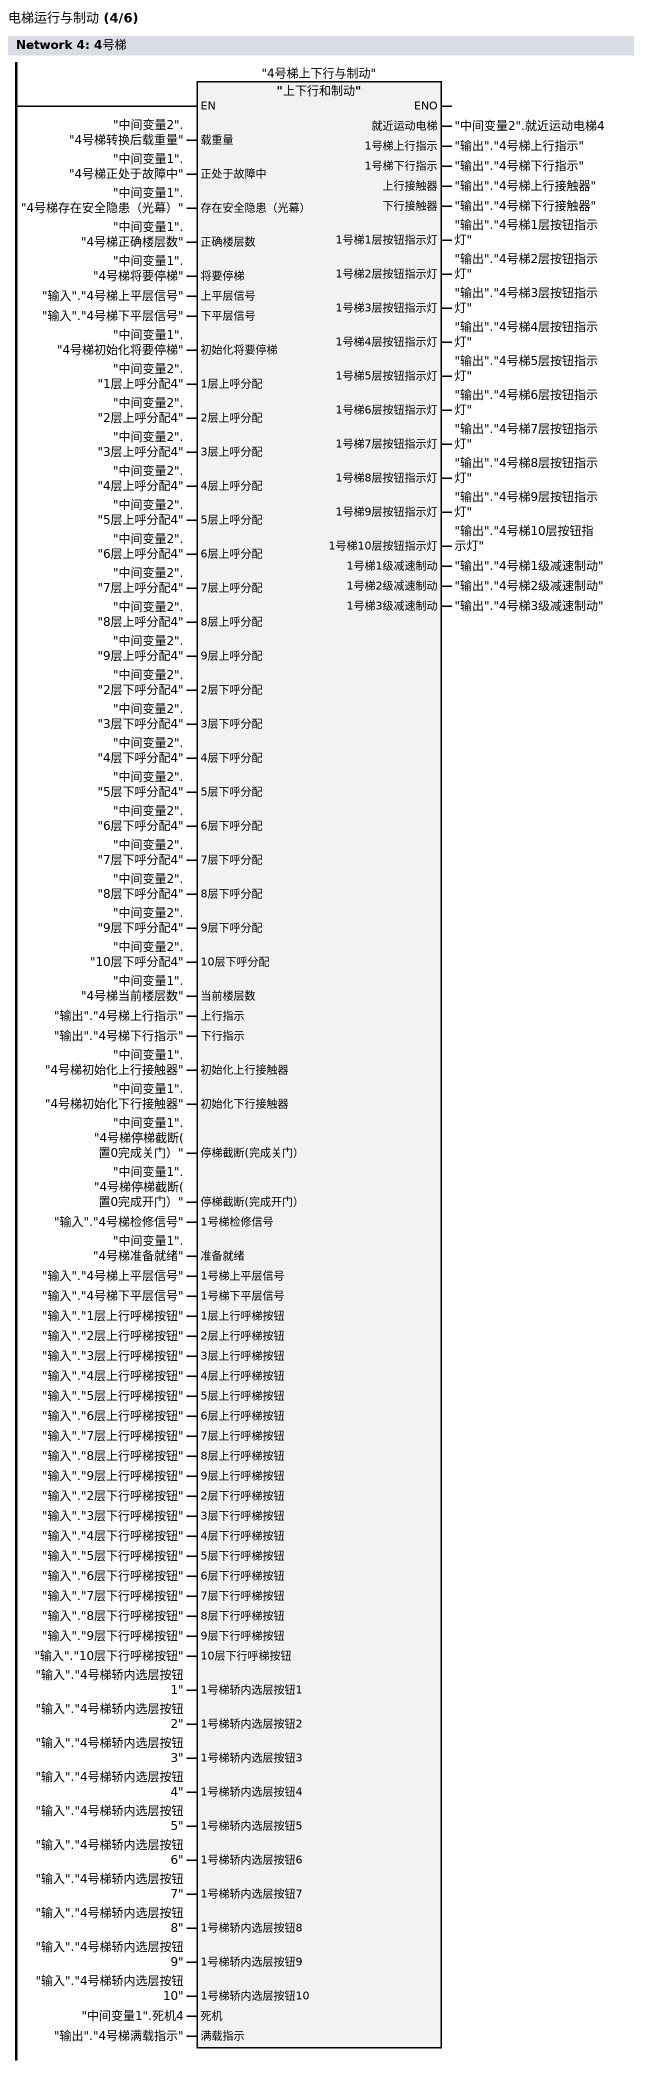
   RUNG wire#powerrail
      "4号梯上下行与制动"(载重量 := "中间变量2"."4号梯转换后载重量", 正处于故障中 := "中间变量1"."4号梯正处于故障中", "存在安全隐患（光幕）" := "中间变量1"."4号梯存在安全隐患（光幕）", 正确楼层数 := "中间变量1"."4号梯正确楼层数", 将要停梯 := "中间变量1"."4号梯将要停梯", 上平层信号 := "输入"."4号梯上平层信号", 下平层信号 := "输入"."4号梯下平层信号", 初始化将要停梯 := "中间变量1"."4号梯初始化将要停梯", "1层上呼分配" := "中间变量2"."1层上呼分配4", "2层上呼分配" := "中间变量2"."2层上呼分配4", "3层上呼分配" := "中间变量2"."3层上呼分配4", "4层上呼分配" := "中间变量2"."4层上呼分配4", "5层上呼分配" := "中间变量2"."5层上呼分配4", "6层上呼分配" := "中间变量2"."6层上呼分配4", "7层上呼分配" := "中间变量2"."7层上呼分配4", "8层上呼分配" := "中间变量2"."8层上呼分配4", "9层上呼分配" := "中间变量2"."9层上呼分配4", "2层下呼分配" := "中间变量2"."2层下呼分配4", "3层下呼分配" := "中间变量2"."3层下呼分配4", "4层下呼分配" := "中间变量2"."4层下呼分配4", "5层下呼分配" := "中间变量2"."5层下呼分配4", "6层下呼分配" := "中间变量2"."6层下呼分配4", "7层下呼分配" := "中间变量2"."7层下呼分配4", "8层下呼分配" := "中间变量2"."8层下呼分配4", "9层下呼分配" := "中间变量2"."9层下呼分配4", "10层下呼分配" := "中间变量2"."10层下呼分配4", 当前楼层数 := "中间变量1"."4号梯当前楼层数", 上行指示 := "输出"."4号梯上行指示", 下行指示 := "输出"."4号梯下行指示", 初始化上行接触器 := "中间变量1"."4号梯初始化上行接触器", 初始化下行接触器 := "中间变量1"."4号梯初始化下行接触器", "停梯截断(完成关门）" := "中间变量1"."4号梯停梯截断(置0完成关门）", "停梯截断(完成开门）" := "中间变量1"."4号梯停梯截断(置0完成开门）", "1号梯检修信号" := "输入"."4号梯检修信号", 准备就绪 := "中间变量1"."4号梯准备就绪", "1号梯上平层信号" := "输入"."4号梯上平层信号", "1号梯下平层信号" := "输入"."4号梯下平层信号", "1层上行呼梯按钮" := "输入"."1层上行呼梯按钮", "2层上行呼梯按钮" := "输入"."2层上行呼梯按钮", "3层上行呼梯按钮" := "输入"."3层上行呼梯按钮", "4层上行呼梯按钮" := "输入"."4层上行呼梯按钮", "5层上行呼梯按钮" := "输入"."5层上行呼梯按钮", "6层上行呼梯按钮" := "输入"."6层上行呼梯按钮", "7层上行呼梯按钮" := "输入"."7层上行呼梯按钮", "8层上行呼梯按钮" := "输入"."8层上行呼梯按钮", "9层上行呼梯按钮" := "输入"."9层上行呼梯按钮", "2层下行呼梯按钮" := "输入"."2层下行呼梯按钮", "3层下行呼梯按钮" := "输入"."3层下行呼梯按钮", "4层下行呼梯按钮" := "输入"."4层下行呼梯按钮", "5层下行呼梯按钮" := "输入"."5层下行呼梯按钮", "6层下行呼梯按钮" := "输入"."6层下行呼梯按钮", "7层下行呼梯按钮" := "输入"."7层下行呼梯按钮", "8层下行呼梯按钮" := "输入"."8层下行呼梯按钮", "9层下行呼梯按钮" := "输入"."9层下行呼梯按钮", "10层下行呼梯按钮" := "输入"."10层下行呼梯按钮", "1号梯轿内选层按钮1" := "输入"."4号梯轿内选层按钮1", "1号梯轿内选层按钮2" := "输入"."4号梯轿内选层按钮2", "1号梯轿内选层按钮3" := "输入"."4号梯轿内选层按钮3", "1号梯轿内选层按钮4" := "输入"."4号梯轿内选层按钮4", "1号梯轿内选层按钮5" := "输入"."4号梯轿内选层按钮5", "1号梯轿内选层按钮6" := "输入"."4号梯轿内选层按钮6", "1号梯轿内选层按钮7" := "输入"."4号梯轿内选层按钮7", "1号梯轿内选层按钮8" := "输入"."4号梯轿内选层按钮8", "1号梯轿内选层按钮9" := "输入"."4号梯轿内选层按钮9", "1号梯轿内选层按钮10" := "输入"."4号梯轿内选层按钮10", 死机 := "中间变量1".死机4, 满载指示 := "输出"."4号梯满载指示", 就近运动电梯 => "中间变量2".就近运动电梯4, "1号梯上行指示" => "输出"."4号梯上行指示", "1号梯下行指示" => "输出"."4号梯下行指示", 上行接触器 => "输出"."4号梯上行接触器", 下行接触器 => "输出"."4号梯下行接触器", "1号梯1层按钮指示灯" => "输出"."4号梯1层按钮指示灯", "1号梯2层按钮指示灯" => "输出"."4号梯2层按钮指示灯", "1号梯3层按钮指示灯" => "输出"."4号梯3层按钮指示灯", "1号梯4层按钮指示灯" => "输出"."4号梯4层按钮指示灯", "1号梯5层按钮指示灯" => "输出"."4号梯5层按钮指示灯", "1号梯6层按钮指示灯" => "输出"."4号梯6层按钮指示灯", "1号梯7层按钮指示灯" => "输出"."4号梯7层按钮指示灯", "1号梯8层按钮指示灯" => "输出"."4号梯8层按钮指示灯", "1号梯9层按钮指示灯" => "输出"."4号梯9层按钮指示灯", "1号梯10层按钮指示灯" => "输出"."4号梯10层按钮指示灯", "1号梯1级减速制动" => "输出"."4号梯1级减速制动", "1号梯2级减速制动" => "输出"."4号梯2级减速制动", "1号梯3级减速制动" => "输出"."4号梯3级减速制动")
   END_RUNG
   // the same network as SCL:
   "4号梯上下行与制动"(载重量 := "中间变量2"."4号梯转换后载重量",   // "上下行和制动"
               正处于故障中 := "中间变量1"."4号梯正处于故障中",
               "存在安全隐患（光幕）" := "中间变量1"."4号梯存在安全隐患（光幕）",
               正确楼层数 := "中间变量1"."4号梯正确楼层数",
               将要停梯 := "中间变量1"."4号梯将要停梯",
               上平层信号 := "输入"."4号梯上平层信号",
               下平层信号 := "输入"."4号梯下平层信号",
               初始化将要停梯 := "中间变量1"."4号梯初始化将要停梯",
               "1层上呼分配" := "中间变量2"."1层上呼分配4",
               "2层上呼分配" := "中间变量2"."2层上呼分配4",
               "3层上呼分配" := "中间变量2"."3层上呼分配4",
               "4层上呼分配" := "中间变量2"."4层上呼分配4",
               "5层上呼分配" := "中间变量2"."5层上呼分配4",
               "6层上呼分配" := "中间变量2"."6层上呼分配4",
               "7层上呼分配" := "中间变量2"."7层上呼分配4",
               "8层上呼分配" := "中间变量2"."8层上呼分配4",
               "9层上呼分配" := "中间变量2"."9层上呼分配4",
               "2层下呼分配" := "中间变量2"."2层下呼分配4",
               "3层下呼分配" := "中间变量2"."3层下呼分配4",
               "4层下呼分配" := "中间变量2"."4层下呼分配4",
               "5层下呼分配" := "中间变量2"."5层下呼分配4",
               "6层下呼分配" := "中间变量2"."6层下呼分配4",
               "7层下呼分配" := "中间变量2"."7层下呼分配4",
               "8层下呼分配" := "中间变量2"."8层下呼分配4",
               "9层下呼分配" := "中间变量2"."9层下呼分配4",
               "10层下呼分配" := "中间变量2"."10层下呼分配4",
               当前楼层数 := "中间变量1"."4号梯当前楼层数",
               上行指示 := "输出"."4号梯上行指示",
               下行指示 := "输出"."4号梯下行指示",
               初始化上行接触器 := "中间变量1"."4号梯初始化上行接触器",
               初始化下行接触器 := "中间变量1"."4号梯初始化下行接触器",
               "停梯截断(完成关门）" := "中间变量1"."4号梯停梯截断(置0完成关门）",
               "停梯截断(完成开门）" := "中间变量1"."4号梯停梯截断(置0完成开门）",
               "1号梯检修信号" := "输入"."4号梯检修信号",
               准备就绪 := "中间变量1"."4号梯准备就绪",
               "1号梯上平层信号" := "输入"."4号梯上平层信号",
               "1号梯下平层信号" := "输入"."4号梯下平层信号",
               "1层上行呼梯按钮" := "输入"."1层上行呼梯按钮",
               "2层上行呼梯按钮" := "输入"."2层上行呼梯按钮",
               "3层上行呼梯按钮" := "输入"."3层上行呼梯按钮",
               "4层上行呼梯按钮" := "输入"."4层上行呼梯按钮",
               "5层上行呼梯按钮" := "输入"."5层上行呼梯按钮",
               "6层上行呼梯按钮" := "输入"."6层上行呼梯按钮",
               "7层上行呼梯按钮" := "输入"."7层上行呼梯按钮",
               "8层上行呼梯按钮" := "输入"."8层上行呼梯按钮",
               "9层上行呼梯按钮" := "输入"."9层上行呼梯按钮",
               "2层下行呼梯按钮" := "输入"."2层下行呼梯按钮",
               "3层下行呼梯按钮" := "输入"."3层下行呼梯按钮",
               "4层下行呼梯按钮" := "输入"."4层下行呼梯按钮",
               "5层下行呼梯按钮" := "输入"."5层下行呼梯按钮",
               "6层下行呼梯按钮" := "输入"."6层下行呼梯按钮",
               "7层下行呼梯按钮" := "输入"."7层下行呼梯按钮",
               "8层下行呼梯按钮" := "输入"."8层下行呼梯按钮",
               "9层下行呼梯按钮" := "输入"."9层下行呼梯按钮",
               "10层下行呼梯按钮" := "输入"."10层下行呼梯按钮",
               "1号梯轿内选层按钮1" := "输入"."4号梯轿内选层按钮1",
               "1号梯轿内选层按钮2" := "输入"."4号梯轿内选层按钮2",
               "1号梯轿内选层按钮3" := "输入"."4号梯轿内选层按钮3",
               "1号梯轿内选层按钮4" := "输入"."4号梯轿内选层按钮4",
               "1号梯轿内选层按钮5" := "输入"."4号梯轿内选层按钮5",
               "1号梯轿内选层按钮6" := "输入"."4号梯轿内选层按钮6",
               "1号梯轿内选层按钮7" := "输入"."4号梯轿内选层按钮7",
               "1号梯轿内选层按钮8" := "输入"."4号梯轿内选层按钮8",
               "1号梯轿内选层按钮9" := "输入"."4号梯轿内选层按钮9",
               "1号梯轿内选层按钮10" := "输入"."4号梯轿内选层按钮10",
               死机 := "中间变量1".死机4,
               满载指示 := "输出"."4号梯满载指示",
               就近运动电梯 => "中间变量2".就近运动电梯4,
               "1号梯上行指示" => "输出"."4号梯上行指示",
               "1号梯下行指示" => "输出"."4号梯下行指示",
               上行接触器 => "输出"."4号梯上行接触器",
               下行接触器 => "输出"."4号梯下行接触器",
               "1号梯1层按钮指示灯" => "输出"."4号梯1层按钮指示灯",
               "1号梯2层按钮指示灯" => "输出"."4号梯2层按钮指示灯",
               "1号梯3层按钮指示灯" => "输出"."4号梯3层按钮指示灯",
               "1号梯4层按钮指示灯" => "输出"."4号梯4层按钮指示灯",
               "1号梯5层按钮指示灯" => "输出"."4号梯5层按钮指示灯",
               "1号梯6层按钮指示灯" => "输出"."4号梯6层按钮指示灯",
               "1号梯7层按钮指示灯" => "输出"."4号梯7层按钮指示灯",
               "1号梯8层按钮指示灯" => "输出"."4号梯8层按钮指示灯",
               "1号梯9层按钮指示灯" => "输出"."4号梯9层按钮指示灯",
               "1号梯10层按钮指示灯" => "输出"."4号梯10层按钮指示灯",
               "1号梯1级减速制动" => "输出"."4号梯1级减速制动",
               "1号梯2级减速制动" => "输出"."4号梯2级减速制动",
               "1号梯3级减速制动" => "输出"."4号梯3级减速制动");
END_REGION

REGION Network 5: 5号梯
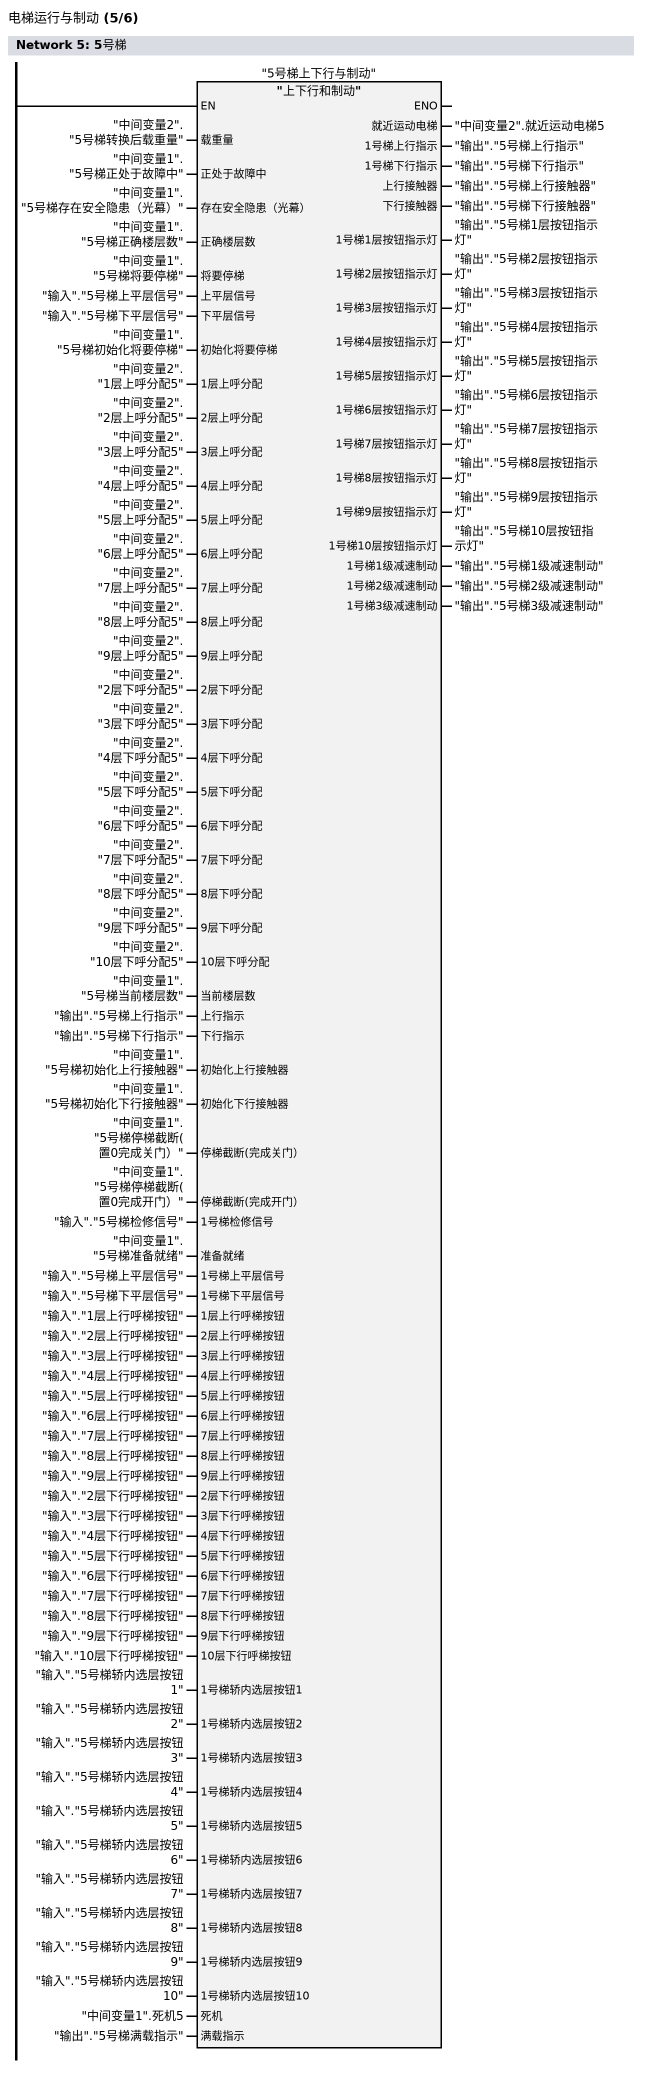
   RUNG wire#powerrail
      "5号梯上下行与制动"(载重量 := "中间变量2"."5号梯转换后载重量", 正处于故障中 := "中间变量1"."5号梯正处于故障中", "存在安全隐患（光幕）" := "中间变量1"."5号梯存在安全隐患（光幕）", 正确楼层数 := "中间变量1"."5号梯正确楼层数", 将要停梯 := "中间变量1"."5号梯将要停梯", 上平层信号 := "输入"."5号梯上平层信号", 下平层信号 := "输入"."5号梯下平层信号", 初始化将要停梯 := "中间变量1"."5号梯初始化将要停梯", "1层上呼分配" := "中间变量2"."1层上呼分配5", "2层上呼分配" := "中间变量2"."2层上呼分配5", "3层上呼分配" := "中间变量2"."3层上呼分配5", "4层上呼分配" := "中间变量2"."4层上呼分配5", "5层上呼分配" := "中间变量2"."5层上呼分配5", "6层上呼分配" := "中间变量2"."6层上呼分配5", "7层上呼分配" := "中间变量2"."7层上呼分配5", "8层上呼分配" := "中间变量2"."8层上呼分配5", "9层上呼分配" := "中间变量2"."9层上呼分配5", "2层下呼分配" := "中间变量2"."2层下呼分配5", "3层下呼分配" := "中间变量2"."3层下呼分配5", "4层下呼分配" := "中间变量2"."4层下呼分配5", "5层下呼分配" := "中间变量2"."5层下呼分配5", "6层下呼分配" := "中间变量2"."6层下呼分配5", "7层下呼分配" := "中间变量2"."7层下呼分配5", "8层下呼分配" := "中间变量2"."8层下呼分配5", "9层下呼分配" := "中间变量2"."9层下呼分配5", "10层下呼分配" := "中间变量2"."10层下呼分配5", 当前楼层数 := "中间变量1"."5号梯当前楼层数", 上行指示 := "输出"."5号梯上行指示", 下行指示 := "输出"."5号梯下行指示", 初始化上行接触器 := "中间变量1"."5号梯初始化上行接触器", 初始化下行接触器 := "中间变量1"."5号梯初始化下行接触器", "停梯截断(完成关门）" := "中间变量1"."5号梯停梯截断(置0完成关门）", "停梯截断(完成开门）" := "中间变量1"."5号梯停梯截断(置0完成开门）", "1号梯检修信号" := "输入"."5号梯检修信号", 准备就绪 := "中间变量1"."5号梯准备就绪", "1号梯上平层信号" := "输入"."5号梯上平层信号", "1号梯下平层信号" := "输入"."5号梯下平层信号", "1层上行呼梯按钮" := "输入"."1层上行呼梯按钮", "2层上行呼梯按钮" := "输入"."2层上行呼梯按钮", "3层上行呼梯按钮" := "输入"."3层上行呼梯按钮", "4层上行呼梯按钮" := "输入"."4层上行呼梯按钮", "5层上行呼梯按钮" := "输入"."5层上行呼梯按钮", "6层上行呼梯按钮" := "输入"."6层上行呼梯按钮", "7层上行呼梯按钮" := "输入"."7层上行呼梯按钮", "8层上行呼梯按钮" := "输入"."8层上行呼梯按钮", "9层上行呼梯按钮" := "输入"."9层上行呼梯按钮", "2层下行呼梯按钮" := "输入"."2层下行呼梯按钮", "3层下行呼梯按钮" := "输入"."3层下行呼梯按钮", "4层下行呼梯按钮" := "输入"."4层下行呼梯按钮", "5层下行呼梯按钮" := "输入"."5层下行呼梯按钮", "6层下行呼梯按钮" := "输入"."6层下行呼梯按钮", "7层下行呼梯按钮" := "输入"."7层下行呼梯按钮", "8层下行呼梯按钮" := "输入"."8层下行呼梯按钮", "9层下行呼梯按钮" := "输入"."9层下行呼梯按钮", "10层下行呼梯按钮" := "输入"."10层下行呼梯按钮", "1号梯轿内选层按钮1" := "输入"."5号梯轿内选层按钮1", "1号梯轿内选层按钮2" := "输入"."5号梯轿内选层按钮2", "1号梯轿内选层按钮3" := "输入"."5号梯轿内选层按钮3", "1号梯轿内选层按钮4" := "输入"."5号梯轿内选层按钮4", "1号梯轿内选层按钮5" := "输入"."5号梯轿内选层按钮5", "1号梯轿内选层按钮6" := "输入"."5号梯轿内选层按钮6", "1号梯轿内选层按钮7" := "输入"."5号梯轿内选层按钮7", "1号梯轿内选层按钮8" := "输入"."5号梯轿内选层按钮8", "1号梯轿内选层按钮9" := "输入"."5号梯轿内选层按钮9", "1号梯轿内选层按钮10" := "输入"."5号梯轿内选层按钮10", 死机 := "中间变量1".死机5, 满载指示 := "输出"."5号梯满载指示", 就近运动电梯 => "中间变量2".就近运动电梯5, "1号梯上行指示" => "输出"."5号梯上行指示", "1号梯下行指示" => "输出"."5号梯下行指示", 上行接触器 => "输出"."5号梯上行接触器", 下行接触器 => "输出"."5号梯下行接触器", "1号梯1层按钮指示灯" => "输出"."5号梯1层按钮指示灯", "1号梯2层按钮指示灯" => "输出"."5号梯2层按钮指示灯", "1号梯3层按钮指示灯" => "输出"."5号梯3层按钮指示灯", "1号梯4层按钮指示灯" => "输出"."5号梯4层按钮指示灯", "1号梯5层按钮指示灯" => "输出"."5号梯5层按钮指示灯", "1号梯6层按钮指示灯" => "输出"."5号梯6层按钮指示灯", "1号梯7层按钮指示灯" => "输出"."5号梯7层按钮指示灯", "1号梯8层按钮指示灯" => "输出"."5号梯8层按钮指示灯", "1号梯9层按钮指示灯" => "输出"."5号梯9层按钮指示灯", "1号梯10层按钮指示灯" => "输出"."5号梯10层按钮指示灯", "1号梯1级减速制动" => "输出"."5号梯1级减速制动", "1号梯2级减速制动" => "输出"."5号梯2级减速制动", "1号梯3级减速制动" => "输出"."5号梯3级减速制动")
   END_RUNG
   // the same network as SCL:
   "5号梯上下行与制动"(载重量 := "中间变量2"."5号梯转换后载重量",   // "上下行和制动"
               正处于故障中 := "中间变量1"."5号梯正处于故障中",
               "存在安全隐患（光幕）" := "中间变量1"."5号梯存在安全隐患（光幕）",
               正确楼层数 := "中间变量1"."5号梯正确楼层数",
               将要停梯 := "中间变量1"."5号梯将要停梯",
               上平层信号 := "输入"."5号梯上平层信号",
               下平层信号 := "输入"."5号梯下平层信号",
               初始化将要停梯 := "中间变量1"."5号梯初始化将要停梯",
               "1层上呼分配" := "中间变量2"."1层上呼分配5",
               "2层上呼分配" := "中间变量2"."2层上呼分配5",
               "3层上呼分配" := "中间变量2"."3层上呼分配5",
               "4层上呼分配" := "中间变量2"."4层上呼分配5",
               "5层上呼分配" := "中间变量2"."5层上呼分配5",
               "6层上呼分配" := "中间变量2"."6层上呼分配5",
               "7层上呼分配" := "中间变量2"."7层上呼分配5",
               "8层上呼分配" := "中间变量2"."8层上呼分配5",
               "9层上呼分配" := "中间变量2"."9层上呼分配5",
               "2层下呼分配" := "中间变量2"."2层下呼分配5",
               "3层下呼分配" := "中间变量2"."3层下呼分配5",
               "4层下呼分配" := "中间变量2"."4层下呼分配5",
               "5层下呼分配" := "中间变量2"."5层下呼分配5",
               "6层下呼分配" := "中间变量2"."6层下呼分配5",
               "7层下呼分配" := "中间变量2"."7层下呼分配5",
               "8层下呼分配" := "中间变量2"."8层下呼分配5",
               "9层下呼分配" := "中间变量2"."9层下呼分配5",
               "10层下呼分配" := "中间变量2"."10层下呼分配5",
               当前楼层数 := "中间变量1"."5号梯当前楼层数",
               上行指示 := "输出"."5号梯上行指示",
               下行指示 := "输出"."5号梯下行指示",
               初始化上行接触器 := "中间变量1"."5号梯初始化上行接触器",
               初始化下行接触器 := "中间变量1"."5号梯初始化下行接触器",
               "停梯截断(完成关门）" := "中间变量1"."5号梯停梯截断(置0完成关门）",
               "停梯截断(完成开门）" := "中间变量1"."5号梯停梯截断(置0完成开门）",
               "1号梯检修信号" := "输入"."5号梯检修信号",
               准备就绪 := "中间变量1"."5号梯准备就绪",
               "1号梯上平层信号" := "输入"."5号梯上平层信号",
               "1号梯下平层信号" := "输入"."5号梯下平层信号",
               "1层上行呼梯按钮" := "输入"."1层上行呼梯按钮",
               "2层上行呼梯按钮" := "输入"."2层上行呼梯按钮",
               "3层上行呼梯按钮" := "输入"."3层上行呼梯按钮",
               "4层上行呼梯按钮" := "输入"."4层上行呼梯按钮",
               "5层上行呼梯按钮" := "输入"."5层上行呼梯按钮",
               "6层上行呼梯按钮" := "输入"."6层上行呼梯按钮",
               "7层上行呼梯按钮" := "输入"."7层上行呼梯按钮",
               "8层上行呼梯按钮" := "输入"."8层上行呼梯按钮",
               "9层上行呼梯按钮" := "输入"."9层上行呼梯按钮",
               "2层下行呼梯按钮" := "输入"."2层下行呼梯按钮",
               "3层下行呼梯按钮" := "输入"."3层下行呼梯按钮",
               "4层下行呼梯按钮" := "输入"."4层下行呼梯按钮",
               "5层下行呼梯按钮" := "输入"."5层下行呼梯按钮",
               "6层下行呼梯按钮" := "输入"."6层下行呼梯按钮",
               "7层下行呼梯按钮" := "输入"."7层下行呼梯按钮",
               "8层下行呼梯按钮" := "输入"."8层下行呼梯按钮",
               "9层下行呼梯按钮" := "输入"."9层下行呼梯按钮",
               "10层下行呼梯按钮" := "输入"."10层下行呼梯按钮",
               "1号梯轿内选层按钮1" := "输入"."5号梯轿内选层按钮1",
               "1号梯轿内选层按钮2" := "输入"."5号梯轿内选层按钮2",
               "1号梯轿内选层按钮3" := "输入"."5号梯轿内选层按钮3",
               "1号梯轿内选层按钮4" := "输入"."5号梯轿内选层按钮4",
               "1号梯轿内选层按钮5" := "输入"."5号梯轿内选层按钮5",
               "1号梯轿内选层按钮6" := "输入"."5号梯轿内选层按钮6",
               "1号梯轿内选层按钮7" := "输入"."5号梯轿内选层按钮7",
               "1号梯轿内选层按钮8" := "输入"."5号梯轿内选层按钮8",
               "1号梯轿内选层按钮9" := "输入"."5号梯轿内选层按钮9",
               "1号梯轿内选层按钮10" := "输入"."5号梯轿内选层按钮10",
               死机 := "中间变量1".死机5,
               满载指示 := "输出"."5号梯满载指示",
               就近运动电梯 => "中间变量2".就近运动电梯5,
               "1号梯上行指示" => "输出"."5号梯上行指示",
               "1号梯下行指示" => "输出"."5号梯下行指示",
               上行接触器 => "输出"."5号梯上行接触器",
               下行接触器 => "输出"."5号梯下行接触器",
               "1号梯1层按钮指示灯" => "输出"."5号梯1层按钮指示灯",
               "1号梯2层按钮指示灯" => "输出"."5号梯2层按钮指示灯",
               "1号梯3层按钮指示灯" => "输出"."5号梯3层按钮指示灯",
               "1号梯4层按钮指示灯" => "输出"."5号梯4层按钮指示灯",
               "1号梯5层按钮指示灯" => "输出"."5号梯5层按钮指示灯",
               "1号梯6层按钮指示灯" => "输出"."5号梯6层按钮指示灯",
               "1号梯7层按钮指示灯" => "输出"."5号梯7层按钮指示灯",
               "1号梯8层按钮指示灯" => "输出"."5号梯8层按钮指示灯",
               "1号梯9层按钮指示灯" => "输出"."5号梯9层按钮指示灯",
               "1号梯10层按钮指示灯" => "输出"."5号梯10层按钮指示灯",
               "1号梯1级减速制动" => "输出"."5号梯1级减速制动",
               "1号梯2级减速制动" => "输出"."5号梯2级减速制动",
               "1号梯3级减速制动" => "输出"."5号梯3级减速制动");
END_REGION

REGION Network 6: 6号梯
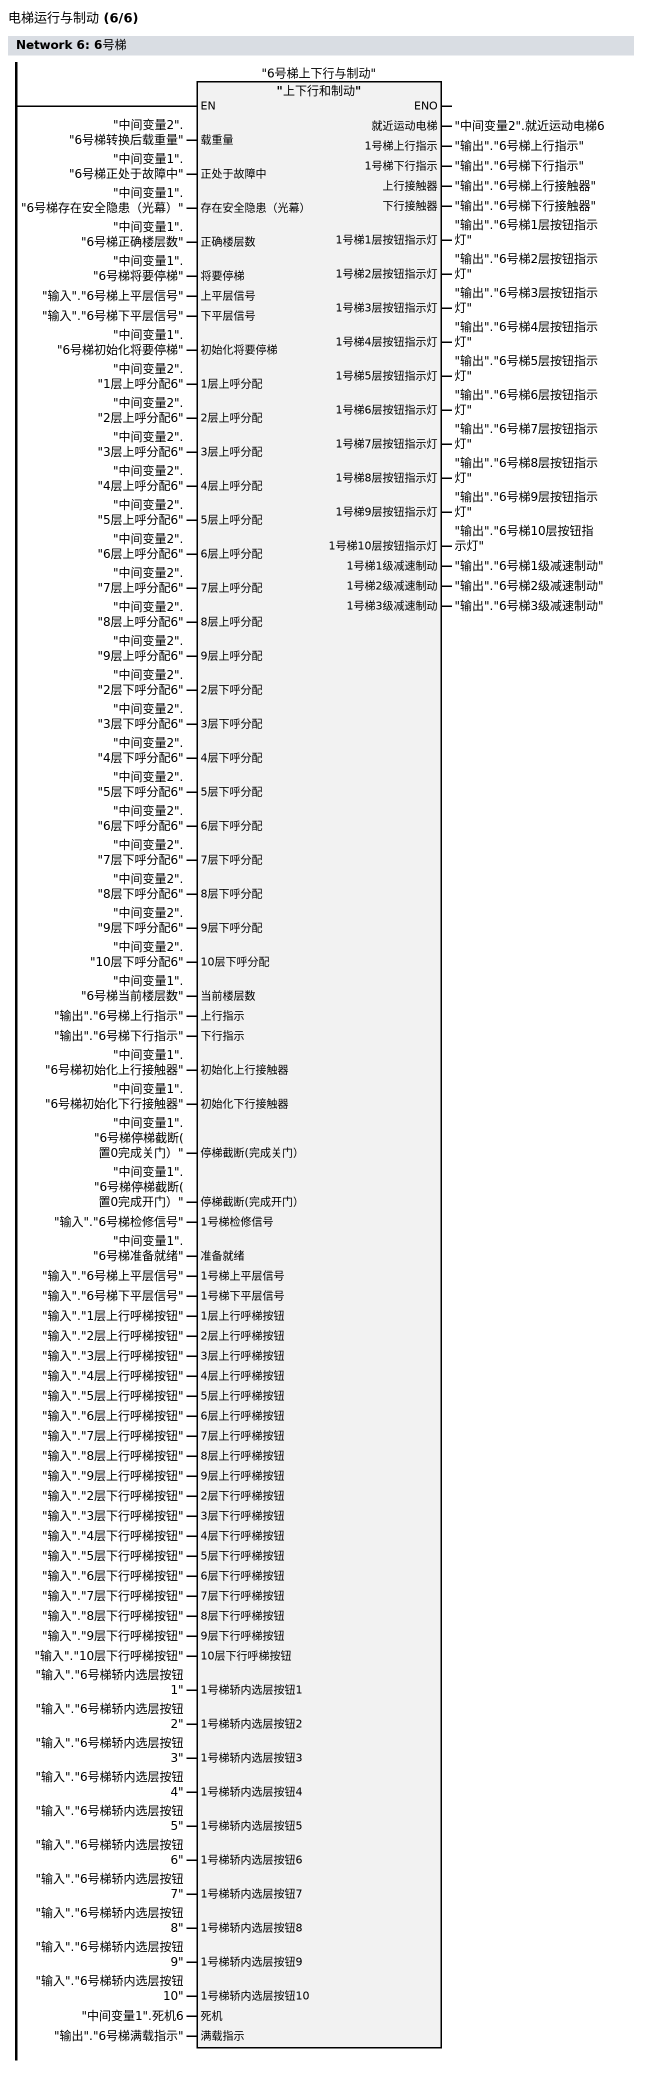
   RUNG wire#powerrail
      "6号梯上下行与制动"(载重量 := "中间变量2"."6号梯转换后载重量", 正处于故障中 := "中间变量1"."6号梯正处于故障中", "存在安全隐患（光幕）" := "中间变量1"."6号梯存在安全隐患（光幕）", 正确楼层数 := "中间变量1"."6号梯正确楼层数", 将要停梯 := "中间变量1"."6号梯将要停梯", 上平层信号 := "输入"."6号梯上平层信号", 下平层信号 := "输入"."6号梯下平层信号", 初始化将要停梯 := "中间变量1"."6号梯初始化将要停梯", "1层上呼分配" := "中间变量2"."1层上呼分配6", "2层上呼分配" := "中间变量2"."2层上呼分配6", "3层上呼分配" := "中间变量2"."3层上呼分配6", "4层上呼分配" := "中间变量2"."4层上呼分配6", "5层上呼分配" := "中间变量2"."5层上呼分配6", "6层上呼分配" := "中间变量2"."6层上呼分配6", "7层上呼分配" := "中间变量2"."7层上呼分配6", "8层上呼分配" := "中间变量2"."8层上呼分配6", "9层上呼分配" := "中间变量2"."9层上呼分配6", "2层下呼分配" := "中间变量2"."2层下呼分配6", "3层下呼分配" := "中间变量2"."3层下呼分配6", "4层下呼分配" := "中间变量2"."4层下呼分配6", "5层下呼分配" := "中间变量2"."5层下呼分配6", "6层下呼分配" := "中间变量2"."6层下呼分配6", "7层下呼分配" := "中间变量2"."7层下呼分配6", "8层下呼分配" := "中间变量2"."8层下呼分配6", "9层下呼分配" := "中间变量2"."9层下呼分配6", "10层下呼分配" := "中间变量2"."10层下呼分配6", 当前楼层数 := "中间变量1"."6号梯当前楼层数", 上行指示 := "输出"."6号梯上行指示", 下行指示 := "输出"."6号梯下行指示", 初始化上行接触器 := "中间变量1"."6号梯初始化上行接触器", 初始化下行接触器 := "中间变量1"."6号梯初始化下行接触器", "停梯截断(完成关门）" := "中间变量1"."6号梯停梯截断(置0完成关门）", "停梯截断(完成开门）" := "中间变量1"."6号梯停梯截断(置0完成开门）", "1号梯检修信号" := "输入"."6号梯检修信号", 准备就绪 := "中间变量1"."6号梯准备就绪", "1号梯上平层信号" := "输入"."6号梯上平层信号", "1号梯下平层信号" := "输入"."6号梯下平层信号", "1层上行呼梯按钮" := "输入"."1层上行呼梯按钮", "2层上行呼梯按钮" := "输入"."2层上行呼梯按钮", "3层上行呼梯按钮" := "输入"."3层上行呼梯按钮", "4层上行呼梯按钮" := "输入"."4层上行呼梯按钮", "5层上行呼梯按钮" := "输入"."5层上行呼梯按钮", "6层上行呼梯按钮" := "输入"."6层上行呼梯按钮", "7层上行呼梯按钮" := "输入"."7层上行呼梯按钮", "8层上行呼梯按钮" := "输入"."8层上行呼梯按钮", "9层上行呼梯按钮" := "输入"."9层上行呼梯按钮", "2层下行呼梯按钮" := "输入"."2层下行呼梯按钮", "3层下行呼梯按钮" := "输入"."3层下行呼梯按钮", "4层下行呼梯按钮" := "输入"."4层下行呼梯按钮", "5层下行呼梯按钮" := "输入"."5层下行呼梯按钮", "6层下行呼梯按钮" := "输入"."6层下行呼梯按钮", "7层下行呼梯按钮" := "输入"."7层下行呼梯按钮", "8层下行呼梯按钮" := "输入"."8层下行呼梯按钮", "9层下行呼梯按钮" := "输入"."9层下行呼梯按钮", "10层下行呼梯按钮" := "输入"."10层下行呼梯按钮", "1号梯轿内选层按钮1" := "输入"."6号梯轿内选层按钮1", "1号梯轿内选层按钮2" := "输入"."6号梯轿内选层按钮2", "1号梯轿内选层按钮3" := "输入"."6号梯轿内选层按钮3", "1号梯轿内选层按钮4" := "输入"."6号梯轿内选层按钮4", "1号梯轿内选层按钮5" := "输入"."6号梯轿内选层按钮5", "1号梯轿内选层按钮6" := "输入"."6号梯轿内选层按钮6", "1号梯轿内选层按钮7" := "输入"."6号梯轿内选层按钮7", "1号梯轿内选层按钮8" := "输入"."6号梯轿内选层按钮8", "1号梯轿内选层按钮9" := "输入"."6号梯轿内选层按钮9", "1号梯轿内选层按钮10" := "输入"."6号梯轿内选层按钮10", 死机 := "中间变量1".死机6, 满载指示 := "输出"."6号梯满载指示", 就近运动电梯 => "中间变量2".就近运动电梯6, "1号梯上行指示" => "输出"."6号梯上行指示", "1号梯下行指示" => "输出"."6号梯下行指示", 上行接触器 => "输出"."6号梯上行接触器", 下行接触器 => "输出"."6号梯下行接触器", "1号梯1层按钮指示灯" => "输出"."6号梯1层按钮指示灯", "1号梯2层按钮指示灯" => "输出"."6号梯2层按钮指示灯", "1号梯3层按钮指示灯" => "输出"."6号梯3层按钮指示灯", "1号梯4层按钮指示灯" => "输出"."6号梯4层按钮指示灯", "1号梯5层按钮指示灯" => "输出"."6号梯5层按钮指示灯", "1号梯6层按钮指示灯" => "输出"."6号梯6层按钮指示灯", "1号梯7层按钮指示灯" => "输出"."6号梯7层按钮指示灯", "1号梯8层按钮指示灯" => "输出"."6号梯8层按钮指示灯", "1号梯9层按钮指示灯" => "输出"."6号梯9层按钮指示灯", "1号梯10层按钮指示灯" => "输出"."6号梯10层按钮指示灯", "1号梯1级减速制动" => "输出"."6号梯1级减速制动", "1号梯2级减速制动" => "输出"."6号梯2级减速制动", "1号梯3级减速制动" => "输出"."6号梯3级减速制动")
   END_RUNG
   // the same network as SCL:
   "6号梯上下行与制动"(载重量 := "中间变量2"."6号梯转换后载重量",   // "上下行和制动"
               正处于故障中 := "中间变量1"."6号梯正处于故障中",
               "存在安全隐患（光幕）" := "中间变量1"."6号梯存在安全隐患（光幕）",
               正确楼层数 := "中间变量1"."6号梯正确楼层数",
               将要停梯 := "中间变量1"."6号梯将要停梯",
               上平层信号 := "输入"."6号梯上平层信号",
               下平层信号 := "输入"."6号梯下平层信号",
               初始化将要停梯 := "中间变量1"."6号梯初始化将要停梯",
               "1层上呼分配" := "中间变量2"."1层上呼分配6",
               "2层上呼分配" := "中间变量2"."2层上呼分配6",
               "3层上呼分配" := "中间变量2"."3层上呼分配6",
               "4层上呼分配" := "中间变量2"."4层上呼分配6",
               "5层上呼分配" := "中间变量2"."5层上呼分配6",
               "6层上呼分配" := "中间变量2"."6层上呼分配6",
               "7层上呼分配" := "中间变量2"."7层上呼分配6",
               "8层上呼分配" := "中间变量2"."8层上呼分配6",
               "9层上呼分配" := "中间变量2"."9层上呼分配6",
               "2层下呼分配" := "中间变量2"."2层下呼分配6",
               "3层下呼分配" := "中间变量2"."3层下呼分配6",
               "4层下呼分配" := "中间变量2"."4层下呼分配6",
               "5层下呼分配" := "中间变量2"."5层下呼分配6",
               "6层下呼分配" := "中间变量2"."6层下呼分配6",
               "7层下呼分配" := "中间变量2"."7层下呼分配6",
               "8层下呼分配" := "中间变量2"."8层下呼分配6",
               "9层下呼分配" := "中间变量2"."9层下呼分配6",
               "10层下呼分配" := "中间变量2"."10层下呼分配6",
               当前楼层数 := "中间变量1"."6号梯当前楼层数",
               上行指示 := "输出"."6号梯上行指示",
               下行指示 := "输出"."6号梯下行指示",
               初始化上行接触器 := "中间变量1"."6号梯初始化上行接触器",
               初始化下行接触器 := "中间变量1"."6号梯初始化下行接触器",
               "停梯截断(完成关门）" := "中间变量1"."6号梯停梯截断(置0完成关门）",
               "停梯截断(完成开门）" := "中间变量1"."6号梯停梯截断(置0完成开门）",
               "1号梯检修信号" := "输入"."6号梯检修信号",
               准备就绪 := "中间变量1"."6号梯准备就绪",
               "1号梯上平层信号" := "输入"."6号梯上平层信号",
               "1号梯下平层信号" := "输入"."6号梯下平层信号",
               "1层上行呼梯按钮" := "输入"."1层上行呼梯按钮",
               "2层上行呼梯按钮" := "输入"."2层上行呼梯按钮",
               "3层上行呼梯按钮" := "输入"."3层上行呼梯按钮",
               "4层上行呼梯按钮" := "输入"."4层上行呼梯按钮",
               "5层上行呼梯按钮" := "输入"."5层上行呼梯按钮",
               "6层上行呼梯按钮" := "输入"."6层上行呼梯按钮",
               "7层上行呼梯按钮" := "输入"."7层上行呼梯按钮",
               "8层上行呼梯按钮" := "输入"."8层上行呼梯按钮",
               "9层上行呼梯按钮" := "输入"."9层上行呼梯按钮",
               "2层下行呼梯按钮" := "输入"."2层下行呼梯按钮",
               "3层下行呼梯按钮" := "输入"."3层下行呼梯按钮",
               "4层下行呼梯按钮" := "输入"."4层下行呼梯按钮",
               "5层下行呼梯按钮" := "输入"."5层下行呼梯按钮",
               "6层下行呼梯按钮" := "输入"."6层下行呼梯按钮",
               "7层下行呼梯按钮" := "输入"."7层下行呼梯按钮",
               "8层下行呼梯按钮" := "输入"."8层下行呼梯按钮",
               "9层下行呼梯按钮" := "输入"."9层下行呼梯按钮",
               "10层下行呼梯按钮" := "输入"."10层下行呼梯按钮",
               "1号梯轿内选层按钮1" := "输入"."6号梯轿内选层按钮1",
               "1号梯轿内选层按钮2" := "输入"."6号梯轿内选层按钮2",
               "1号梯轿内选层按钮3" := "输入"."6号梯轿内选层按钮3",
               "1号梯轿内选层按钮4" := "输入"."6号梯轿内选层按钮4",
               "1号梯轿内选层按钮5" := "输入"."6号梯轿内选层按钮5",
               "1号梯轿内选层按钮6" := "输入"."6号梯轿内选层按钮6",
               "1号梯轿内选层按钮7" := "输入"."6号梯轿内选层按钮7",
               "1号梯轿内选层按钮8" := "输入"."6号梯轿内选层按钮8",
               "1号梯轿内选层按钮9" := "输入"."6号梯轿内选层按钮9",
               "1号梯轿内选层按钮10" := "输入"."6号梯轿内选层按钮10",
               死机 := "中间变量1".死机6,
               满载指示 := "输出"."6号梯满载指示",
               就近运动电梯 => "中间变量2".就近运动电梯6,
               "1号梯上行指示" => "输出"."6号梯上行指示",
               "1号梯下行指示" => "输出"."6号梯下行指示",
               上行接触器 => "输出"."6号梯上行接触器",
               下行接触器 => "输出"."6号梯下行接触器",
               "1号梯1层按钮指示灯" => "输出"."6号梯1层按钮指示灯",
               "1号梯2层按钮指示灯" => "输出"."6号梯2层按钮指示灯",
               "1号梯3层按钮指示灯" => "输出"."6号梯3层按钮指示灯",
               "1号梯4层按钮指示灯" => "输出"."6号梯4层按钮指示灯",
               "1号梯5层按钮指示灯" => "输出"."6号梯5层按钮指示灯",
               "1号梯6层按钮指示灯" => "输出"."6号梯6层按钮指示灯",
               "1号梯7层按钮指示灯" => "输出"."6号梯7层按钮指示灯",
               "1号梯8层按钮指示灯" => "输出"."6号梯8层按钮指示灯",
               "1号梯9层按钮指示灯" => "输出"."6号梯9层按钮指示灯",
               "1号梯10层按钮指示灯" => "输出"."6号梯10层按钮指示灯",
               "1号梯1级减速制动" => "输出"."6号梯1级减速制动",
               "1号梯2级减速制动" => "输出"."6号梯2级减速制动",
               "1号梯3级减速制动" => "输出"."6号梯3级减速制动");
END_REGION
END_FUNCTION

FUNCTION "距离调度算法" : Void   // FC5, LAD
{ S7_Optimized_Access := 'TRUE' }
VERSION : 0.1
BEGIN

REGION Network 2: 1号梯调度距离
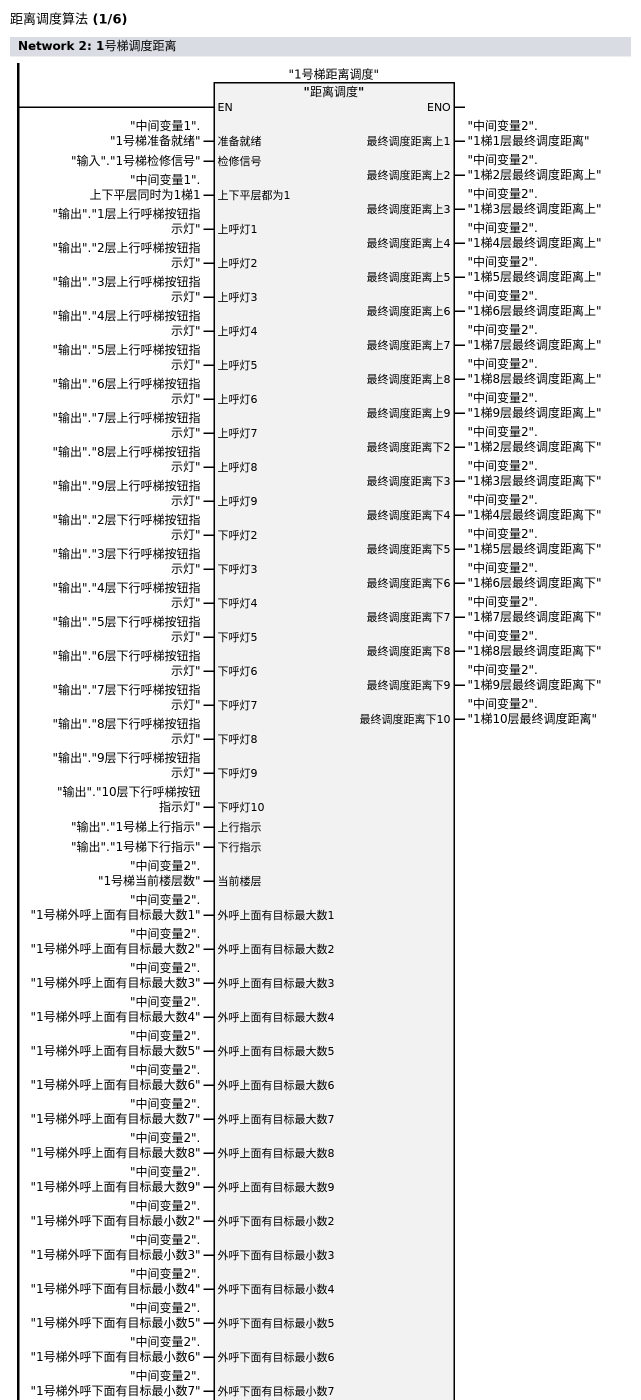
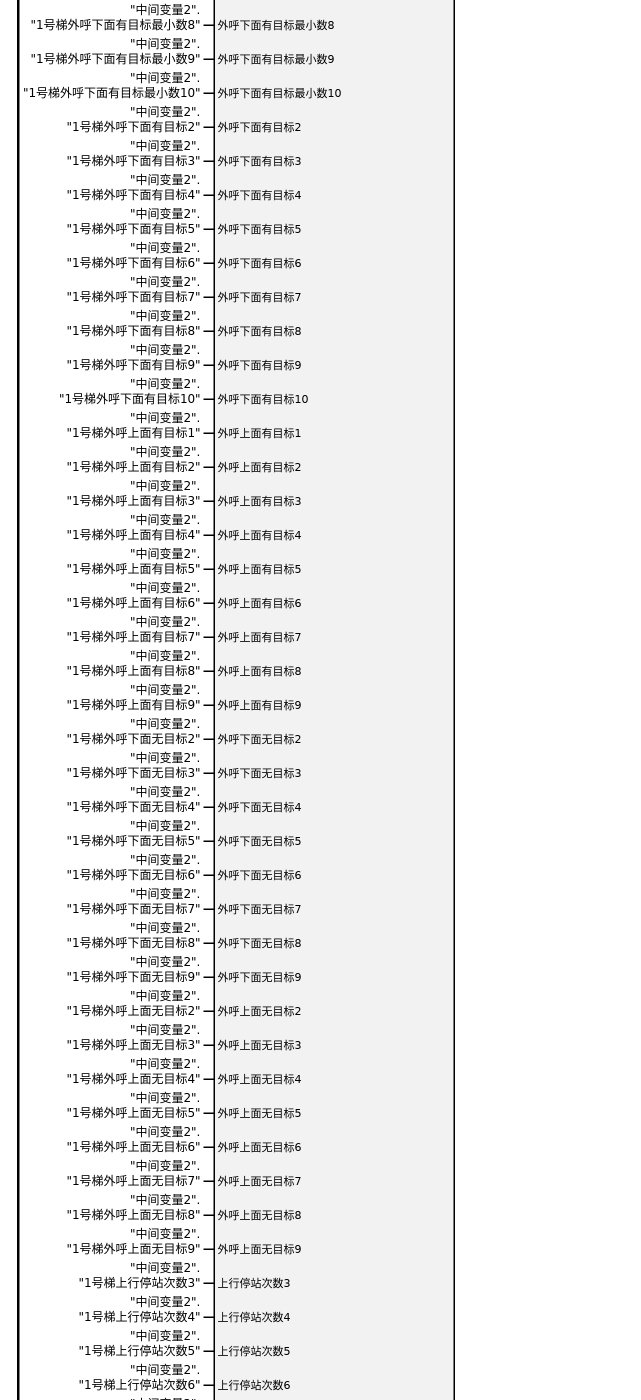
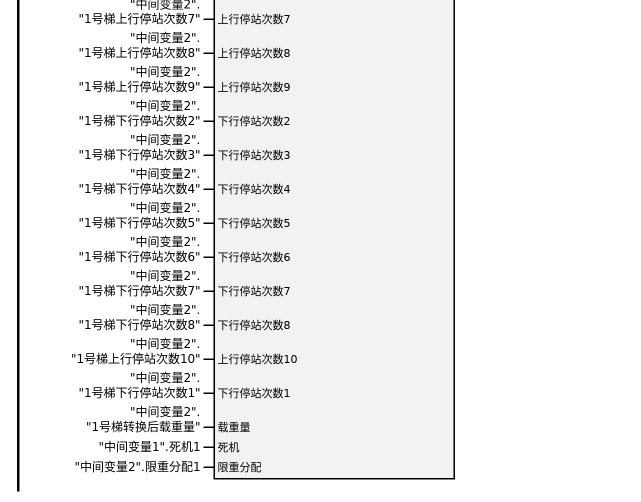
   RUNG wire#powerrail
      "1号梯距离调度"(准备就绪 := "中间变量1"."1号梯准备就绪", 检修信号 := "输入"."1号梯检修信号", 上下平层都为1 := "中间变量1".上下平层同时为1梯1, 上呼灯1 := "输出"."1层上行呼梯按钮指示灯", 上呼灯2 := "输出"."2层上行呼梯按钮指示灯", 上呼灯3 := "输出"."3层上行呼梯按钮指示灯", 上呼灯4 := "输出"."4层上行呼梯按钮指示灯", 上呼灯5 := "输出"."5层上行呼梯按钮指示灯", 上呼灯6 := "输出"."6层上行呼梯按钮指示灯", 上呼灯7 := "输出"."7层上行呼梯按钮指示灯", 上呼灯8 := "输出"."8层上行呼梯按钮指示灯", 上呼灯9 := "输出"."9层上行呼梯按钮指示灯", 下呼灯2 := "输出"."2层下行呼梯按钮指示灯", 下呼灯3 := "输出"."3层下行呼梯按钮指示灯", 下呼灯4 := "输出"."4层下行呼梯按钮指示灯", 下呼灯5 := "输出"."5层下行呼梯按钮指示灯", 下呼灯6 := "输出"."6层下行呼梯按钮指示灯", 下呼灯7 := "输出"."7层下行呼梯按钮指示灯", 下呼灯8 := "输出"."8层下行呼梯按钮指示灯", 下呼灯9 := "输出"."9层下行呼梯按钮指示灯", 下呼灯10 := "输出"."10层下行呼梯按钮指示灯", 上行指示 := "输出"."1号梯上行指示", 下行指示 := "输出"."1号梯下行指示", 当前楼层 := "中间变量2"."1号梯当前楼层数", 外呼上面有目标最大数1 := "中间变量2"."1号梯外呼上面有目标最大数1", 外呼上面有目标最大数2 := "中间变量2"."1号梯外呼上面有目标最大数2", 外呼上面有目标最大数3 := "中间变量2"."1号梯外呼上面有目标最大数3", 外呼上面有目标最大数4 := "中间变量2"."1号梯外呼上面有目标最大数4", 外呼上面有目标最大数5 := "中间变量2"."1号梯外呼上面有目标最大数5", 外呼上面有目标最大数6 := "中间变量2"."1号梯外呼上面有目标最大数6", 外呼上面有目标最大数7 := "中间变量2"."1号梯外呼上面有目标最大数7", 外呼上面有目标最大数8 := "中间变量2"."1号梯外呼上面有目标最大数8", 外呼上面有目标最大数9 := "中间变量2"."1号梯外呼上面有目标最大数9", 外呼下面有目标最小数2 := "中间变量2"."1号梯外呼下面有目标最小数2", 外呼下面有目标最小数3 := "中间变量2"."1号梯外呼下面有目标最小数3", 外呼下面有目标最小数4 := "中间变量2"."1号梯外呼下面有目标最小数4", 外呼下面有目标最小数5 := "中间变量2"."1号梯外呼下面有目标最小数5", 外呼下面有目标最小数6 := "中间变量2"."1号梯外呼下面有目标最小数6", 外呼下面有目标最小数7 := "中间变量2"."1号梯外呼下面有目标最小数7", 外呼下面有目标最小数8 := "中间变量2"."1号梯外呼下面有目标最小数8", 外呼下面有目标最小数9 := "中间变量2"."1号梯外呼下面有目标最小数9", 外呼下面有目标最小数10 := "中间变量2"."1号梯外呼下面有目标最小数10", 外呼下面有目标2 := "中间变量2"."1号梯外呼下面有目标2", 外呼下面有目标3 := "中间变量2"."1号梯外呼下面有目标3", 外呼下面有目标4 := "中间变量2"."1号梯外呼下面有目标4", 外呼下面有目标5 := "中间变量2"."1号梯外呼下面有目标5", 外呼下面有目标6 := "中间变量2"."1号梯外呼下面有目标6", 外呼下面有目标7 := "中间变量2"."1号梯外呼下面有目标7", 外呼下面有目标8 := "中间变量2"."1号梯外呼下面有目标8", 外呼下面有目标9 := "中间变量2"."1号梯外呼下面有目标9", 外呼下面有目标10 := "中间变量2"."1号梯外呼下面有目标10", 外呼上面有目标1 := "中间变量2"."1号梯外呼上面有目标1", 外呼上面有目标2 := "中间变量2"."1号梯外呼上面有目标2", 外呼上面有目标3 := "中间变量2"."1号梯外呼上面有目标3", 外呼上面有目标4 := "中间变量2"."1号梯外呼上面有目标4", 外呼上面有目标5 := "中间变量2"."1号梯外呼上面有目标5", 外呼上面有目标6 := "中间变量2"."1号梯外呼上面有目标6", 外呼上面有目标7 := "中间变量2"."1号梯外呼上面有目标7", 外呼上面有目标8 := "中间变量2"."1号梯外呼上面有目标8", 外呼上面有目标9 := "中间变量2"."1号梯外呼上面有目标9", 外呼下面无目标2 := "中间变量2"."1号梯外呼下面无目标2", 外呼下面无目标3 := "中间变量2"."1号梯外呼下面无目标3", 外呼下面无目标4 := "中间变量2"."1号梯外呼下面无目标4", 外呼下面无目标5 := "中间变量2"."1号梯外呼下面无目标5", 外呼下面无目标6 := "中间变量2"."1号梯外呼下面无目标6", 外呼下面无目标7 := "中间变量2"."1号梯外呼下面无目标7", 外呼下面无目标8 := "中间变量2"."1号梯外呼下面无目标8", 外呼下面无目标9 := "中间变量2"."1号梯外呼下面无目标9", 外呼上面无目标2 := "中间变量2"."1号梯外呼上面无目标2", 外呼上面无目标3 := "中间变量2"."1号梯外呼上面无目标3", 外呼上面无目标4 := "中间变量2"."1号梯外呼上面无目标4", 外呼上面无目标5 := "中间变量2"."1号梯外呼上面无目标5", 外呼上面无目标6 := "中间变量2"."1号梯外呼上面无目标6", 外呼上面无目标7 := "中间变量2"."1号梯外呼上面无目标7", 外呼上面无目标8 := "中间变量2"."1号梯外呼上面无目标8", 外呼上面无目标9 := "中间变量2"."1号梯外呼上面无目标9", 上行停站次数3 := "中间变量2"."1号梯上行停站次数3", 上行停站次数4 := "中间变量2"."1号梯上行停站次数4", 上行停站次数5 := "中间变量2"."1号梯上行停站次数5", 上行停站次数6 := "中间变量2"."1号梯上行停站次数6", 上行停站次数7 := "中间变量2"."1号梯上行停站次数7", 上行停站次数8 := "中间变量2"."1号梯上行停站次数8", 上行停站次数9 := "中间变量2"."1号梯上行停站次数9", 下行停站次数2 := "中间变量2"."1号梯下行停站次数2", 下行停站次数3 := "中间变量2"."1号梯下行停站次数3", 下行停站次数4 := "中间变量2"."1号梯下行停站次数4", 下行停站次数5 := "中间变量2"."1号梯下行停站次数5", 下行停站次数6 := "中间变量2"."1号梯下行停站次数6", 下行停站次数7 := "中间变量2"."1号梯下行停站次数7", 下行停站次数8 := "中间变量2"."1号梯下行停站次数8", 上行停站次数10 := "中间变量2"."1号梯上行停站次数10", 下行停站次数1 := "中间变量2"."1号梯下行停站次数1", 载重量 := "中间变量2"."1号梯转换后载重量", 死机 := "中间变量1".死机1, 限重分配 := "中间变量2".限重分配1, 最终调度距离上1 => "中间变量2"."1梯1层最终调度距离", 最终调度距离上2 => "中间变量2"."1梯2层最终调度距离上", 最终调度距离上3 => "中间变量2"."1梯3层最终调度距离上", 最终调度距离上4 => "中间变量2"."1梯4层最终调度距离上", 最终调度距离上5 => "中间变量2"."1梯5层最终调度距离上", 最终调度距离上6 => "中间变量2"."1梯6层最终调度距离上", 最终调度距离上7 => "中间变量2"."1梯7层最终调度距离上", 最终调度距离上8 => "中间变量2"."1梯8层最终调度距离上", 最终调度距离上9 => "中间变量2"."1梯9层最终调度距离上", 最终调度距离下2 => "中间变量2"."1梯2层最终调度距离下", 最终调度距离下3 => "中间变量2"."1梯3层最终调度距离下", 最终调度距离下4 => "中间变量2"."1梯4层最终调度距离下", 最终调度距离下5 => "中间变量2"."1梯5层最终调度距离下", 最终调度距离下6 => "中间变量2"."1梯6层最终调度距离下", 最终调度距离下7 => "中间变量2"."1梯7层最终调度距离下", 最终调度距离下8 => "中间变量2"."1梯8层最终调度距离下", 最终调度距离下9 => "中间变量2"."1梯9层最终调度距离下", 最终调度距离下10 => "中间变量2"."1梯10层最终调度距离")
   END_RUNG
   // the same network as SCL:
   "1号梯距离调度"(准备就绪 := "中间变量1"."1号梯准备就绪",   // "距离调度"
             检修信号 := "输入"."1号梯检修信号",
             上下平层都为1 := "中间变量1".上下平层同时为1梯1,
             上呼灯1 := "输出"."1层上行呼梯按钮指示灯",
             上呼灯2 := "输出"."2层上行呼梯按钮指示灯",
             上呼灯3 := "输出"."3层上行呼梯按钮指示灯",
             上呼灯4 := "输出"."4层上行呼梯按钮指示灯",
             上呼灯5 := "输出"."5层上行呼梯按钮指示灯",
             上呼灯6 := "输出"."6层上行呼梯按钮指示灯",
             上呼灯7 := "输出"."7层上行呼梯按钮指示灯",
             上呼灯8 := "输出"."8层上行呼梯按钮指示灯",
             上呼灯9 := "输出"."9层上行呼梯按钮指示灯",
             下呼灯2 := "输出"."2层下行呼梯按钮指示灯",
             下呼灯3 := "输出"."3层下行呼梯按钮指示灯",
             下呼灯4 := "输出"."4层下行呼梯按钮指示灯",
             下呼灯5 := "输出"."5层下行呼梯按钮指示灯",
             下呼灯6 := "输出"."6层下行呼梯按钮指示灯",
             下呼灯7 := "输出"."7层下行呼梯按钮指示灯",
             下呼灯8 := "输出"."8层下行呼梯按钮指示灯",
             下呼灯9 := "输出"."9层下行呼梯按钮指示灯",
             下呼灯10 := "输出"."10层下行呼梯按钮指示灯",
             上行指示 := "输出"."1号梯上行指示",
             下行指示 := "输出"."1号梯下行指示",
             当前楼层 := "中间变量2"."1号梯当前楼层数",
             外呼上面有目标最大数1 := "中间变量2"."1号梯外呼上面有目标最大数1",
             外呼上面有目标最大数2 := "中间变量2"."1号梯外呼上面有目标最大数2",
             外呼上面有目标最大数3 := "中间变量2"."1号梯外呼上面有目标最大数3",
             外呼上面有目标最大数4 := "中间变量2"."1号梯外呼上面有目标最大数4",
             外呼上面有目标最大数5 := "中间变量2"."1号梯外呼上面有目标最大数5",
             外呼上面有目标最大数6 := "中间变量2"."1号梯外呼上面有目标最大数6",
             外呼上面有目标最大数7 := "中间变量2"."1号梯外呼上面有目标最大数7",
             外呼上面有目标最大数8 := "中间变量2"."1号梯外呼上面有目标最大数8",
             外呼上面有目标最大数9 := "中间变量2"."1号梯外呼上面有目标最大数9",
             外呼下面有目标最小数2 := "中间变量2"."1号梯外呼下面有目标最小数2",
             外呼下面有目标最小数3 := "中间变量2"."1号梯外呼下面有目标最小数3",
             外呼下面有目标最小数4 := "中间变量2"."1号梯外呼下面有目标最小数4",
             外呼下面有目标最小数5 := "中间变量2"."1号梯外呼下面有目标最小数5",
             外呼下面有目标最小数6 := "中间变量2"."1号梯外呼下面有目标最小数6",
             外呼下面有目标最小数7 := "中间变量2"."1号梯外呼下面有目标最小数7",
             外呼下面有目标最小数8 := "中间变量2"."1号梯外呼下面有目标最小数8",
             外呼下面有目标最小数9 := "中间变量2"."1号梯外呼下面有目标最小数9",
             外呼下面有目标最小数10 := "中间变量2"."1号梯外呼下面有目标最小数10",
             外呼下面有目标2 := "中间变量2"."1号梯外呼下面有目标2",
             外呼下面有目标3 := "中间变量2"."1号梯外呼下面有目标3",
             外呼下面有目标4 := "中间变量2"."1号梯外呼下面有目标4",
             外呼下面有目标5 := "中间变量2"."1号梯外呼下面有目标5",
             外呼下面有目标6 := "中间变量2"."1号梯外呼下面有目标6",
             外呼下面有目标7 := "中间变量2"."1号梯外呼下面有目标7",
             外呼下面有目标8 := "中间变量2"."1号梯外呼下面有目标8",
             外呼下面有目标9 := "中间变量2"."1号梯外呼下面有目标9",
             外呼下面有目标10 := "中间变量2"."1号梯外呼下面有目标10",
             外呼上面有目标1 := "中间变量2"."1号梯外呼上面有目标1",
             外呼上面有目标2 := "中间变量2"."1号梯外呼上面有目标2",
             外呼上面有目标3 := "中间变量2"."1号梯外呼上面有目标3",
             外呼上面有目标4 := "中间变量2"."1号梯外呼上面有目标4",
             外呼上面有目标5 := "中间变量2"."1号梯外呼上面有目标5",
             外呼上面有目标6 := "中间变量2"."1号梯外呼上面有目标6",
             外呼上面有目标7 := "中间变量2"."1号梯外呼上面有目标7",
             外呼上面有目标8 := "中间变量2"."1号梯外呼上面有目标8",
             外呼上面有目标9 := "中间变量2"."1号梯外呼上面有目标9",
             外呼下面无目标2 := "中间变量2"."1号梯外呼下面无目标2",
             外呼下面无目标3 := "中间变量2"."1号梯外呼下面无目标3",
             外呼下面无目标4 := "中间变量2"."1号梯外呼下面无目标4",
             外呼下面无目标5 := "中间变量2"."1号梯外呼下面无目标5",
             外呼下面无目标6 := "中间变量2"."1号梯外呼下面无目标6",
             外呼下面无目标7 := "中间变量2"."1号梯外呼下面无目标7",
             外呼下面无目标8 := "中间变量2"."1号梯外呼下面无目标8",
             外呼下面无目标9 := "中间变量2"."1号梯外呼下面无目标9",
             外呼上面无目标2 := "中间变量2"."1号梯外呼上面无目标2",
             外呼上面无目标3 := "中间变量2"."1号梯外呼上面无目标3",
             外呼上面无目标4 := "中间变量2"."1号梯外呼上面无目标4",
             外呼上面无目标5 := "中间变量2"."1号梯外呼上面无目标5",
             外呼上面无目标6 := "中间变量2"."1号梯外呼上面无目标6",
             外呼上面无目标7 := "中间变量2"."1号梯外呼上面无目标7",
             外呼上面无目标8 := "中间变量2"."1号梯外呼上面无目标8",
             外呼上面无目标9 := "中间变量2"."1号梯外呼上面无目标9",
             上行停站次数3 := "中间变量2"."1号梯上行停站次数3",
             上行停站次数4 := "中间变量2"."1号梯上行停站次数4",
             上行停站次数5 := "中间变量2"."1号梯上行停站次数5",
             上行停站次数6 := "中间变量2"."1号梯上行停站次数6",
             上行停站次数7 := "中间变量2"."1号梯上行停站次数7",
             上行停站次数8 := "中间变量2"."1号梯上行停站次数8",
             上行停站次数9 := "中间变量2"."1号梯上行停站次数9",
             下行停站次数2 := "中间变量2"."1号梯下行停站次数2",
             下行停站次数3 := "中间变量2"."1号梯下行停站次数3",
             下行停站次数4 := "中间变量2"."1号梯下行停站次数4",
             下行停站次数5 := "中间变量2"."1号梯下行停站次数5",
             下行停站次数6 := "中间变量2"."1号梯下行停站次数6",
             下行停站次数7 := "中间变量2"."1号梯下行停站次数7",
             下行停站次数8 := "中间变量2"."1号梯下行停站次数8",
             上行停站次数10 := "中间变量2"."1号梯上行停站次数10",
             下行停站次数1 := "中间变量2"."1号梯下行停站次数1",
             载重量 := "中间变量2"."1号梯转换后载重量",
             死机 := "中间变量1".死机1,
             限重分配 := "中间变量2".限重分配1,
             最终调度距离上1 => "中间变量2"."1梯1层最终调度距离",
             最终调度距离上2 => "中间变量2"."1梯2层最终调度距离上",
             最终调度距离上3 => "中间变量2"."1梯3层最终调度距离上",
             最终调度距离上4 => "中间变量2"."1梯4层最终调度距离上",
             最终调度距离上5 => "中间变量2"."1梯5层最终调度距离上",
             最终调度距离上6 => "中间变量2"."1梯6层最终调度距离上",
             最终调度距离上7 => "中间变量2"."1梯7层最终调度距离上",
             最终调度距离上8 => "中间变量2"."1梯8层最终调度距离上",
             最终调度距离上9 => "中间变量2"."1梯9层最终调度距离上",
             最终调度距离下2 => "中间变量2"."1梯2层最终调度距离下",
             最终调度距离下3 => "中间变量2"."1梯3层最终调度距离下",
             最终调度距离下4 => "中间变量2"."1梯4层最终调度距离下",
             最终调度距离下5 => "中间变量2"."1梯5层最终调度距离下",
             最终调度距离下6 => "中间变量2"."1梯6层最终调度距离下",
             最终调度距离下7 => "中间变量2"."1梯7层最终调度距离下",
             最终调度距离下8 => "中间变量2"."1梯8层最终调度距离下",
             最终调度距离下9 => "中间变量2"."1梯9层最终调度距离下",
             最终调度距离下10 => "中间变量2"."1梯10层最终调度距离");
END_REGION

REGION Network 3: 2号梯调度距离
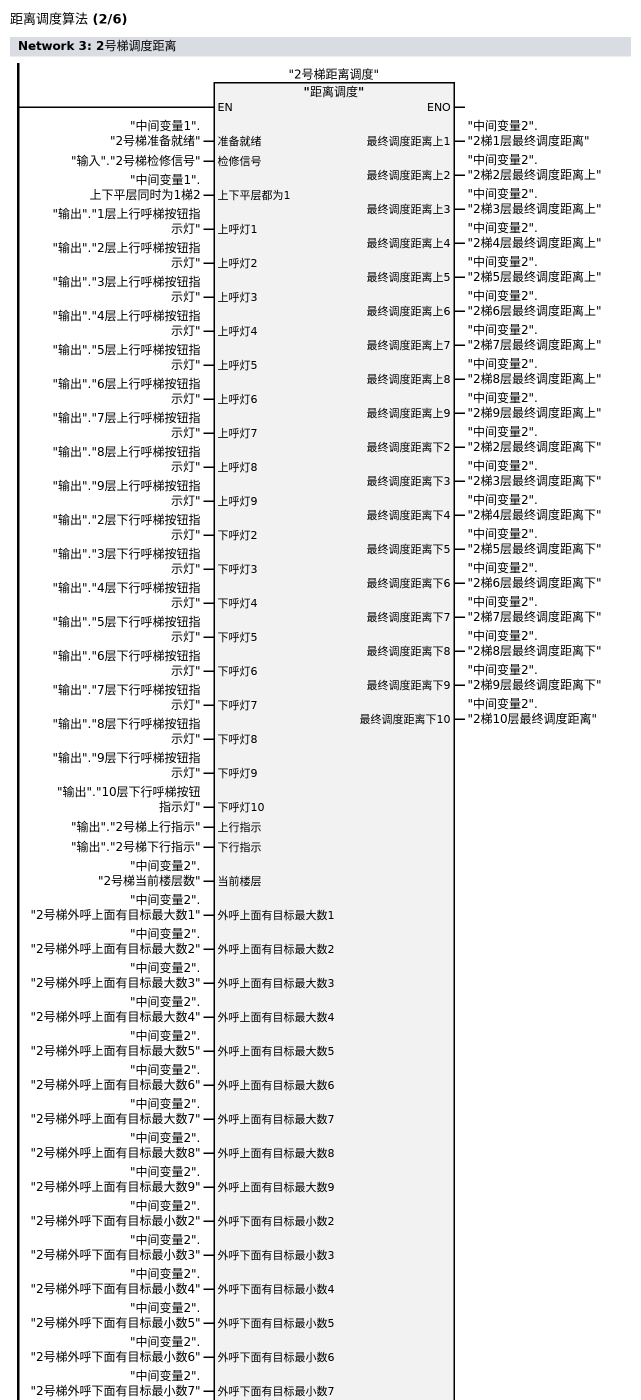
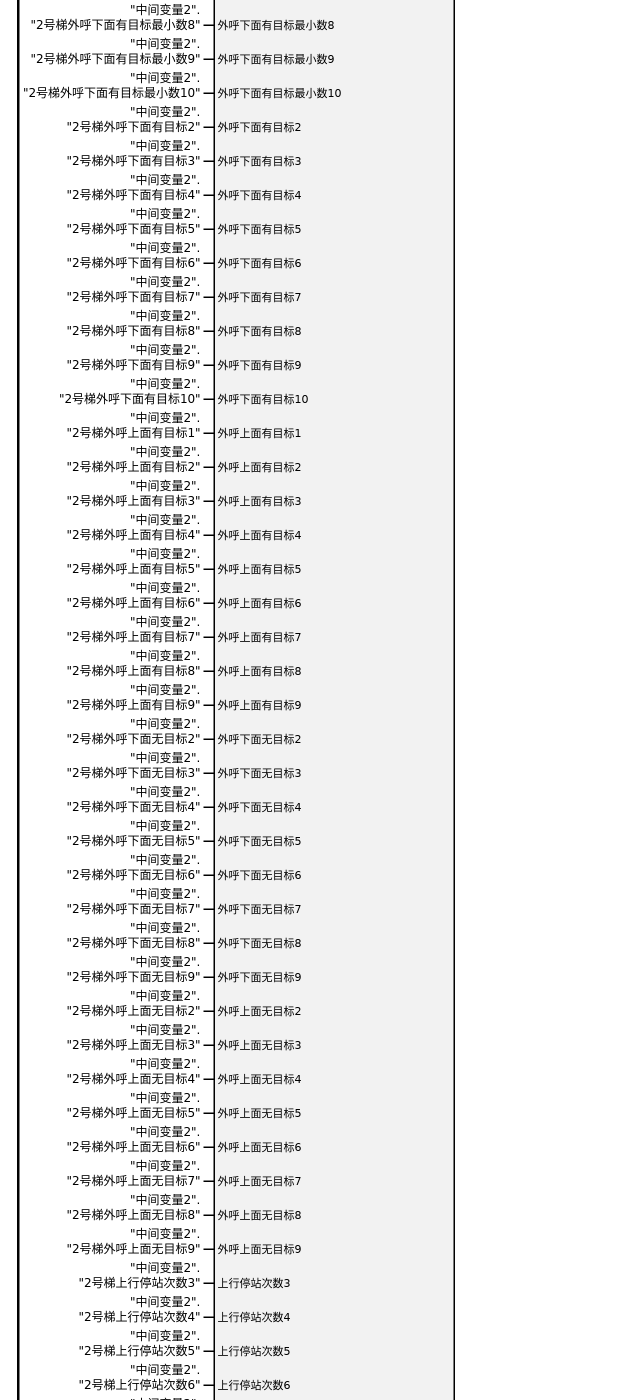
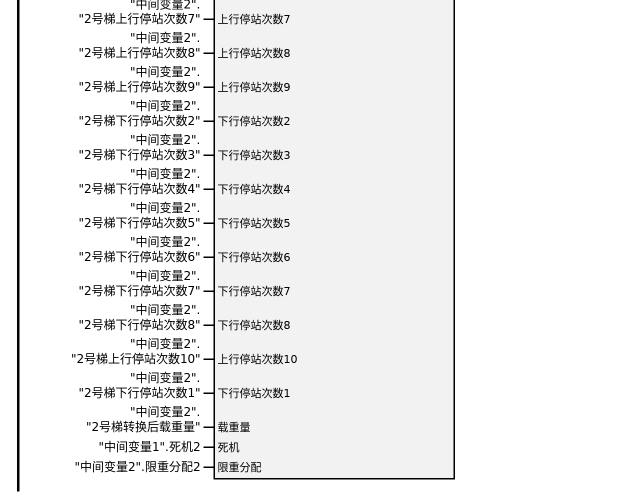
   RUNG wire#powerrail
      "2号梯距离调度"(准备就绪 := "中间变量1"."2号梯准备就绪", 检修信号 := "输入"."2号梯检修信号", 上下平层都为1 := "中间变量1".上下平层同时为1梯2, 上呼灯1 := "输出"."1层上行呼梯按钮指示灯", 上呼灯2 := "输出"."2层上行呼梯按钮指示灯", 上呼灯3 := "输出"."3层上行呼梯按钮指示灯", 上呼灯4 := "输出"."4层上行呼梯按钮指示灯", 上呼灯5 := "输出"."5层上行呼梯按钮指示灯", 上呼灯6 := "输出"."6层上行呼梯按钮指示灯", 上呼灯7 := "输出"."7层上行呼梯按钮指示灯", 上呼灯8 := "输出"."8层上行呼梯按钮指示灯", 上呼灯9 := "输出"."9层上行呼梯按钮指示灯", 下呼灯2 := "输出"."2层下行呼梯按钮指示灯", 下呼灯3 := "输出"."3层下行呼梯按钮指示灯", 下呼灯4 := "输出"."4层下行呼梯按钮指示灯", 下呼灯5 := "输出"."5层下行呼梯按钮指示灯", 下呼灯6 := "输出"."6层下行呼梯按钮指示灯", 下呼灯7 := "输出"."7层下行呼梯按钮指示灯", 下呼灯8 := "输出"."8层下行呼梯按钮指示灯", 下呼灯9 := "输出"."9层下行呼梯按钮指示灯", 下呼灯10 := "输出"."10层下行呼梯按钮指示灯", 上行指示 := "输出"."2号梯上行指示", 下行指示 := "输出"."2号梯下行指示", 当前楼层 := "中间变量2"."2号梯当前楼层数", 外呼上面有目标最大数1 := "中间变量2"."2号梯外呼上面有目标最大数1", 外呼上面有目标最大数2 := "中间变量2"."2号梯外呼上面有目标最大数2", 外呼上面有目标最大数3 := "中间变量2"."2号梯外呼上面有目标最大数3", 外呼上面有目标最大数4 := "中间变量2"."2号梯外呼上面有目标最大数4", 外呼上面有目标最大数5 := "中间变量2"."2号梯外呼上面有目标最大数5", 外呼上面有目标最大数6 := "中间变量2"."2号梯外呼上面有目标最大数6", 外呼上面有目标最大数7 := "中间变量2"."2号梯外呼上面有目标最大数7", 外呼上面有目标最大数8 := "中间变量2"."2号梯外呼上面有目标最大数8", 外呼上面有目标最大数9 := "中间变量2"."2号梯外呼上面有目标最大数9", 外呼下面有目标最小数2 := "中间变量2"."2号梯外呼下面有目标最小数2", 外呼下面有目标最小数3 := "中间变量2"."2号梯外呼下面有目标最小数3", 外呼下面有目标最小数4 := "中间变量2"."2号梯外呼下面有目标最小数4", 外呼下面有目标最小数5 := "中间变量2"."2号梯外呼下面有目标最小数5", 外呼下面有目标最小数6 := "中间变量2"."2号梯外呼下面有目标最小数6", 外呼下面有目标最小数7 := "中间变量2"."2号梯外呼下面有目标最小数7", 外呼下面有目标最小数8 := "中间变量2"."2号梯外呼下面有目标最小数8", 外呼下面有目标最小数9 := "中间变量2"."2号梯外呼下面有目标最小数9", 外呼下面有目标最小数10 := "中间变量2"."2号梯外呼下面有目标最小数10", 外呼下面有目标2 := "中间变量2"."2号梯外呼下面有目标2", 外呼下面有目标3 := "中间变量2"."2号梯外呼下面有目标3", 外呼下面有目标4 := "中间变量2"."2号梯外呼下面有目标4", 外呼下面有目标5 := "中间变量2"."2号梯外呼下面有目标5", 外呼下面有目标6 := "中间变量2"."2号梯外呼下面有目标6", 外呼下面有目标7 := "中间变量2"."2号梯外呼下面有目标7", 外呼下面有目标8 := "中间变量2"."2号梯外呼下面有目标8", 外呼下面有目标9 := "中间变量2"."2号梯外呼下面有目标9", 外呼下面有目标10 := "中间变量2"."2号梯外呼下面有目标10", 外呼上面有目标1 := "中间变量2"."2号梯外呼上面有目标1", 外呼上面有目标2 := "中间变量2"."2号梯外呼上面有目标2", 外呼上面有目标3 := "中间变量2"."2号梯外呼上面有目标3", 外呼上面有目标4 := "中间变量2"."2号梯外呼上面有目标4", 外呼上面有目标5 := "中间变量2"."2号梯外呼上面有目标5", 外呼上面有目标6 := "中间变量2"."2号梯外呼上面有目标6", 外呼上面有目标7 := "中间变量2"."2号梯外呼上面有目标7", 外呼上面有目标8 := "中间变量2"."2号梯外呼上面有目标8", 外呼上面有目标9 := "中间变量2"."2号梯外呼上面有目标9", 外呼下面无目标2 := "中间变量2"."2号梯外呼下面无目标2", 外呼下面无目标3 := "中间变量2"."2号梯外呼下面无目标3", 外呼下面无目标4 := "中间变量2"."2号梯外呼下面无目标4", 外呼下面无目标5 := "中间变量2"."2号梯外呼下面无目标5", 外呼下面无目标6 := "中间变量2"."2号梯外呼下面无目标6", 外呼下面无目标7 := "中间变量2"."2号梯外呼下面无目标7", 外呼下面无目标8 := "中间变量2"."2号梯外呼下面无目标8", 外呼下面无目标9 := "中间变量2"."2号梯外呼下面无目标9", 外呼上面无目标2 := "中间变量2"."2号梯外呼上面无目标2", 外呼上面无目标3 := "中间变量2"."2号梯外呼上面无目标3", 外呼上面无目标4 := "中间变量2"."2号梯外呼上面无目标4", 外呼上面无目标5 := "中间变量2"."2号梯外呼上面无目标5", 外呼上面无目标6 := "中间变量2"."2号梯外呼上面无目标6", 外呼上面无目标7 := "中间变量2"."2号梯外呼上面无目标7", 外呼上面无目标8 := "中间变量2"."2号梯外呼上面无目标8", 外呼上面无目标9 := "中间变量2"."2号梯外呼上面无目标9", 上行停站次数3 := "中间变量2"."2号梯上行停站次数3", 上行停站次数4 := "中间变量2"."2号梯上行停站次数4", 上行停站次数5 := "中间变量2"."2号梯上行停站次数5", 上行停站次数6 := "中间变量2"."2号梯上行停站次数6", 上行停站次数7 := "中间变量2"."2号梯上行停站次数7", 上行停站次数8 := "中间变量2"."2号梯上行停站次数8", 上行停站次数9 := "中间变量2"."2号梯上行停站次数9", 下行停站次数2 := "中间变量2"."2号梯下行停站次数2", 下行停站次数3 := "中间变量2"."2号梯下行停站次数3", 下行停站次数4 := "中间变量2"."2号梯下行停站次数4", 下行停站次数5 := "中间变量2"."2号梯下行停站次数5", 下行停站次数6 := "中间变量2"."2号梯下行停站次数6", 下行停站次数7 := "中间变量2"."2号梯下行停站次数7", 下行停站次数8 := "中间变量2"."2号梯下行停站次数8", 上行停站次数10 := "中间变量2"."2号梯上行停站次数10", 下行停站次数1 := "中间变量2"."2号梯下行停站次数1", 载重量 := "中间变量2"."2号梯转换后载重量", 死机 := "中间变量1".死机2, 限重分配 := "中间变量2".限重分配2, 最终调度距离上1 => "中间变量2"."2梯1层最终调度距离", 最终调度距离上2 => "中间变量2"."2梯2层最终调度距离上", 最终调度距离上3 => "中间变量2"."2梯3层最终调度距离上", 最终调度距离上4 => "中间变量2"."2梯4层最终调度距离上", 最终调度距离上5 => "中间变量2"."2梯5层最终调度距离上", 最终调度距离上6 => "中间变量2"."2梯6层最终调度距离上", 最终调度距离上7 => "中间变量2"."2梯7层最终调度距离上", 最终调度距离上8 => "中间变量2"."2梯8层最终调度距离上", 最终调度距离上9 => "中间变量2"."2梯9层最终调度距离上", 最终调度距离下2 => "中间变量2"."2梯2层最终调度距离下", 最终调度距离下3 => "中间变量2"."2梯3层最终调度距离下", 最终调度距离下4 => "中间变量2"."2梯4层最终调度距离下", 最终调度距离下5 => "中间变量2"."2梯5层最终调度距离下", 最终调度距离下6 => "中间变量2"."2梯6层最终调度距离下", 最终调度距离下7 => "中间变量2"."2梯7层最终调度距离下", 最终调度距离下8 => "中间变量2"."2梯8层最终调度距离下", 最终调度距离下9 => "中间变量2"."2梯9层最终调度距离下", 最终调度距离下10 => "中间变量2"."2梯10层最终调度距离")
   END_RUNG
   // the same network as SCL:
   "2号梯距离调度"(准备就绪 := "中间变量1"."2号梯准备就绪",   // "距离调度"
             检修信号 := "输入"."2号梯检修信号",
             上下平层都为1 := "中间变量1".上下平层同时为1梯2,
             上呼灯1 := "输出"."1层上行呼梯按钮指示灯",
             上呼灯2 := "输出"."2层上行呼梯按钮指示灯",
             上呼灯3 := "输出"."3层上行呼梯按钮指示灯",
             上呼灯4 := "输出"."4层上行呼梯按钮指示灯",
             上呼灯5 := "输出"."5层上行呼梯按钮指示灯",
             上呼灯6 := "输出"."6层上行呼梯按钮指示灯",
             上呼灯7 := "输出"."7层上行呼梯按钮指示灯",
             上呼灯8 := "输出"."8层上行呼梯按钮指示灯",
             上呼灯9 := "输出"."9层上行呼梯按钮指示灯",
             下呼灯2 := "输出"."2层下行呼梯按钮指示灯",
             下呼灯3 := "输出"."3层下行呼梯按钮指示灯",
             下呼灯4 := "输出"."4层下行呼梯按钮指示灯",
             下呼灯5 := "输出"."5层下行呼梯按钮指示灯",
             下呼灯6 := "输出"."6层下行呼梯按钮指示灯",
             下呼灯7 := "输出"."7层下行呼梯按钮指示灯",
             下呼灯8 := "输出"."8层下行呼梯按钮指示灯",
             下呼灯9 := "输出"."9层下行呼梯按钮指示灯",
             下呼灯10 := "输出"."10层下行呼梯按钮指示灯",
             上行指示 := "输出"."2号梯上行指示",
             下行指示 := "输出"."2号梯下行指示",
             当前楼层 := "中间变量2"."2号梯当前楼层数",
             外呼上面有目标最大数1 := "中间变量2"."2号梯外呼上面有目标最大数1",
             外呼上面有目标最大数2 := "中间变量2"."2号梯外呼上面有目标最大数2",
             外呼上面有目标最大数3 := "中间变量2"."2号梯外呼上面有目标最大数3",
             外呼上面有目标最大数4 := "中间变量2"."2号梯外呼上面有目标最大数4",
             外呼上面有目标最大数5 := "中间变量2"."2号梯外呼上面有目标最大数5",
             外呼上面有目标最大数6 := "中间变量2"."2号梯外呼上面有目标最大数6",
             外呼上面有目标最大数7 := "中间变量2"."2号梯外呼上面有目标最大数7",
             外呼上面有目标最大数8 := "中间变量2"."2号梯外呼上面有目标最大数8",
             外呼上面有目标最大数9 := "中间变量2"."2号梯外呼上面有目标最大数9",
             外呼下面有目标最小数2 := "中间变量2"."2号梯外呼下面有目标最小数2",
             外呼下面有目标最小数3 := "中间变量2"."2号梯外呼下面有目标最小数3",
             外呼下面有目标最小数4 := "中间变量2"."2号梯外呼下面有目标最小数4",
             外呼下面有目标最小数5 := "中间变量2"."2号梯外呼下面有目标最小数5",
             外呼下面有目标最小数6 := "中间变量2"."2号梯外呼下面有目标最小数6",
             外呼下面有目标最小数7 := "中间变量2"."2号梯外呼下面有目标最小数7",
             外呼下面有目标最小数8 := "中间变量2"."2号梯外呼下面有目标最小数8",
             外呼下面有目标最小数9 := "中间变量2"."2号梯外呼下面有目标最小数9",
             外呼下面有目标最小数10 := "中间变量2"."2号梯外呼下面有目标最小数10",
             外呼下面有目标2 := "中间变量2"."2号梯外呼下面有目标2",
             外呼下面有目标3 := "中间变量2"."2号梯外呼下面有目标3",
             外呼下面有目标4 := "中间变量2"."2号梯外呼下面有目标4",
             外呼下面有目标5 := "中间变量2"."2号梯外呼下面有目标5",
             外呼下面有目标6 := "中间变量2"."2号梯外呼下面有目标6",
             外呼下面有目标7 := "中间变量2"."2号梯外呼下面有目标7",
             外呼下面有目标8 := "中间变量2"."2号梯外呼下面有目标8",
             外呼下面有目标9 := "中间变量2"."2号梯外呼下面有目标9",
             外呼下面有目标10 := "中间变量2"."2号梯外呼下面有目标10",
             外呼上面有目标1 := "中间变量2"."2号梯外呼上面有目标1",
             外呼上面有目标2 := "中间变量2"."2号梯外呼上面有目标2",
             外呼上面有目标3 := "中间变量2"."2号梯外呼上面有目标3",
             外呼上面有目标4 := "中间变量2"."2号梯外呼上面有目标4",
             外呼上面有目标5 := "中间变量2"."2号梯外呼上面有目标5",
             外呼上面有目标6 := "中间变量2"."2号梯外呼上面有目标6",
             外呼上面有目标7 := "中间变量2"."2号梯外呼上面有目标7",
             外呼上面有目标8 := "中间变量2"."2号梯外呼上面有目标8",
             外呼上面有目标9 := "中间变量2"."2号梯外呼上面有目标9",
             外呼下面无目标2 := "中间变量2"."2号梯外呼下面无目标2",
             外呼下面无目标3 := "中间变量2"."2号梯外呼下面无目标3",
             外呼下面无目标4 := "中间变量2"."2号梯外呼下面无目标4",
             外呼下面无目标5 := "中间变量2"."2号梯外呼下面无目标5",
             外呼下面无目标6 := "中间变量2"."2号梯外呼下面无目标6",
             外呼下面无目标7 := "中间变量2"."2号梯外呼下面无目标7",
             外呼下面无目标8 := "中间变量2"."2号梯外呼下面无目标8",
             外呼下面无目标9 := "中间变量2"."2号梯外呼下面无目标9",
             外呼上面无目标2 := "中间变量2"."2号梯外呼上面无目标2",
             外呼上面无目标3 := "中间变量2"."2号梯外呼上面无目标3",
             外呼上面无目标4 := "中间变量2"."2号梯外呼上面无目标4",
             外呼上面无目标5 := "中间变量2"."2号梯外呼上面无目标5",
             外呼上面无目标6 := "中间变量2"."2号梯外呼上面无目标6",
             外呼上面无目标7 := "中间变量2"."2号梯外呼上面无目标7",
             外呼上面无目标8 := "中间变量2"."2号梯外呼上面无目标8",
             外呼上面无目标9 := "中间变量2"."2号梯外呼上面无目标9",
             上行停站次数3 := "中间变量2"."2号梯上行停站次数3",
             上行停站次数4 := "中间变量2"."2号梯上行停站次数4",
             上行停站次数5 := "中间变量2"."2号梯上行停站次数5",
             上行停站次数6 := "中间变量2"."2号梯上行停站次数6",
             上行停站次数7 := "中间变量2"."2号梯上行停站次数7",
             上行停站次数8 := "中间变量2"."2号梯上行停站次数8",
             上行停站次数9 := "中间变量2"."2号梯上行停站次数9",
             下行停站次数2 := "中间变量2"."2号梯下行停站次数2",
             下行停站次数3 := "中间变量2"."2号梯下行停站次数3",
             下行停站次数4 := "中间变量2"."2号梯下行停站次数4",
             下行停站次数5 := "中间变量2"."2号梯下行停站次数5",
             下行停站次数6 := "中间变量2"."2号梯下行停站次数6",
             下行停站次数7 := "中间变量2"."2号梯下行停站次数7",
             下行停站次数8 := "中间变量2"."2号梯下行停站次数8",
             上行停站次数10 := "中间变量2"."2号梯上行停站次数10",
             下行停站次数1 := "中间变量2"."2号梯下行停站次数1",
             载重量 := "中间变量2"."2号梯转换后载重量",
             死机 := "中间变量1".死机2,
             限重分配 := "中间变量2".限重分配2,
             最终调度距离上1 => "中间变量2"."2梯1层最终调度距离",
             最终调度距离上2 => "中间变量2"."2梯2层最终调度距离上",
             最终调度距离上3 => "中间变量2"."2梯3层最终调度距离上",
             最终调度距离上4 => "中间变量2"."2梯4层最终调度距离上",
             最终调度距离上5 => "中间变量2"."2梯5层最终调度距离上",
             最终调度距离上6 => "中间变量2"."2梯6层最终调度距离上",
             最终调度距离上7 => "中间变量2"."2梯7层最终调度距离上",
             最终调度距离上8 => "中间变量2"."2梯8层最终调度距离上",
             最终调度距离上9 => "中间变量2"."2梯9层最终调度距离上",
             最终调度距离下2 => "中间变量2"."2梯2层最终调度距离下",
             最终调度距离下3 => "中间变量2"."2梯3层最终调度距离下",
             最终调度距离下4 => "中间变量2"."2梯4层最终调度距离下",
             最终调度距离下5 => "中间变量2"."2梯5层最终调度距离下",
             最终调度距离下6 => "中间变量2"."2梯6层最终调度距离下",
             最终调度距离下7 => "中间变量2"."2梯7层最终调度距离下",
             最终调度距离下8 => "中间变量2"."2梯8层最终调度距离下",
             最终调度距离下9 => "中间变量2"."2梯9层最终调度距离下",
             最终调度距离下10 => "中间变量2"."2梯10层最终调度距离");
END_REGION

REGION Network 4: 3号梯调度距离
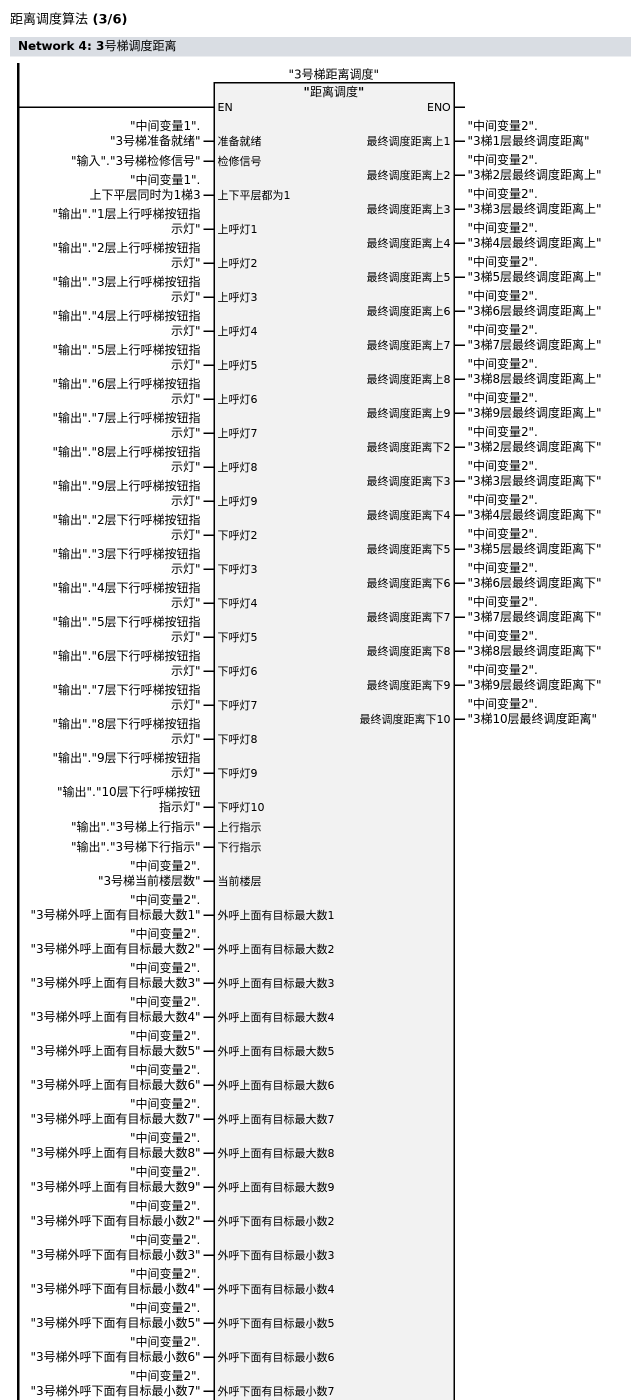
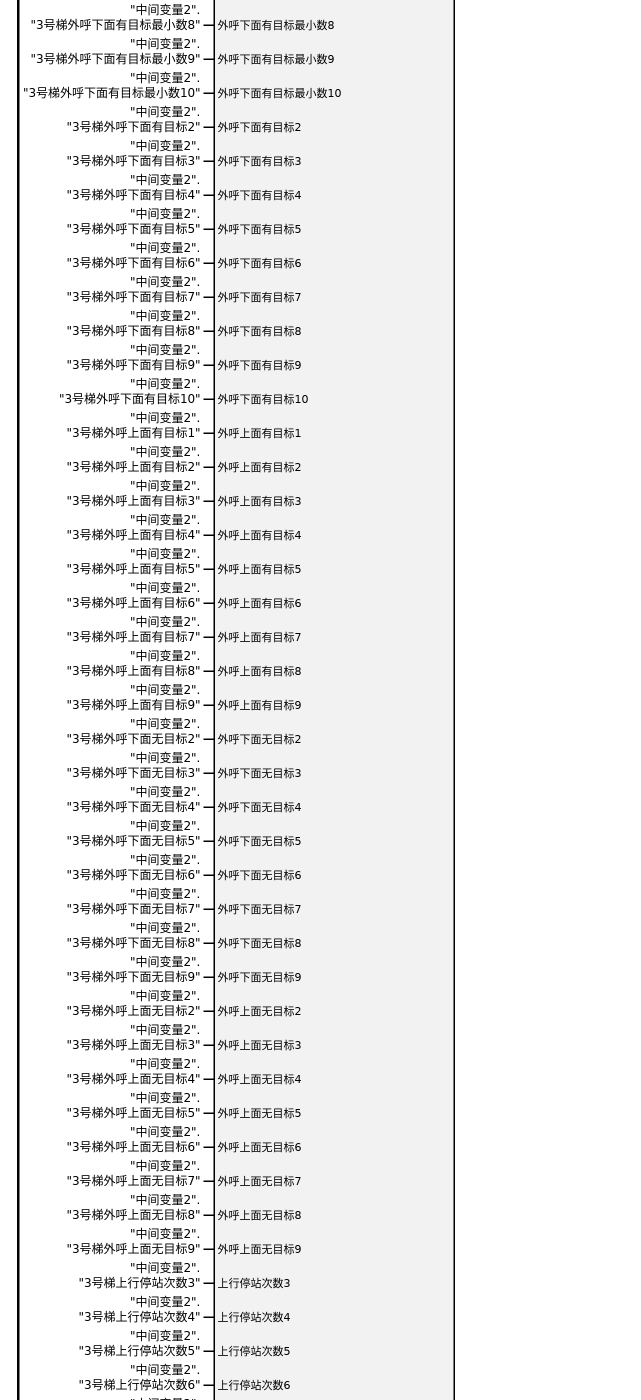
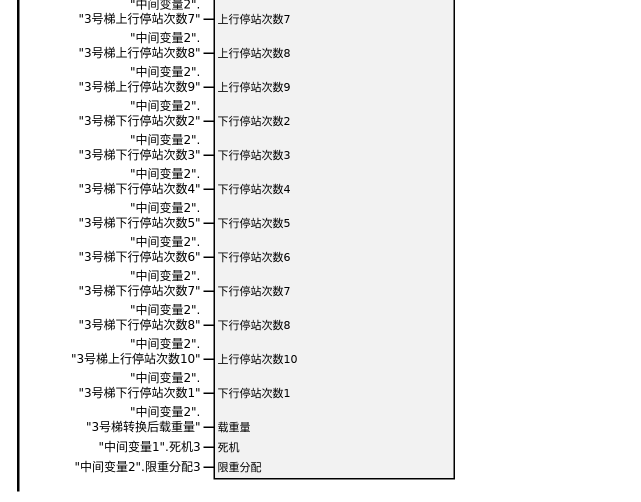
   RUNG wire#powerrail
      "3号梯距离调度"(准备就绪 := "中间变量1"."3号梯准备就绪", 检修信号 := "输入"."3号梯检修信号", 上下平层都为1 := "中间变量1".上下平层同时为1梯3, 上呼灯1 := "输出"."1层上行呼梯按钮指示灯", 上呼灯2 := "输出"."2层上行呼梯按钮指示灯", 上呼灯3 := "输出"."3层上行呼梯按钮指示灯", 上呼灯4 := "输出"."4层上行呼梯按钮指示灯", 上呼灯5 := "输出"."5层上行呼梯按钮指示灯", 上呼灯6 := "输出"."6层上行呼梯按钮指示灯", 上呼灯7 := "输出"."7层上行呼梯按钮指示灯", 上呼灯8 := "输出"."8层上行呼梯按钮指示灯", 上呼灯9 := "输出"."9层上行呼梯按钮指示灯", 下呼灯2 := "输出"."2层下行呼梯按钮指示灯", 下呼灯3 := "输出"."3层下行呼梯按钮指示灯", 下呼灯4 := "输出"."4层下行呼梯按钮指示灯", 下呼灯5 := "输出"."5层下行呼梯按钮指示灯", 下呼灯6 := "输出"."6层下行呼梯按钮指示灯", 下呼灯7 := "输出"."7层下行呼梯按钮指示灯", 下呼灯8 := "输出"."8层下行呼梯按钮指示灯", 下呼灯9 := "输出"."9层下行呼梯按钮指示灯", 下呼灯10 := "输出"."10层下行呼梯按钮指示灯", 上行指示 := "输出"."3号梯上行指示", 下行指示 := "输出"."3号梯下行指示", 当前楼层 := "中间变量2"."3号梯当前楼层数", 外呼上面有目标最大数1 := "中间变量2"."3号梯外呼上面有目标最大数1", 外呼上面有目标最大数2 := "中间变量2"."3号梯外呼上面有目标最大数2", 外呼上面有目标最大数3 := "中间变量2"."3号梯外呼上面有目标最大数3", 外呼上面有目标最大数4 := "中间变量2"."3号梯外呼上面有目标最大数4", 外呼上面有目标最大数5 := "中间变量2"."3号梯外呼上面有目标最大数5", 外呼上面有目标最大数6 := "中间变量2"."3号梯外呼上面有目标最大数6", 外呼上面有目标最大数7 := "中间变量2"."3号梯外呼上面有目标最大数7", 外呼上面有目标最大数8 := "中间变量2"."3号梯外呼上面有目标最大数8", 外呼上面有目标最大数9 := "中间变量2"."3号梯外呼上面有目标最大数9", 外呼下面有目标最小数2 := "中间变量2"."3号梯外呼下面有目标最小数2", 外呼下面有目标最小数3 := "中间变量2"."3号梯外呼下面有目标最小数3", 外呼下面有目标最小数4 := "中间变量2"."3号梯外呼下面有目标最小数4", 外呼下面有目标最小数5 := "中间变量2"."3号梯外呼下面有目标最小数5", 外呼下面有目标最小数6 := "中间变量2"."3号梯外呼下面有目标最小数6", 外呼下面有目标最小数7 := "中间变量2"."3号梯外呼下面有目标最小数7", 外呼下面有目标最小数8 := "中间变量2"."3号梯外呼下面有目标最小数8", 外呼下面有目标最小数9 := "中间变量2"."3号梯外呼下面有目标最小数9", 外呼下面有目标最小数10 := "中间变量2"."3号梯外呼下面有目标最小数10", 外呼下面有目标2 := "中间变量2"."3号梯外呼下面有目标2", 外呼下面有目标3 := "中间变量2"."3号梯外呼下面有目标3", 外呼下面有目标4 := "中间变量2"."3号梯外呼下面有目标4", 外呼下面有目标5 := "中间变量2"."3号梯外呼下面有目标5", 外呼下面有目标6 := "中间变量2"."3号梯外呼下面有目标6", 外呼下面有目标7 := "中间变量2"."3号梯外呼下面有目标7", 外呼下面有目标8 := "中间变量2"."3号梯外呼下面有目标8", 外呼下面有目标9 := "中间变量2"."3号梯外呼下面有目标9", 外呼下面有目标10 := "中间变量2"."3号梯外呼下面有目标10", 外呼上面有目标1 := "中间变量2"."3号梯外呼上面有目标1", 外呼上面有目标2 := "中间变量2"."3号梯外呼上面有目标2", 外呼上面有目标3 := "中间变量2"."3号梯外呼上面有目标3", 外呼上面有目标4 := "中间变量2"."3号梯外呼上面有目标4", 外呼上面有目标5 := "中间变量2"."3号梯外呼上面有目标5", 外呼上面有目标6 := "中间变量2"."3号梯外呼上面有目标6", 外呼上面有目标7 := "中间变量2"."3号梯外呼上面有目标7", 外呼上面有目标8 := "中间变量2"."3号梯外呼上面有目标8", 外呼上面有目标9 := "中间变量2"."3号梯外呼上面有目标9", 外呼下面无目标2 := "中间变量2"."3号梯外呼下面无目标2", 外呼下面无目标3 := "中间变量2"."3号梯外呼下面无目标3", 外呼下面无目标4 := "中间变量2"."3号梯外呼下面无目标4", 外呼下面无目标5 := "中间变量2"."3号梯外呼下面无目标5", 外呼下面无目标6 := "中间变量2"."3号梯外呼下面无目标6", 外呼下面无目标7 := "中间变量2"."3号梯外呼下面无目标7", 外呼下面无目标8 := "中间变量2"."3号梯外呼下面无目标8", 外呼下面无目标9 := "中间变量2"."3号梯外呼下面无目标9", 外呼上面无目标2 := "中间变量2"."3号梯外呼上面无目标2", 外呼上面无目标3 := "中间变量2"."3号梯外呼上面无目标3", 外呼上面无目标4 := "中间变量2"."3号梯外呼上面无目标4", 外呼上面无目标5 := "中间变量2"."3号梯外呼上面无目标5", 外呼上面无目标6 := "中间变量2"."3号梯外呼上面无目标6", 外呼上面无目标7 := "中间变量2"."3号梯外呼上面无目标7", 外呼上面无目标8 := "中间变量2"."3号梯外呼上面无目标8", 外呼上面无目标9 := "中间变量2"."3号梯外呼上面无目标9", 上行停站次数3 := "中间变量2"."3号梯上行停站次数3", 上行停站次数4 := "中间变量2"."3号梯上行停站次数4", 上行停站次数5 := "中间变量2"."3号梯上行停站次数5", 上行停站次数6 := "中间变量2"."3号梯上行停站次数6", 上行停站次数7 := "中间变量2"."3号梯上行停站次数7", 上行停站次数8 := "中间变量2"."3号梯上行停站次数8", 上行停站次数9 := "中间变量2"."3号梯上行停站次数9", 下行停站次数2 := "中间变量2"."3号梯下行停站次数2", 下行停站次数3 := "中间变量2"."3号梯下行停站次数3", 下行停站次数4 := "中间变量2"."3号梯下行停站次数4", 下行停站次数5 := "中间变量2"."3号梯下行停站次数5", 下行停站次数6 := "中间变量2"."3号梯下行停站次数6", 下行停站次数7 := "中间变量2"."3号梯下行停站次数7", 下行停站次数8 := "中间变量2"."3号梯下行停站次数8", 上行停站次数10 := "中间变量2"."3号梯上行停站次数10", 下行停站次数1 := "中间变量2"."3号梯下行停站次数1", 载重量 := "中间变量2"."3号梯转换后载重量", 死机 := "中间变量1".死机3, 限重分配 := "中间变量2".限重分配3, 最终调度距离上1 => "中间变量2"."3梯1层最终调度距离", 最终调度距离上2 => "中间变量2"."3梯2层最终调度距离上", 最终调度距离上3 => "中间变量2"."3梯3层最终调度距离上", 最终调度距离上4 => "中间变量2"."3梯4层最终调度距离上", 最终调度距离上5 => "中间变量2"."3梯5层最终调度距离上", 最终调度距离上6 => "中间变量2"."3梯6层最终调度距离上", 最终调度距离上7 => "中间变量2"."3梯7层最终调度距离上", 最终调度距离上8 => "中间变量2"."3梯8层最终调度距离上", 最终调度距离上9 => "中间变量2"."3梯9层最终调度距离上", 最终调度距离下2 => "中间变量2"."3梯2层最终调度距离下", 最终调度距离下3 => "中间变量2"."3梯3层最终调度距离下", 最终调度距离下4 => "中间变量2"."3梯4层最终调度距离下", 最终调度距离下5 => "中间变量2"."3梯5层最终调度距离下", 最终调度距离下6 => "中间变量2"."3梯6层最终调度距离下", 最终调度距离下7 => "中间变量2"."3梯7层最终调度距离下", 最终调度距离下8 => "中间变量2"."3梯8层最终调度距离下", 最终调度距离下9 => "中间变量2"."3梯9层最终调度距离下", 最终调度距离下10 => "中间变量2"."3梯10层最终调度距离")
   END_RUNG
   // the same network as SCL:
   "3号梯距离调度"(准备就绪 := "中间变量1"."3号梯准备就绪",   // "距离调度"
             检修信号 := "输入"."3号梯检修信号",
             上下平层都为1 := "中间变量1".上下平层同时为1梯3,
             上呼灯1 := "输出"."1层上行呼梯按钮指示灯",
             上呼灯2 := "输出"."2层上行呼梯按钮指示灯",
             上呼灯3 := "输出"."3层上行呼梯按钮指示灯",
             上呼灯4 := "输出"."4层上行呼梯按钮指示灯",
             上呼灯5 := "输出"."5层上行呼梯按钮指示灯",
             上呼灯6 := "输出"."6层上行呼梯按钮指示灯",
             上呼灯7 := "输出"."7层上行呼梯按钮指示灯",
             上呼灯8 := "输出"."8层上行呼梯按钮指示灯",
             上呼灯9 := "输出"."9层上行呼梯按钮指示灯",
             下呼灯2 := "输出"."2层下行呼梯按钮指示灯",
             下呼灯3 := "输出"."3层下行呼梯按钮指示灯",
             下呼灯4 := "输出"."4层下行呼梯按钮指示灯",
             下呼灯5 := "输出"."5层下行呼梯按钮指示灯",
             下呼灯6 := "输出"."6层下行呼梯按钮指示灯",
             下呼灯7 := "输出"."7层下行呼梯按钮指示灯",
             下呼灯8 := "输出"."8层下行呼梯按钮指示灯",
             下呼灯9 := "输出"."9层下行呼梯按钮指示灯",
             下呼灯10 := "输出"."10层下行呼梯按钮指示灯",
             上行指示 := "输出"."3号梯上行指示",
             下行指示 := "输出"."3号梯下行指示",
             当前楼层 := "中间变量2"."3号梯当前楼层数",
             外呼上面有目标最大数1 := "中间变量2"."3号梯外呼上面有目标最大数1",
             外呼上面有目标最大数2 := "中间变量2"."3号梯外呼上面有目标最大数2",
             外呼上面有目标最大数3 := "中间变量2"."3号梯外呼上面有目标最大数3",
             外呼上面有目标最大数4 := "中间变量2"."3号梯外呼上面有目标最大数4",
             外呼上面有目标最大数5 := "中间变量2"."3号梯外呼上面有目标最大数5",
             外呼上面有目标最大数6 := "中间变量2"."3号梯外呼上面有目标最大数6",
             外呼上面有目标最大数7 := "中间变量2"."3号梯外呼上面有目标最大数7",
             外呼上面有目标最大数8 := "中间变量2"."3号梯外呼上面有目标最大数8",
             外呼上面有目标最大数9 := "中间变量2"."3号梯外呼上面有目标最大数9",
             外呼下面有目标最小数2 := "中间变量2"."3号梯外呼下面有目标最小数2",
             外呼下面有目标最小数3 := "中间变量2"."3号梯外呼下面有目标最小数3",
             外呼下面有目标最小数4 := "中间变量2"."3号梯外呼下面有目标最小数4",
             外呼下面有目标最小数5 := "中间变量2"."3号梯外呼下面有目标最小数5",
             外呼下面有目标最小数6 := "中间变量2"."3号梯外呼下面有目标最小数6",
             外呼下面有目标最小数7 := "中间变量2"."3号梯外呼下面有目标最小数7",
             外呼下面有目标最小数8 := "中间变量2"."3号梯外呼下面有目标最小数8",
             外呼下面有目标最小数9 := "中间变量2"."3号梯外呼下面有目标最小数9",
             外呼下面有目标最小数10 := "中间变量2"."3号梯外呼下面有目标最小数10",
             外呼下面有目标2 := "中间变量2"."3号梯外呼下面有目标2",
             外呼下面有目标3 := "中间变量2"."3号梯外呼下面有目标3",
             外呼下面有目标4 := "中间变量2"."3号梯外呼下面有目标4",
             外呼下面有目标5 := "中间变量2"."3号梯外呼下面有目标5",
             外呼下面有目标6 := "中间变量2"."3号梯外呼下面有目标6",
             外呼下面有目标7 := "中间变量2"."3号梯外呼下面有目标7",
             外呼下面有目标8 := "中间变量2"."3号梯外呼下面有目标8",
             外呼下面有目标9 := "中间变量2"."3号梯外呼下面有目标9",
             外呼下面有目标10 := "中间变量2"."3号梯外呼下面有目标10",
             外呼上面有目标1 := "中间变量2"."3号梯外呼上面有目标1",
             外呼上面有目标2 := "中间变量2"."3号梯外呼上面有目标2",
             外呼上面有目标3 := "中间变量2"."3号梯外呼上面有目标3",
             外呼上面有目标4 := "中间变量2"."3号梯外呼上面有目标4",
             外呼上面有目标5 := "中间变量2"."3号梯外呼上面有目标5",
             外呼上面有目标6 := "中间变量2"."3号梯外呼上面有目标6",
             外呼上面有目标7 := "中间变量2"."3号梯外呼上面有目标7",
             外呼上面有目标8 := "中间变量2"."3号梯外呼上面有目标8",
             外呼上面有目标9 := "中间变量2"."3号梯外呼上面有目标9",
             外呼下面无目标2 := "中间变量2"."3号梯外呼下面无目标2",
             外呼下面无目标3 := "中间变量2"."3号梯外呼下面无目标3",
             外呼下面无目标4 := "中间变量2"."3号梯外呼下面无目标4",
             外呼下面无目标5 := "中间变量2"."3号梯外呼下面无目标5",
             外呼下面无目标6 := "中间变量2"."3号梯外呼下面无目标6",
             外呼下面无目标7 := "中间变量2"."3号梯外呼下面无目标7",
             外呼下面无目标8 := "中间变量2"."3号梯外呼下面无目标8",
             外呼下面无目标9 := "中间变量2"."3号梯外呼下面无目标9",
             外呼上面无目标2 := "中间变量2"."3号梯外呼上面无目标2",
             外呼上面无目标3 := "中间变量2"."3号梯外呼上面无目标3",
             外呼上面无目标4 := "中间变量2"."3号梯外呼上面无目标4",
             外呼上面无目标5 := "中间变量2"."3号梯外呼上面无目标5",
             外呼上面无目标6 := "中间变量2"."3号梯外呼上面无目标6",
             外呼上面无目标7 := "中间变量2"."3号梯外呼上面无目标7",
             外呼上面无目标8 := "中间变量2"."3号梯外呼上面无目标8",
             外呼上面无目标9 := "中间变量2"."3号梯外呼上面无目标9",
             上行停站次数3 := "中间变量2"."3号梯上行停站次数3",
             上行停站次数4 := "中间变量2"."3号梯上行停站次数4",
             上行停站次数5 := "中间变量2"."3号梯上行停站次数5",
             上行停站次数6 := "中间变量2"."3号梯上行停站次数6",
             上行停站次数7 := "中间变量2"."3号梯上行停站次数7",
             上行停站次数8 := "中间变量2"."3号梯上行停站次数8",
             上行停站次数9 := "中间变量2"."3号梯上行停站次数9",
             下行停站次数2 := "中间变量2"."3号梯下行停站次数2",
             下行停站次数3 := "中间变量2"."3号梯下行停站次数3",
             下行停站次数4 := "中间变量2"."3号梯下行停站次数4",
             下行停站次数5 := "中间变量2"."3号梯下行停站次数5",
             下行停站次数6 := "中间变量2"."3号梯下行停站次数6",
             下行停站次数7 := "中间变量2"."3号梯下行停站次数7",
             下行停站次数8 := "中间变量2"."3号梯下行停站次数8",
             上行停站次数10 := "中间变量2"."3号梯上行停站次数10",
             下行停站次数1 := "中间变量2"."3号梯下行停站次数1",
             载重量 := "中间变量2"."3号梯转换后载重量",
             死机 := "中间变量1".死机3,
             限重分配 := "中间变量2".限重分配3,
             最终调度距离上1 => "中间变量2"."3梯1层最终调度距离",
             最终调度距离上2 => "中间变量2"."3梯2层最终调度距离上",
             最终调度距离上3 => "中间变量2"."3梯3层最终调度距离上",
             最终调度距离上4 => "中间变量2"."3梯4层最终调度距离上",
             最终调度距离上5 => "中间变量2"."3梯5层最终调度距离上",
             最终调度距离上6 => "中间变量2"."3梯6层最终调度距离上",
             最终调度距离上7 => "中间变量2"."3梯7层最终调度距离上",
             最终调度距离上8 => "中间变量2"."3梯8层最终调度距离上",
             最终调度距离上9 => "中间变量2"."3梯9层最终调度距离上",
             最终调度距离下2 => "中间变量2"."3梯2层最终调度距离下",
             最终调度距离下3 => "中间变量2"."3梯3层最终调度距离下",
             最终调度距离下4 => "中间变量2"."3梯4层最终调度距离下",
             最终调度距离下5 => "中间变量2"."3梯5层最终调度距离下",
             最终调度距离下6 => "中间变量2"."3梯6层最终调度距离下",
             最终调度距离下7 => "中间变量2"."3梯7层最终调度距离下",
             最终调度距离下8 => "中间变量2"."3梯8层最终调度距离下",
             最终调度距离下9 => "中间变量2"."3梯9层最终调度距离下",
             最终调度距离下10 => "中间变量2"."3梯10层最终调度距离");
END_REGION

REGION Network 5: 4号梯调度距离
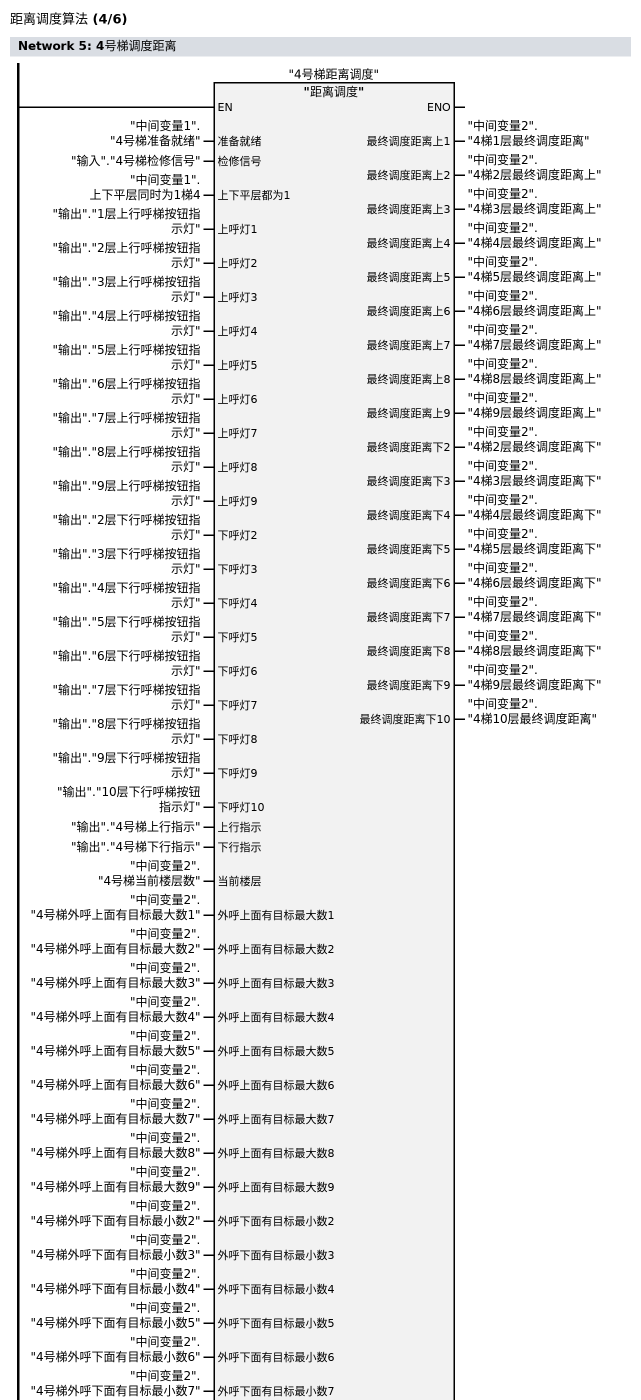
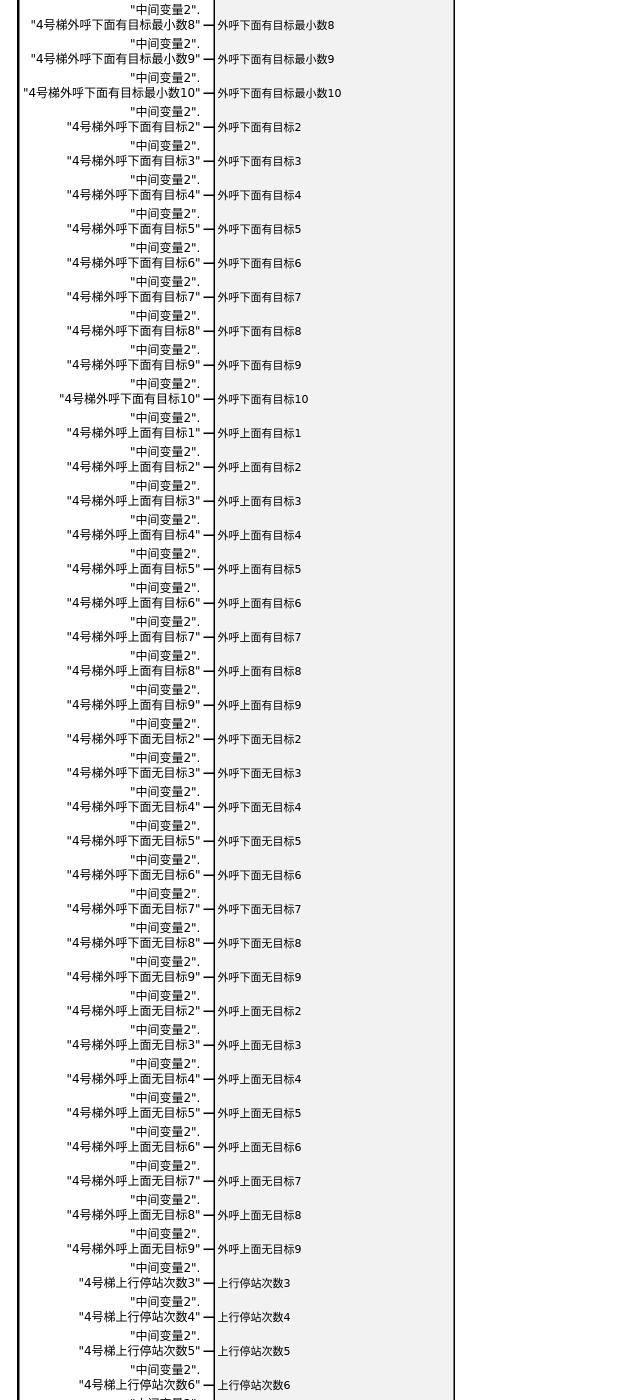
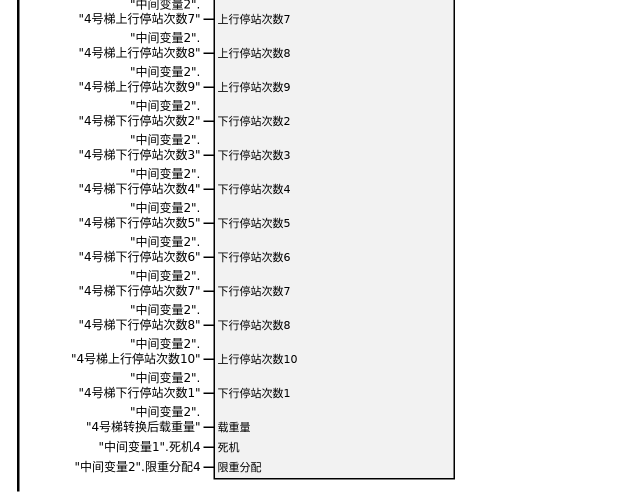
   RUNG wire#powerrail
      "4号梯距离调度"(准备就绪 := "中间变量1"."4号梯准备就绪", 检修信号 := "输入"."4号梯检修信号", 上下平层都为1 := "中间变量1".上下平层同时为1梯4, 上呼灯1 := "输出"."1层上行呼梯按钮指示灯", 上呼灯2 := "输出"."2层上行呼梯按钮指示灯", 上呼灯3 := "输出"."3层上行呼梯按钮指示灯", 上呼灯4 := "输出"."4层上行呼梯按钮指示灯", 上呼灯5 := "输出"."5层上行呼梯按钮指示灯", 上呼灯6 := "输出"."6层上行呼梯按钮指示灯", 上呼灯7 := "输出"."7层上行呼梯按钮指示灯", 上呼灯8 := "输出"."8层上行呼梯按钮指示灯", 上呼灯9 := "输出"."9层上行呼梯按钮指示灯", 下呼灯2 := "输出"."2层下行呼梯按钮指示灯", 下呼灯3 := "输出"."3层下行呼梯按钮指示灯", 下呼灯4 := "输出"."4层下行呼梯按钮指示灯", 下呼灯5 := "输出"."5层下行呼梯按钮指示灯", 下呼灯6 := "输出"."6层下行呼梯按钮指示灯", 下呼灯7 := "输出"."7层下行呼梯按钮指示灯", 下呼灯8 := "输出"."8层下行呼梯按钮指示灯", 下呼灯9 := "输出"."9层下行呼梯按钮指示灯", 下呼灯10 := "输出"."10层下行呼梯按钮指示灯", 上行指示 := "输出"."4号梯上行指示", 下行指示 := "输出"."4号梯下行指示", 当前楼层 := "中间变量2"."4号梯当前楼层数", 外呼上面有目标最大数1 := "中间变量2"."4号梯外呼上面有目标最大数1", 外呼上面有目标最大数2 := "中间变量2"."4号梯外呼上面有目标最大数2", 外呼上面有目标最大数3 := "中间变量2"."4号梯外呼上面有目标最大数3", 外呼上面有目标最大数4 := "中间变量2"."4号梯外呼上面有目标最大数4", 外呼上面有目标最大数5 := "中间变量2"."4号梯外呼上面有目标最大数5", 外呼上面有目标最大数6 := "中间变量2"."4号梯外呼上面有目标最大数6", 外呼上面有目标最大数7 := "中间变量2"."4号梯外呼上面有目标最大数7", 外呼上面有目标最大数8 := "中间变量2"."4号梯外呼上面有目标最大数8", 外呼上面有目标最大数9 := "中间变量2"."4号梯外呼上面有目标最大数9", 外呼下面有目标最小数2 := "中间变量2"."4号梯外呼下面有目标最小数2", 外呼下面有目标最小数3 := "中间变量2"."4号梯外呼下面有目标最小数3", 外呼下面有目标最小数4 := "中间变量2"."4号梯外呼下面有目标最小数4", 外呼下面有目标最小数5 := "中间变量2"."4号梯外呼下面有目标最小数5", 外呼下面有目标最小数6 := "中间变量2"."4号梯外呼下面有目标最小数6", 外呼下面有目标最小数7 := "中间变量2"."4号梯外呼下面有目标最小数7", 外呼下面有目标最小数8 := "中间变量2"."4号梯外呼下面有目标最小数8", 外呼下面有目标最小数9 := "中间变量2"."4号梯外呼下面有目标最小数9", 外呼下面有目标最小数10 := "中间变量2"."4号梯外呼下面有目标最小数10", 外呼下面有目标2 := "中间变量2"."4号梯外呼下面有目标2", 外呼下面有目标3 := "中间变量2"."4号梯外呼下面有目标3", 外呼下面有目标4 := "中间变量2"."4号梯外呼下面有目标4", 外呼下面有目标5 := "中间变量2"."4号梯外呼下面有目标5", 外呼下面有目标6 := "中间变量2"."4号梯外呼下面有目标6", 外呼下面有目标7 := "中间变量2"."4号梯外呼下面有目标7", 外呼下面有目标8 := "中间变量2"."4号梯外呼下面有目标8", 外呼下面有目标9 := "中间变量2"."4号梯外呼下面有目标9", 外呼下面有目标10 := "中间变量2"."4号梯外呼下面有目标10", 外呼上面有目标1 := "中间变量2"."4号梯外呼上面有目标1", 外呼上面有目标2 := "中间变量2"."4号梯外呼上面有目标2", 外呼上面有目标3 := "中间变量2"."4号梯外呼上面有目标3", 外呼上面有目标4 := "中间变量2"."4号梯外呼上面有目标4", 外呼上面有目标5 := "中间变量2"."4号梯外呼上面有目标5", 外呼上面有目标6 := "中间变量2"."4号梯外呼上面有目标6", 外呼上面有目标7 := "中间变量2"."4号梯外呼上面有目标7", 外呼上面有目标8 := "中间变量2"."4号梯外呼上面有目标8", 外呼上面有目标9 := "中间变量2"."4号梯外呼上面有目标9", 外呼下面无目标2 := "中间变量2"."4号梯外呼下面无目标2", 外呼下面无目标3 := "中间变量2"."4号梯外呼下面无目标3", 外呼下面无目标4 := "中间变量2"."4号梯外呼下面无目标4", 外呼下面无目标5 := "中间变量2"."4号梯外呼下面无目标5", 外呼下面无目标6 := "中间变量2"."4号梯外呼下面无目标6", 外呼下面无目标7 := "中间变量2"."4号梯外呼下面无目标7", 外呼下面无目标8 := "中间变量2"."4号梯外呼下面无目标8", 外呼下面无目标9 := "中间变量2"."4号梯外呼下面无目标9", 外呼上面无目标2 := "中间变量2"."4号梯外呼上面无目标2", 外呼上面无目标3 := "中间变量2"."4号梯外呼上面无目标3", 外呼上面无目标4 := "中间变量2"."4号梯外呼上面无目标4", 外呼上面无目标5 := "中间变量2"."4号梯外呼上面无目标5", 外呼上面无目标6 := "中间变量2"."4号梯外呼上面无目标6", 外呼上面无目标7 := "中间变量2"."4号梯外呼上面无目标7", 外呼上面无目标8 := "中间变量2"."4号梯外呼上面无目标8", 外呼上面无目标9 := "中间变量2"."4号梯外呼上面无目标9", 上行停站次数3 := "中间变量2"."4号梯上行停站次数3", 上行停站次数4 := "中间变量2"."4号梯上行停站次数4", 上行停站次数5 := "中间变量2"."4号梯上行停站次数5", 上行停站次数6 := "中间变量2"."4号梯上行停站次数6", 上行停站次数7 := "中间变量2"."4号梯上行停站次数7", 上行停站次数8 := "中间变量2"."4号梯上行停站次数8", 上行停站次数9 := "中间变量2"."4号梯上行停站次数9", 下行停站次数2 := "中间变量2"."4号梯下行停站次数2", 下行停站次数3 := "中间变量2"."4号梯下行停站次数3", 下行停站次数4 := "中间变量2"."4号梯下行停站次数4", 下行停站次数5 := "中间变量2"."4号梯下行停站次数5", 下行停站次数6 := "中间变量2"."4号梯下行停站次数6", 下行停站次数7 := "中间变量2"."4号梯下行停站次数7", 下行停站次数8 := "中间变量2"."4号梯下行停站次数8", 上行停站次数10 := "中间变量2"."4号梯上行停站次数10", 下行停站次数1 := "中间变量2"."4号梯下行停站次数1", 载重量 := "中间变量2"."4号梯转换后载重量", 死机 := "中间变量1".死机4, 限重分配 := "中间变量2".限重分配4, 最终调度距离上1 => "中间变量2"."4梯1层最终调度距离", 最终调度距离上2 => "中间变量2"."4梯2层最终调度距离上", 最终调度距离上3 => "中间变量2"."4梯3层最终调度距离上", 最终调度距离上4 => "中间变量2"."4梯4层最终调度距离上", 最终调度距离上5 => "中间变量2"."4梯5层最终调度距离上", 最终调度距离上6 => "中间变量2"."4梯6层最终调度距离上", 最终调度距离上7 => "中间变量2"."4梯7层最终调度距离上", 最终调度距离上8 => "中间变量2"."4梯8层最终调度距离上", 最终调度距离上9 => "中间变量2"."4梯9层最终调度距离上", 最终调度距离下2 => "中间变量2"."4梯2层最终调度距离下", 最终调度距离下3 => "中间变量2"."4梯3层最终调度距离下", 最终调度距离下4 => "中间变量2"."4梯4层最终调度距离下", 最终调度距离下5 => "中间变量2"."4梯5层最终调度距离下", 最终调度距离下6 => "中间变量2"."4梯6层最终调度距离下", 最终调度距离下7 => "中间变量2"."4梯7层最终调度距离下", 最终调度距离下8 => "中间变量2"."4梯8层最终调度距离下", 最终调度距离下9 => "中间变量2"."4梯9层最终调度距离下", 最终调度距离下10 => "中间变量2"."4梯10层最终调度距离")
   END_RUNG
   // the same network as SCL:
   "4号梯距离调度"(准备就绪 := "中间变量1"."4号梯准备就绪",   // "距离调度"
             检修信号 := "输入"."4号梯检修信号",
             上下平层都为1 := "中间变量1".上下平层同时为1梯4,
             上呼灯1 := "输出"."1层上行呼梯按钮指示灯",
             上呼灯2 := "输出"."2层上行呼梯按钮指示灯",
             上呼灯3 := "输出"."3层上行呼梯按钮指示灯",
             上呼灯4 := "输出"."4层上行呼梯按钮指示灯",
             上呼灯5 := "输出"."5层上行呼梯按钮指示灯",
             上呼灯6 := "输出"."6层上行呼梯按钮指示灯",
             上呼灯7 := "输出"."7层上行呼梯按钮指示灯",
             上呼灯8 := "输出"."8层上行呼梯按钮指示灯",
             上呼灯9 := "输出"."9层上行呼梯按钮指示灯",
             下呼灯2 := "输出"."2层下行呼梯按钮指示灯",
             下呼灯3 := "输出"."3层下行呼梯按钮指示灯",
             下呼灯4 := "输出"."4层下行呼梯按钮指示灯",
             下呼灯5 := "输出"."5层下行呼梯按钮指示灯",
             下呼灯6 := "输出"."6层下行呼梯按钮指示灯",
             下呼灯7 := "输出"."7层下行呼梯按钮指示灯",
             下呼灯8 := "输出"."8层下行呼梯按钮指示灯",
             下呼灯9 := "输出"."9层下行呼梯按钮指示灯",
             下呼灯10 := "输出"."10层下行呼梯按钮指示灯",
             上行指示 := "输出"."4号梯上行指示",
             下行指示 := "输出"."4号梯下行指示",
             当前楼层 := "中间变量2"."4号梯当前楼层数",
             外呼上面有目标最大数1 := "中间变量2"."4号梯外呼上面有目标最大数1",
             外呼上面有目标最大数2 := "中间变量2"."4号梯外呼上面有目标最大数2",
             外呼上面有目标最大数3 := "中间变量2"."4号梯外呼上面有目标最大数3",
             外呼上面有目标最大数4 := "中间变量2"."4号梯外呼上面有目标最大数4",
             外呼上面有目标最大数5 := "中间变量2"."4号梯外呼上面有目标最大数5",
             外呼上面有目标最大数6 := "中间变量2"."4号梯外呼上面有目标最大数6",
             外呼上面有目标最大数7 := "中间变量2"."4号梯外呼上面有目标最大数7",
             外呼上面有目标最大数8 := "中间变量2"."4号梯外呼上面有目标最大数8",
             外呼上面有目标最大数9 := "中间变量2"."4号梯外呼上面有目标最大数9",
             外呼下面有目标最小数2 := "中间变量2"."4号梯外呼下面有目标最小数2",
             外呼下面有目标最小数3 := "中间变量2"."4号梯外呼下面有目标最小数3",
             外呼下面有目标最小数4 := "中间变量2"."4号梯外呼下面有目标最小数4",
             外呼下面有目标最小数5 := "中间变量2"."4号梯外呼下面有目标最小数5",
             外呼下面有目标最小数6 := "中间变量2"."4号梯外呼下面有目标最小数6",
             外呼下面有目标最小数7 := "中间变量2"."4号梯外呼下面有目标最小数7",
             外呼下面有目标最小数8 := "中间变量2"."4号梯外呼下面有目标最小数8",
             外呼下面有目标最小数9 := "中间变量2"."4号梯外呼下面有目标最小数9",
             外呼下面有目标最小数10 := "中间变量2"."4号梯外呼下面有目标最小数10",
             外呼下面有目标2 := "中间变量2"."4号梯外呼下面有目标2",
             外呼下面有目标3 := "中间变量2"."4号梯外呼下面有目标3",
             外呼下面有目标4 := "中间变量2"."4号梯外呼下面有目标4",
             外呼下面有目标5 := "中间变量2"."4号梯外呼下面有目标5",
             外呼下面有目标6 := "中间变量2"."4号梯外呼下面有目标6",
             外呼下面有目标7 := "中间变量2"."4号梯外呼下面有目标7",
             外呼下面有目标8 := "中间变量2"."4号梯外呼下面有目标8",
             外呼下面有目标9 := "中间变量2"."4号梯外呼下面有目标9",
             外呼下面有目标10 := "中间变量2"."4号梯外呼下面有目标10",
             外呼上面有目标1 := "中间变量2"."4号梯外呼上面有目标1",
             外呼上面有目标2 := "中间变量2"."4号梯外呼上面有目标2",
             外呼上面有目标3 := "中间变量2"."4号梯外呼上面有目标3",
             外呼上面有目标4 := "中间变量2"."4号梯外呼上面有目标4",
             外呼上面有目标5 := "中间变量2"."4号梯外呼上面有目标5",
             外呼上面有目标6 := "中间变量2"."4号梯外呼上面有目标6",
             外呼上面有目标7 := "中间变量2"."4号梯外呼上面有目标7",
             外呼上面有目标8 := "中间变量2"."4号梯外呼上面有目标8",
             外呼上面有目标9 := "中间变量2"."4号梯外呼上面有目标9",
             外呼下面无目标2 := "中间变量2"."4号梯外呼下面无目标2",
             外呼下面无目标3 := "中间变量2"."4号梯外呼下面无目标3",
             外呼下面无目标4 := "中间变量2"."4号梯外呼下面无目标4",
             外呼下面无目标5 := "中间变量2"."4号梯外呼下面无目标5",
             外呼下面无目标6 := "中间变量2"."4号梯外呼下面无目标6",
             外呼下面无目标7 := "中间变量2"."4号梯外呼下面无目标7",
             外呼下面无目标8 := "中间变量2"."4号梯外呼下面无目标8",
             外呼下面无目标9 := "中间变量2"."4号梯外呼下面无目标9",
             外呼上面无目标2 := "中间变量2"."4号梯外呼上面无目标2",
             外呼上面无目标3 := "中间变量2"."4号梯外呼上面无目标3",
             外呼上面无目标4 := "中间变量2"."4号梯外呼上面无目标4",
             外呼上面无目标5 := "中间变量2"."4号梯外呼上面无目标5",
             外呼上面无目标6 := "中间变量2"."4号梯外呼上面无目标6",
             外呼上面无目标7 := "中间变量2"."4号梯外呼上面无目标7",
             外呼上面无目标8 := "中间变量2"."4号梯外呼上面无目标8",
             外呼上面无目标9 := "中间变量2"."4号梯外呼上面无目标9",
             上行停站次数3 := "中间变量2"."4号梯上行停站次数3",
             上行停站次数4 := "中间变量2"."4号梯上行停站次数4",
             上行停站次数5 := "中间变量2"."4号梯上行停站次数5",
             上行停站次数6 := "中间变量2"."4号梯上行停站次数6",
             上行停站次数7 := "中间变量2"."4号梯上行停站次数7",
             上行停站次数8 := "中间变量2"."4号梯上行停站次数8",
             上行停站次数9 := "中间变量2"."4号梯上行停站次数9",
             下行停站次数2 := "中间变量2"."4号梯下行停站次数2",
             下行停站次数3 := "中间变量2"."4号梯下行停站次数3",
             下行停站次数4 := "中间变量2"."4号梯下行停站次数4",
             下行停站次数5 := "中间变量2"."4号梯下行停站次数5",
             下行停站次数6 := "中间变量2"."4号梯下行停站次数6",
             下行停站次数7 := "中间变量2"."4号梯下行停站次数7",
             下行停站次数8 := "中间变量2"."4号梯下行停站次数8",
             上行停站次数10 := "中间变量2"."4号梯上行停站次数10",
             下行停站次数1 := "中间变量2"."4号梯下行停站次数1",
             载重量 := "中间变量2"."4号梯转换后载重量",
             死机 := "中间变量1".死机4,
             限重分配 := "中间变量2".限重分配4,
             最终调度距离上1 => "中间变量2"."4梯1层最终调度距离",
             最终调度距离上2 => "中间变量2"."4梯2层最终调度距离上",
             最终调度距离上3 => "中间变量2"."4梯3层最终调度距离上",
             最终调度距离上4 => "中间变量2"."4梯4层最终调度距离上",
             最终调度距离上5 => "中间变量2"."4梯5层最终调度距离上",
             最终调度距离上6 => "中间变量2"."4梯6层最终调度距离上",
             最终调度距离上7 => "中间变量2"."4梯7层最终调度距离上",
             最终调度距离上8 => "中间变量2"."4梯8层最终调度距离上",
             最终调度距离上9 => "中间变量2"."4梯9层最终调度距离上",
             最终调度距离下2 => "中间变量2"."4梯2层最终调度距离下",
             最终调度距离下3 => "中间变量2"."4梯3层最终调度距离下",
             最终调度距离下4 => "中间变量2"."4梯4层最终调度距离下",
             最终调度距离下5 => "中间变量2"."4梯5层最终调度距离下",
             最终调度距离下6 => "中间变量2"."4梯6层最终调度距离下",
             最终调度距离下7 => "中间变量2"."4梯7层最终调度距离下",
             最终调度距离下8 => "中间变量2"."4梯8层最终调度距离下",
             最终调度距离下9 => "中间变量2"."4梯9层最终调度距离下",
             最终调度距离下10 => "中间变量2"."4梯10层最终调度距离");
END_REGION

REGION Network 6: 5号梯调度距离
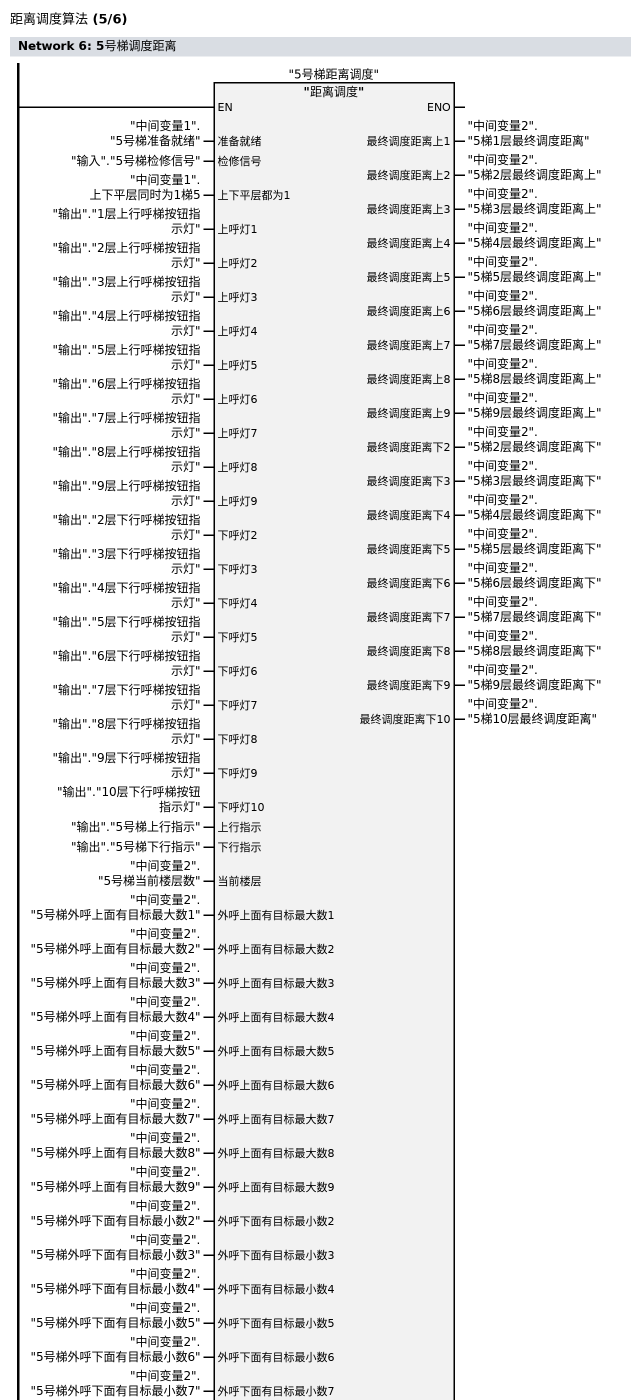
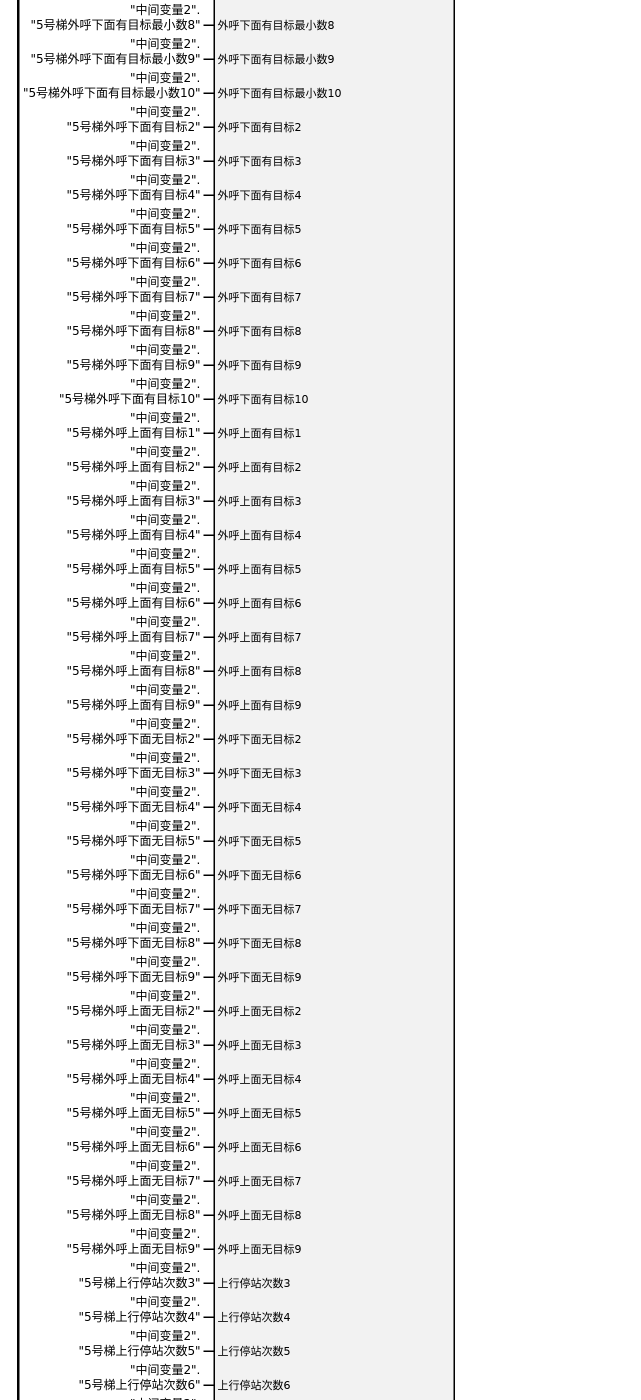
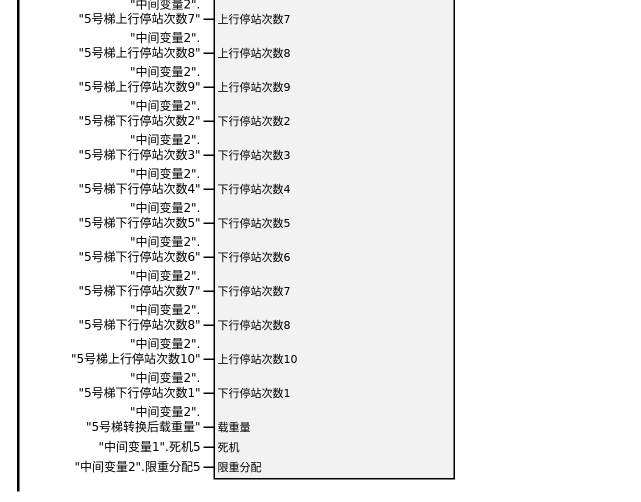
   RUNG wire#powerrail
      "5号梯距离调度"(准备就绪 := "中间变量1"."5号梯准备就绪", 检修信号 := "输入"."5号梯检修信号", 上下平层都为1 := "中间变量1".上下平层同时为1梯5, 上呼灯1 := "输出"."1层上行呼梯按钮指示灯", 上呼灯2 := "输出"."2层上行呼梯按钮指示灯", 上呼灯3 := "输出"."3层上行呼梯按钮指示灯", 上呼灯4 := "输出"."4层上行呼梯按钮指示灯", 上呼灯5 := "输出"."5层上行呼梯按钮指示灯", 上呼灯6 := "输出"."6层上行呼梯按钮指示灯", 上呼灯7 := "输出"."7层上行呼梯按钮指示灯", 上呼灯8 := "输出"."8层上行呼梯按钮指示灯", 上呼灯9 := "输出"."9层上行呼梯按钮指示灯", 下呼灯2 := "输出"."2层下行呼梯按钮指示灯", 下呼灯3 := "输出"."3层下行呼梯按钮指示灯", 下呼灯4 := "输出"."4层下行呼梯按钮指示灯", 下呼灯5 := "输出"."5层下行呼梯按钮指示灯", 下呼灯6 := "输出"."6层下行呼梯按钮指示灯", 下呼灯7 := "输出"."7层下行呼梯按钮指示灯", 下呼灯8 := "输出"."8层下行呼梯按钮指示灯", 下呼灯9 := "输出"."9层下行呼梯按钮指示灯", 下呼灯10 := "输出"."10层下行呼梯按钮指示灯", 上行指示 := "输出"."5号梯上行指示", 下行指示 := "输出"."5号梯下行指示", 当前楼层 := "中间变量2"."5号梯当前楼层数", 外呼上面有目标最大数1 := "中间变量2"."5号梯外呼上面有目标最大数1", 外呼上面有目标最大数2 := "中间变量2"."5号梯外呼上面有目标最大数2", 外呼上面有目标最大数3 := "中间变量2"."5号梯外呼上面有目标最大数3", 外呼上面有目标最大数4 := "中间变量2"."5号梯外呼上面有目标最大数4", 外呼上面有目标最大数5 := "中间变量2"."5号梯外呼上面有目标最大数5", 外呼上面有目标最大数6 := "中间变量2"."5号梯外呼上面有目标最大数6", 外呼上面有目标最大数7 := "中间变量2"."5号梯外呼上面有目标最大数7", 外呼上面有目标最大数8 := "中间变量2"."5号梯外呼上面有目标最大数8", 外呼上面有目标最大数9 := "中间变量2"."5号梯外呼上面有目标最大数9", 外呼下面有目标最小数2 := "中间变量2"."5号梯外呼下面有目标最小数2", 外呼下面有目标最小数3 := "中间变量2"."5号梯外呼下面有目标最小数3", 外呼下面有目标最小数4 := "中间变量2"."5号梯外呼下面有目标最小数4", 外呼下面有目标最小数5 := "中间变量2"."5号梯外呼下面有目标最小数5", 外呼下面有目标最小数6 := "中间变量2"."5号梯外呼下面有目标最小数6", 外呼下面有目标最小数7 := "中间变量2"."5号梯外呼下面有目标最小数7", 外呼下面有目标最小数8 := "中间变量2"."5号梯外呼下面有目标最小数8", 外呼下面有目标最小数9 := "中间变量2"."5号梯外呼下面有目标最小数9", 外呼下面有目标最小数10 := "中间变量2"."5号梯外呼下面有目标最小数10", 外呼下面有目标2 := "中间变量2"."5号梯外呼下面有目标2", 外呼下面有目标3 := "中间变量2"."5号梯外呼下面有目标3", 外呼下面有目标4 := "中间变量2"."5号梯外呼下面有目标4", 外呼下面有目标5 := "中间变量2"."5号梯外呼下面有目标5", 外呼下面有目标6 := "中间变量2"."5号梯外呼下面有目标6", 外呼下面有目标7 := "中间变量2"."5号梯外呼下面有目标7", 外呼下面有目标8 := "中间变量2"."5号梯外呼下面有目标8", 外呼下面有目标9 := "中间变量2"."5号梯外呼下面有目标9", 外呼下面有目标10 := "中间变量2"."5号梯外呼下面有目标10", 外呼上面有目标1 := "中间变量2"."5号梯外呼上面有目标1", 外呼上面有目标2 := "中间变量2"."5号梯外呼上面有目标2", 外呼上面有目标3 := "中间变量2"."5号梯外呼上面有目标3", 外呼上面有目标4 := "中间变量2"."5号梯外呼上面有目标4", 外呼上面有目标5 := "中间变量2"."5号梯外呼上面有目标5", 外呼上面有目标6 := "中间变量2"."5号梯外呼上面有目标6", 外呼上面有目标7 := "中间变量2"."5号梯外呼上面有目标7", 外呼上面有目标8 := "中间变量2"."5号梯外呼上面有目标8", 外呼上面有目标9 := "中间变量2"."5号梯外呼上面有目标9", 外呼下面无目标2 := "中间变量2"."5号梯外呼下面无目标2", 外呼下面无目标3 := "中间变量2"."5号梯外呼下面无目标3", 外呼下面无目标4 := "中间变量2"."5号梯外呼下面无目标4", 外呼下面无目标5 := "中间变量2"."5号梯外呼下面无目标5", 外呼下面无目标6 := "中间变量2"."5号梯外呼下面无目标6", 外呼下面无目标7 := "中间变量2"."5号梯外呼下面无目标7", 外呼下面无目标8 := "中间变量2"."5号梯外呼下面无目标8", 外呼下面无目标9 := "中间变量2"."5号梯外呼下面无目标9", 外呼上面无目标2 := "中间变量2"."5号梯外呼上面无目标2", 外呼上面无目标3 := "中间变量2"."5号梯外呼上面无目标3", 外呼上面无目标4 := "中间变量2"."5号梯外呼上面无目标4", 外呼上面无目标5 := "中间变量2"."5号梯外呼上面无目标5", 外呼上面无目标6 := "中间变量2"."5号梯外呼上面无目标6", 外呼上面无目标7 := "中间变量2"."5号梯外呼上面无目标7", 外呼上面无目标8 := "中间变量2"."5号梯外呼上面无目标8", 外呼上面无目标9 := "中间变量2"."5号梯外呼上面无目标9", 上行停站次数3 := "中间变量2"."5号梯上行停站次数3", 上行停站次数4 := "中间变量2"."5号梯上行停站次数4", 上行停站次数5 := "中间变量2"."5号梯上行停站次数5", 上行停站次数6 := "中间变量2"."5号梯上行停站次数6", 上行停站次数7 := "中间变量2"."5号梯上行停站次数7", 上行停站次数8 := "中间变量2"."5号梯上行停站次数8", 上行停站次数9 := "中间变量2"."5号梯上行停站次数9", 下行停站次数2 := "中间变量2"."5号梯下行停站次数2", 下行停站次数3 := "中间变量2"."5号梯下行停站次数3", 下行停站次数4 := "中间变量2"."5号梯下行停站次数4", 下行停站次数5 := "中间变量2"."5号梯下行停站次数5", 下行停站次数6 := "中间变量2"."5号梯下行停站次数6", 下行停站次数7 := "中间变量2"."5号梯下行停站次数7", 下行停站次数8 := "中间变量2"."5号梯下行停站次数8", 上行停站次数10 := "中间变量2"."5号梯上行停站次数10", 下行停站次数1 := "中间变量2"."5号梯下行停站次数1", 载重量 := "中间变量2"."5号梯转换后载重量", 死机 := "中间变量1".死机5, 限重分配 := "中间变量2".限重分配5, 最终调度距离上1 => "中间变量2"."5梯1层最终调度距离", 最终调度距离上2 => "中间变量2"."5梯2层最终调度距离上", 最终调度距离上3 => "中间变量2"."5梯3层最终调度距离上", 最终调度距离上4 => "中间变量2"."5梯4层最终调度距离上", 最终调度距离上5 => "中间变量2"."5梯5层最终调度距离上", 最终调度距离上6 => "中间变量2"."5梯6层最终调度距离上", 最终调度距离上7 => "中间变量2"."5梯7层最终调度距离上", 最终调度距离上8 => "中间变量2"."5梯8层最终调度距离上", 最终调度距离上9 => "中间变量2"."5梯9层最终调度距离上", 最终调度距离下2 => "中间变量2"."5梯2层最终调度距离下", 最终调度距离下3 => "中间变量2"."5梯3层最终调度距离下", 最终调度距离下4 => "中间变量2"."5梯4层最终调度距离下", 最终调度距离下5 => "中间变量2"."5梯5层最终调度距离下", 最终调度距离下6 => "中间变量2"."5梯6层最终调度距离下", 最终调度距离下7 => "中间变量2"."5梯7层最终调度距离下", 最终调度距离下8 => "中间变量2"."5梯8层最终调度距离下", 最终调度距离下9 => "中间变量2"."5梯9层最终调度距离下", 最终调度距离下10 => "中间变量2"."5梯10层最终调度距离")
   END_RUNG
   // the same network as SCL:
   "5号梯距离调度"(准备就绪 := "中间变量1"."5号梯准备就绪",   // "距离调度"
             检修信号 := "输入"."5号梯检修信号",
             上下平层都为1 := "中间变量1".上下平层同时为1梯5,
             上呼灯1 := "输出"."1层上行呼梯按钮指示灯",
             上呼灯2 := "输出"."2层上行呼梯按钮指示灯",
             上呼灯3 := "输出"."3层上行呼梯按钮指示灯",
             上呼灯4 := "输出"."4层上行呼梯按钮指示灯",
             上呼灯5 := "输出"."5层上行呼梯按钮指示灯",
             上呼灯6 := "输出"."6层上行呼梯按钮指示灯",
             上呼灯7 := "输出"."7层上行呼梯按钮指示灯",
             上呼灯8 := "输出"."8层上行呼梯按钮指示灯",
             上呼灯9 := "输出"."9层上行呼梯按钮指示灯",
             下呼灯2 := "输出"."2层下行呼梯按钮指示灯",
             下呼灯3 := "输出"."3层下行呼梯按钮指示灯",
             下呼灯4 := "输出"."4层下行呼梯按钮指示灯",
             下呼灯5 := "输出"."5层下行呼梯按钮指示灯",
             下呼灯6 := "输出"."6层下行呼梯按钮指示灯",
             下呼灯7 := "输出"."7层下行呼梯按钮指示灯",
             下呼灯8 := "输出"."8层下行呼梯按钮指示灯",
             下呼灯9 := "输出"."9层下行呼梯按钮指示灯",
             下呼灯10 := "输出"."10层下行呼梯按钮指示灯",
             上行指示 := "输出"."5号梯上行指示",
             下行指示 := "输出"."5号梯下行指示",
             当前楼层 := "中间变量2"."5号梯当前楼层数",
             外呼上面有目标最大数1 := "中间变量2"."5号梯外呼上面有目标最大数1",
             外呼上面有目标最大数2 := "中间变量2"."5号梯外呼上面有目标最大数2",
             外呼上面有目标最大数3 := "中间变量2"."5号梯外呼上面有目标最大数3",
             外呼上面有目标最大数4 := "中间变量2"."5号梯外呼上面有目标最大数4",
             外呼上面有目标最大数5 := "中间变量2"."5号梯外呼上面有目标最大数5",
             外呼上面有目标最大数6 := "中间变量2"."5号梯外呼上面有目标最大数6",
             外呼上面有目标最大数7 := "中间变量2"."5号梯外呼上面有目标最大数7",
             外呼上面有目标最大数8 := "中间变量2"."5号梯外呼上面有目标最大数8",
             外呼上面有目标最大数9 := "中间变量2"."5号梯外呼上面有目标最大数9",
             外呼下面有目标最小数2 := "中间变量2"."5号梯外呼下面有目标最小数2",
             外呼下面有目标最小数3 := "中间变量2"."5号梯外呼下面有目标最小数3",
             外呼下面有目标最小数4 := "中间变量2"."5号梯外呼下面有目标最小数4",
             外呼下面有目标最小数5 := "中间变量2"."5号梯外呼下面有目标最小数5",
             外呼下面有目标最小数6 := "中间变量2"."5号梯外呼下面有目标最小数6",
             外呼下面有目标最小数7 := "中间变量2"."5号梯外呼下面有目标最小数7",
             外呼下面有目标最小数8 := "中间变量2"."5号梯外呼下面有目标最小数8",
             外呼下面有目标最小数9 := "中间变量2"."5号梯外呼下面有目标最小数9",
             外呼下面有目标最小数10 := "中间变量2"."5号梯外呼下面有目标最小数10",
             外呼下面有目标2 := "中间变量2"."5号梯外呼下面有目标2",
             外呼下面有目标3 := "中间变量2"."5号梯外呼下面有目标3",
             外呼下面有目标4 := "中间变量2"."5号梯外呼下面有目标4",
             外呼下面有目标5 := "中间变量2"."5号梯外呼下面有目标5",
             外呼下面有目标6 := "中间变量2"."5号梯外呼下面有目标6",
             外呼下面有目标7 := "中间变量2"."5号梯外呼下面有目标7",
             外呼下面有目标8 := "中间变量2"."5号梯外呼下面有目标8",
             外呼下面有目标9 := "中间变量2"."5号梯外呼下面有目标9",
             外呼下面有目标10 := "中间变量2"."5号梯外呼下面有目标10",
             外呼上面有目标1 := "中间变量2"."5号梯外呼上面有目标1",
             外呼上面有目标2 := "中间变量2"."5号梯外呼上面有目标2",
             外呼上面有目标3 := "中间变量2"."5号梯外呼上面有目标3",
             外呼上面有目标4 := "中间变量2"."5号梯外呼上面有目标4",
             外呼上面有目标5 := "中间变量2"."5号梯外呼上面有目标5",
             外呼上面有目标6 := "中间变量2"."5号梯外呼上面有目标6",
             外呼上面有目标7 := "中间变量2"."5号梯外呼上面有目标7",
             外呼上面有目标8 := "中间变量2"."5号梯外呼上面有目标8",
             外呼上面有目标9 := "中间变量2"."5号梯外呼上面有目标9",
             外呼下面无目标2 := "中间变量2"."5号梯外呼下面无目标2",
             外呼下面无目标3 := "中间变量2"."5号梯外呼下面无目标3",
             外呼下面无目标4 := "中间变量2"."5号梯外呼下面无目标4",
             外呼下面无目标5 := "中间变量2"."5号梯外呼下面无目标5",
             外呼下面无目标6 := "中间变量2"."5号梯外呼下面无目标6",
             外呼下面无目标7 := "中间变量2"."5号梯外呼下面无目标7",
             外呼下面无目标8 := "中间变量2"."5号梯外呼下面无目标8",
             外呼下面无目标9 := "中间变量2"."5号梯外呼下面无目标9",
             外呼上面无目标2 := "中间变量2"."5号梯外呼上面无目标2",
             外呼上面无目标3 := "中间变量2"."5号梯外呼上面无目标3",
             外呼上面无目标4 := "中间变量2"."5号梯外呼上面无目标4",
             外呼上面无目标5 := "中间变量2"."5号梯外呼上面无目标5",
             外呼上面无目标6 := "中间变量2"."5号梯外呼上面无目标6",
             外呼上面无目标7 := "中间变量2"."5号梯外呼上面无目标7",
             外呼上面无目标8 := "中间变量2"."5号梯外呼上面无目标8",
             外呼上面无目标9 := "中间变量2"."5号梯外呼上面无目标9",
             上行停站次数3 := "中间变量2"."5号梯上行停站次数3",
             上行停站次数4 := "中间变量2"."5号梯上行停站次数4",
             上行停站次数5 := "中间变量2"."5号梯上行停站次数5",
             上行停站次数6 := "中间变量2"."5号梯上行停站次数6",
             上行停站次数7 := "中间变量2"."5号梯上行停站次数7",
             上行停站次数8 := "中间变量2"."5号梯上行停站次数8",
             上行停站次数9 := "中间变量2"."5号梯上行停站次数9",
             下行停站次数2 := "中间变量2"."5号梯下行停站次数2",
             下行停站次数3 := "中间变量2"."5号梯下行停站次数3",
             下行停站次数4 := "中间变量2"."5号梯下行停站次数4",
             下行停站次数5 := "中间变量2"."5号梯下行停站次数5",
             下行停站次数6 := "中间变量2"."5号梯下行停站次数6",
             下行停站次数7 := "中间变量2"."5号梯下行停站次数7",
             下行停站次数8 := "中间变量2"."5号梯下行停站次数8",
             上行停站次数10 := "中间变量2"."5号梯上行停站次数10",
             下行停站次数1 := "中间变量2"."5号梯下行停站次数1",
             载重量 := "中间变量2"."5号梯转换后载重量",
             死机 := "中间变量1".死机5,
             限重分配 := "中间变量2".限重分配5,
             最终调度距离上1 => "中间变量2"."5梯1层最终调度距离",
             最终调度距离上2 => "中间变量2"."5梯2层最终调度距离上",
             最终调度距离上3 => "中间变量2"."5梯3层最终调度距离上",
             最终调度距离上4 => "中间变量2"."5梯4层最终调度距离上",
             最终调度距离上5 => "中间变量2"."5梯5层最终调度距离上",
             最终调度距离上6 => "中间变量2"."5梯6层最终调度距离上",
             最终调度距离上7 => "中间变量2"."5梯7层最终调度距离上",
             最终调度距离上8 => "中间变量2"."5梯8层最终调度距离上",
             最终调度距离上9 => "中间变量2"."5梯9层最终调度距离上",
             最终调度距离下2 => "中间变量2"."5梯2层最终调度距离下",
             最终调度距离下3 => "中间变量2"."5梯3层最终调度距离下",
             最终调度距离下4 => "中间变量2"."5梯4层最终调度距离下",
             最终调度距离下5 => "中间变量2"."5梯5层最终调度距离下",
             最终调度距离下6 => "中间变量2"."5梯6层最终调度距离下",
             最终调度距离下7 => "中间变量2"."5梯7层最终调度距离下",
             最终调度距离下8 => "中间变量2"."5梯8层最终调度距离下",
             最终调度距离下9 => "中间变量2"."5梯9层最终调度距离下",
             最终调度距离下10 => "中间变量2"."5梯10层最终调度距离");
END_REGION

REGION Network 7: 6号梯调度距离
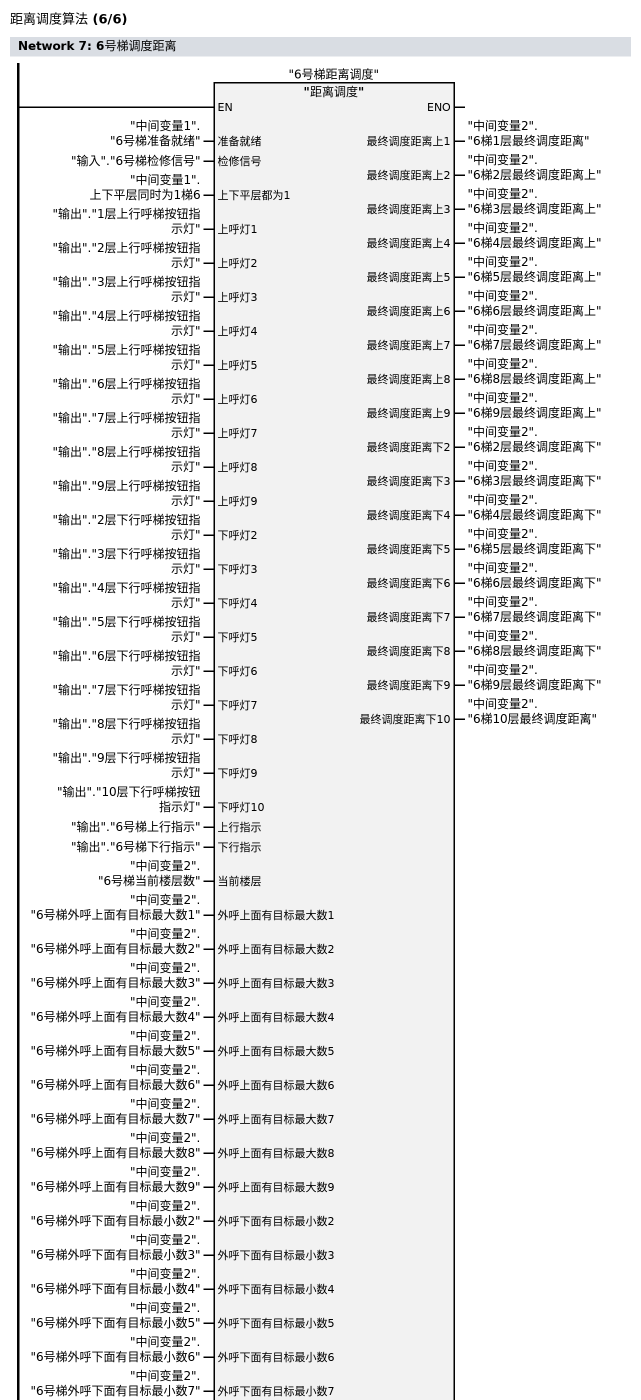
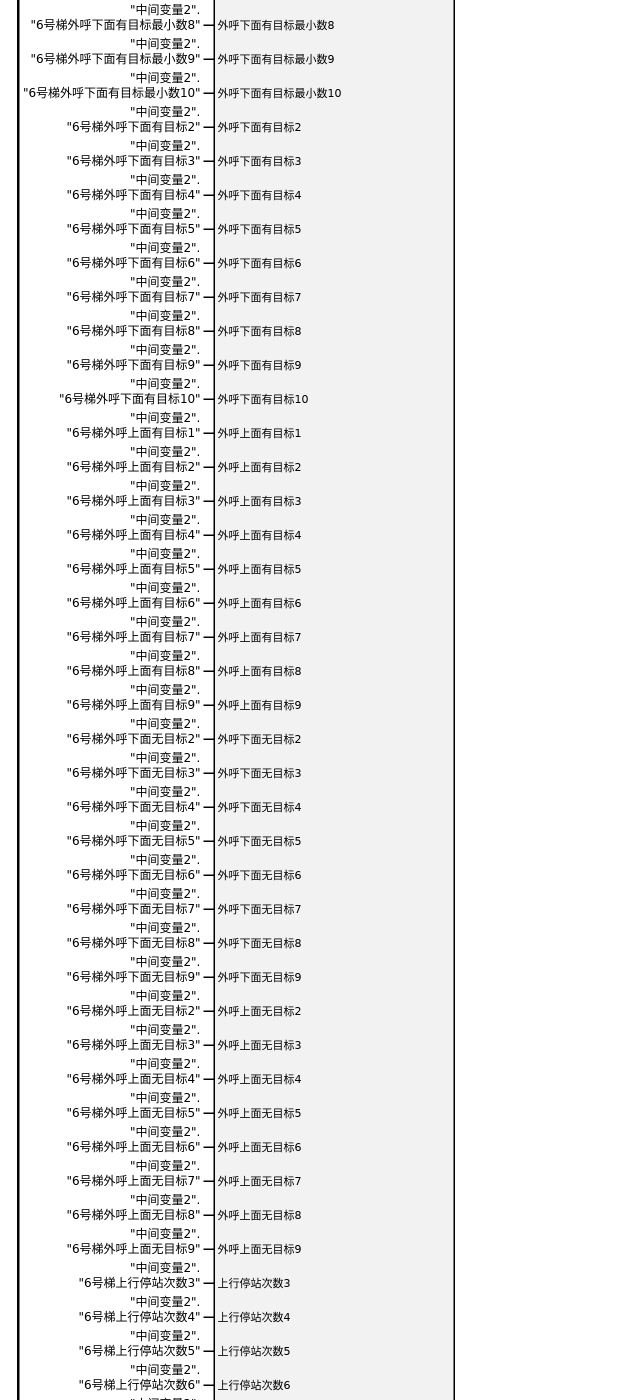
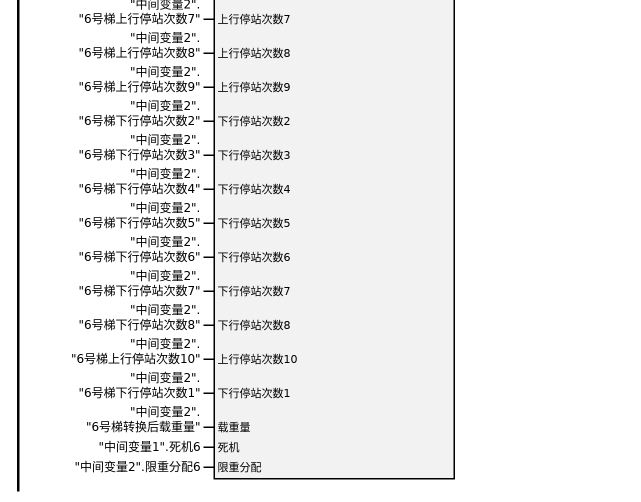
   RUNG wire#powerrail
      "6号梯距离调度"(准备就绪 := "中间变量1"."6号梯准备就绪", 检修信号 := "输入"."6号梯检修信号", 上下平层都为1 := "中间变量1".上下平层同时为1梯6, 上呼灯1 := "输出"."1层上行呼梯按钮指示灯", 上呼灯2 := "输出"."2层上行呼梯按钮指示灯", 上呼灯3 := "输出"."3层上行呼梯按钮指示灯", 上呼灯4 := "输出"."4层上行呼梯按钮指示灯", 上呼灯5 := "输出"."5层上行呼梯按钮指示灯", 上呼灯6 := "输出"."6层上行呼梯按钮指示灯", 上呼灯7 := "输出"."7层上行呼梯按钮指示灯", 上呼灯8 := "输出"."8层上行呼梯按钮指示灯", 上呼灯9 := "输出"."9层上行呼梯按钮指示灯", 下呼灯2 := "输出"."2层下行呼梯按钮指示灯", 下呼灯3 := "输出"."3层下行呼梯按钮指示灯", 下呼灯4 := "输出"."4层下行呼梯按钮指示灯", 下呼灯5 := "输出"."5层下行呼梯按钮指示灯", 下呼灯6 := "输出"."6层下行呼梯按钮指示灯", 下呼灯7 := "输出"."7层下行呼梯按钮指示灯", 下呼灯8 := "输出"."8层下行呼梯按钮指示灯", 下呼灯9 := "输出"."9层下行呼梯按钮指示灯", 下呼灯10 := "输出"."10层下行呼梯按钮指示灯", 上行指示 := "输出"."6号梯上行指示", 下行指示 := "输出"."6号梯下行指示", 当前楼层 := "中间变量2"."6号梯当前楼层数", 外呼上面有目标最大数1 := "中间变量2"."6号梯外呼上面有目标最大数1", 外呼上面有目标最大数2 := "中间变量2"."6号梯外呼上面有目标最大数2", 外呼上面有目标最大数3 := "中间变量2"."6号梯外呼上面有目标最大数3", 外呼上面有目标最大数4 := "中间变量2"."6号梯外呼上面有目标最大数4", 外呼上面有目标最大数5 := "中间变量2"."6号梯外呼上面有目标最大数5", 外呼上面有目标最大数6 := "中间变量2"."6号梯外呼上面有目标最大数6", 外呼上面有目标最大数7 := "中间变量2"."6号梯外呼上面有目标最大数7", 外呼上面有目标最大数8 := "中间变量2"."6号梯外呼上面有目标最大数8", 外呼上面有目标最大数9 := "中间变量2"."6号梯外呼上面有目标最大数9", 外呼下面有目标最小数2 := "中间变量2"."6号梯外呼下面有目标最小数2", 外呼下面有目标最小数3 := "中间变量2"."6号梯外呼下面有目标最小数3", 外呼下面有目标最小数4 := "中间变量2"."6号梯外呼下面有目标最小数4", 外呼下面有目标最小数5 := "中间变量2"."6号梯外呼下面有目标最小数5", 外呼下面有目标最小数6 := "中间变量2"."6号梯外呼下面有目标最小数6", 外呼下面有目标最小数7 := "中间变量2"."6号梯外呼下面有目标最小数7", 外呼下面有目标最小数8 := "中间变量2"."6号梯外呼下面有目标最小数8", 外呼下面有目标最小数9 := "中间变量2"."6号梯外呼下面有目标最小数9", 外呼下面有目标最小数10 := "中间变量2"."6号梯外呼下面有目标最小数10", 外呼下面有目标2 := "中间变量2"."6号梯外呼下面有目标2", 外呼下面有目标3 := "中间变量2"."6号梯外呼下面有目标3", 外呼下面有目标4 := "中间变量2"."6号梯外呼下面有目标4", 外呼下面有目标5 := "中间变量2"."6号梯外呼下面有目标5", 外呼下面有目标6 := "中间变量2"."6号梯外呼下面有目标6", 外呼下面有目标7 := "中间变量2"."6号梯外呼下面有目标7", 外呼下面有目标8 := "中间变量2"."6号梯外呼下面有目标8", 外呼下面有目标9 := "中间变量2"."6号梯外呼下面有目标9", 外呼下面有目标10 := "中间变量2"."6号梯外呼下面有目标10", 外呼上面有目标1 := "中间变量2"."6号梯外呼上面有目标1", 外呼上面有目标2 := "中间变量2"."6号梯外呼上面有目标2", 外呼上面有目标3 := "中间变量2"."6号梯外呼上面有目标3", 外呼上面有目标4 := "中间变量2"."6号梯外呼上面有目标4", 外呼上面有目标5 := "中间变量2"."6号梯外呼上面有目标5", 外呼上面有目标6 := "中间变量2"."6号梯外呼上面有目标6", 外呼上面有目标7 := "中间变量2"."6号梯外呼上面有目标7", 外呼上面有目标8 := "中间变量2"."6号梯外呼上面有目标8", 外呼上面有目标9 := "中间变量2"."6号梯外呼上面有目标9", 外呼下面无目标2 := "中间变量2"."6号梯外呼下面无目标2", 外呼下面无目标3 := "中间变量2"."6号梯外呼下面无目标3", 外呼下面无目标4 := "中间变量2"."6号梯外呼下面无目标4", 外呼下面无目标5 := "中间变量2"."6号梯外呼下面无目标5", 外呼下面无目标6 := "中间变量2"."6号梯外呼下面无目标6", 外呼下面无目标7 := "中间变量2"."6号梯外呼下面无目标7", 外呼下面无目标8 := "中间变量2"."6号梯外呼下面无目标8", 外呼下面无目标9 := "中间变量2"."6号梯外呼下面无目标9", 外呼上面无目标2 := "中间变量2"."6号梯外呼上面无目标2", 外呼上面无目标3 := "中间变量2"."6号梯外呼上面无目标3", 外呼上面无目标4 := "中间变量2"."6号梯外呼上面无目标4", 外呼上面无目标5 := "中间变量2"."6号梯外呼上面无目标5", 外呼上面无目标6 := "中间变量2"."6号梯外呼上面无目标6", 外呼上面无目标7 := "中间变量2"."6号梯外呼上面无目标7", 外呼上面无目标8 := "中间变量2"."6号梯外呼上面无目标8", 外呼上面无目标9 := "中间变量2"."6号梯外呼上面无目标9", 上行停站次数3 := "中间变量2"."6号梯上行停站次数3", 上行停站次数4 := "中间变量2"."6号梯上行停站次数4", 上行停站次数5 := "中间变量2"."6号梯上行停站次数5", 上行停站次数6 := "中间变量2"."6号梯上行停站次数6", 上行停站次数7 := "中间变量2"."6号梯上行停站次数7", 上行停站次数8 := "中间变量2"."6号梯上行停站次数8", 上行停站次数9 := "中间变量2"."6号梯上行停站次数9", 下行停站次数2 := "中间变量2"."6号梯下行停站次数2", 下行停站次数3 := "中间变量2"."6号梯下行停站次数3", 下行停站次数4 := "中间变量2"."6号梯下行停站次数4", 下行停站次数5 := "中间变量2"."6号梯下行停站次数5", 下行停站次数6 := "中间变量2"."6号梯下行停站次数6", 下行停站次数7 := "中间变量2"."6号梯下行停站次数7", 下行停站次数8 := "中间变量2"."6号梯下行停站次数8", 上行停站次数10 := "中间变量2"."6号梯上行停站次数10", 下行停站次数1 := "中间变量2"."6号梯下行停站次数1", 载重量 := "中间变量2"."6号梯转换后载重量", 死机 := "中间变量1".死机6, 限重分配 := "中间变量2".限重分配6, 最终调度距离上1 => "中间变量2"."6梯1层最终调度距离", 最终调度距离上2 => "中间变量2"."6梯2层最终调度距离上", 最终调度距离上3 => "中间变量2"."6梯3层最终调度距离上", 最终调度距离上4 => "中间变量2"."6梯4层最终调度距离上", 最终调度距离上5 => "中间变量2"."6梯5层最终调度距离上", 最终调度距离上6 => "中间变量2"."6梯6层最终调度距离上", 最终调度距离上7 => "中间变量2"."6梯7层最终调度距离上", 最终调度距离上8 => "中间变量2"."6梯8层最终调度距离上", 最终调度距离上9 => "中间变量2"."6梯9层最终调度距离上", 最终调度距离下2 => "中间变量2"."6梯2层最终调度距离下", 最终调度距离下3 => "中间变量2"."6梯3层最终调度距离下", 最终调度距离下4 => "中间变量2"."6梯4层最终调度距离下", 最终调度距离下5 => "中间变量2"."6梯5层最终调度距离下", 最终调度距离下6 => "中间变量2"."6梯6层最终调度距离下", 最终调度距离下7 => "中间变量2"."6梯7层最终调度距离下", 最终调度距离下8 => "中间变量2"."6梯8层最终调度距离下", 最终调度距离下9 => "中间变量2"."6梯9层最终调度距离下", 最终调度距离下10 => "中间变量2"."6梯10层最终调度距离")
   END_RUNG
   // the same network as SCL:
   "6号梯距离调度"(准备就绪 := "中间变量1"."6号梯准备就绪",   // "距离调度"
             检修信号 := "输入"."6号梯检修信号",
             上下平层都为1 := "中间变量1".上下平层同时为1梯6,
             上呼灯1 := "输出"."1层上行呼梯按钮指示灯",
             上呼灯2 := "输出"."2层上行呼梯按钮指示灯",
             上呼灯3 := "输出"."3层上行呼梯按钮指示灯",
             上呼灯4 := "输出"."4层上行呼梯按钮指示灯",
             上呼灯5 := "输出"."5层上行呼梯按钮指示灯",
             上呼灯6 := "输出"."6层上行呼梯按钮指示灯",
             上呼灯7 := "输出"."7层上行呼梯按钮指示灯",
             上呼灯8 := "输出"."8层上行呼梯按钮指示灯",
             上呼灯9 := "输出"."9层上行呼梯按钮指示灯",
             下呼灯2 := "输出"."2层下行呼梯按钮指示灯",
             下呼灯3 := "输出"."3层下行呼梯按钮指示灯",
             下呼灯4 := "输出"."4层下行呼梯按钮指示灯",
             下呼灯5 := "输出"."5层下行呼梯按钮指示灯",
             下呼灯6 := "输出"."6层下行呼梯按钮指示灯",
             下呼灯7 := "输出"."7层下行呼梯按钮指示灯",
             下呼灯8 := "输出"."8层下行呼梯按钮指示灯",
             下呼灯9 := "输出"."9层下行呼梯按钮指示灯",
             下呼灯10 := "输出"."10层下行呼梯按钮指示灯",
             上行指示 := "输出"."6号梯上行指示",
             下行指示 := "输出"."6号梯下行指示",
             当前楼层 := "中间变量2"."6号梯当前楼层数",
             外呼上面有目标最大数1 := "中间变量2"."6号梯外呼上面有目标最大数1",
             外呼上面有目标最大数2 := "中间变量2"."6号梯外呼上面有目标最大数2",
             外呼上面有目标最大数3 := "中间变量2"."6号梯外呼上面有目标最大数3",
             外呼上面有目标最大数4 := "中间变量2"."6号梯外呼上面有目标最大数4",
             外呼上面有目标最大数5 := "中间变量2"."6号梯外呼上面有目标最大数5",
             外呼上面有目标最大数6 := "中间变量2"."6号梯外呼上面有目标最大数6",
             外呼上面有目标最大数7 := "中间变量2"."6号梯外呼上面有目标最大数7",
             外呼上面有目标最大数8 := "中间变量2"."6号梯外呼上面有目标最大数8",
             外呼上面有目标最大数9 := "中间变量2"."6号梯外呼上面有目标最大数9",
             外呼下面有目标最小数2 := "中间变量2"."6号梯外呼下面有目标最小数2",
             外呼下面有目标最小数3 := "中间变量2"."6号梯外呼下面有目标最小数3",
             外呼下面有目标最小数4 := "中间变量2"."6号梯外呼下面有目标最小数4",
             外呼下面有目标最小数5 := "中间变量2"."6号梯外呼下面有目标最小数5",
             外呼下面有目标最小数6 := "中间变量2"."6号梯外呼下面有目标最小数6",
             外呼下面有目标最小数7 := "中间变量2"."6号梯外呼下面有目标最小数7",
             外呼下面有目标最小数8 := "中间变量2"."6号梯外呼下面有目标最小数8",
             外呼下面有目标最小数9 := "中间变量2"."6号梯外呼下面有目标最小数9",
             外呼下面有目标最小数10 := "中间变量2"."6号梯外呼下面有目标最小数10",
             外呼下面有目标2 := "中间变量2"."6号梯外呼下面有目标2",
             外呼下面有目标3 := "中间变量2"."6号梯外呼下面有目标3",
             外呼下面有目标4 := "中间变量2"."6号梯外呼下面有目标4",
             外呼下面有目标5 := "中间变量2"."6号梯外呼下面有目标5",
             外呼下面有目标6 := "中间变量2"."6号梯外呼下面有目标6",
             外呼下面有目标7 := "中间变量2"."6号梯外呼下面有目标7",
             外呼下面有目标8 := "中间变量2"."6号梯外呼下面有目标8",
             外呼下面有目标9 := "中间变量2"."6号梯外呼下面有目标9",
             外呼下面有目标10 := "中间变量2"."6号梯外呼下面有目标10",
             外呼上面有目标1 := "中间变量2"."6号梯外呼上面有目标1",
             外呼上面有目标2 := "中间变量2"."6号梯外呼上面有目标2",
             外呼上面有目标3 := "中间变量2"."6号梯外呼上面有目标3",
             外呼上面有目标4 := "中间变量2"."6号梯外呼上面有目标4",
             外呼上面有目标5 := "中间变量2"."6号梯外呼上面有目标5",
             外呼上面有目标6 := "中间变量2"."6号梯外呼上面有目标6",
             外呼上面有目标7 := "中间变量2"."6号梯外呼上面有目标7",
             外呼上面有目标8 := "中间变量2"."6号梯外呼上面有目标8",
             外呼上面有目标9 := "中间变量2"."6号梯外呼上面有目标9",
             外呼下面无目标2 := "中间变量2"."6号梯外呼下面无目标2",
             外呼下面无目标3 := "中间变量2"."6号梯外呼下面无目标3",
             外呼下面无目标4 := "中间变量2"."6号梯外呼下面无目标4",
             外呼下面无目标5 := "中间变量2"."6号梯外呼下面无目标5",
             外呼下面无目标6 := "中间变量2"."6号梯外呼下面无目标6",
             外呼下面无目标7 := "中间变量2"."6号梯外呼下面无目标7",
             外呼下面无目标8 := "中间变量2"."6号梯外呼下面无目标8",
             外呼下面无目标9 := "中间变量2"."6号梯外呼下面无目标9",
             外呼上面无目标2 := "中间变量2"."6号梯外呼上面无目标2",
             外呼上面无目标3 := "中间变量2"."6号梯外呼上面无目标3",
             外呼上面无目标4 := "中间变量2"."6号梯外呼上面无目标4",
             外呼上面无目标5 := "中间变量2"."6号梯外呼上面无目标5",
             外呼上面无目标6 := "中间变量2"."6号梯外呼上面无目标6",
             外呼上面无目标7 := "中间变量2"."6号梯外呼上面无目标7",
             外呼上面无目标8 := "中间变量2"."6号梯外呼上面无目标8",
             外呼上面无目标9 := "中间变量2"."6号梯外呼上面无目标9",
             上行停站次数3 := "中间变量2"."6号梯上行停站次数3",
             上行停站次数4 := "中间变量2"."6号梯上行停站次数4",
             上行停站次数5 := "中间变量2"."6号梯上行停站次数5",
             上行停站次数6 := "中间变量2"."6号梯上行停站次数6",
             上行停站次数7 := "中间变量2"."6号梯上行停站次数7",
             上行停站次数8 := "中间变量2"."6号梯上行停站次数8",
             上行停站次数9 := "中间变量2"."6号梯上行停站次数9",
             下行停站次数2 := "中间变量2"."6号梯下行停站次数2",
             下行停站次数3 := "中间变量2"."6号梯下行停站次数3",
             下行停站次数4 := "中间变量2"."6号梯下行停站次数4",
             下行停站次数5 := "中间变量2"."6号梯下行停站次数5",
             下行停站次数6 := "中间变量2"."6号梯下行停站次数6",
             下行停站次数7 := "中间变量2"."6号梯下行停站次数7",
             下行停站次数8 := "中间变量2"."6号梯下行停站次数8",
             上行停站次数10 := "中间变量2"."6号梯上行停站次数10",
             下行停站次数1 := "中间变量2"."6号梯下行停站次数1",
             载重量 := "中间变量2"."6号梯转换后载重量",
             死机 := "中间变量1".死机6,
             限重分配 := "中间变量2".限重分配6,
             最终调度距离上1 => "中间变量2"."6梯1层最终调度距离",
             最终调度距离上2 => "中间变量2"."6梯2层最终调度距离上",
             最终调度距离上3 => "中间变量2"."6梯3层最终调度距离上",
             最终调度距离上4 => "中间变量2"."6梯4层最终调度距离上",
             最终调度距离上5 => "中间变量2"."6梯5层最终调度距离上",
             最终调度距离上6 => "中间变量2"."6梯6层最终调度距离上",
             最终调度距离上7 => "中间变量2"."6梯7层最终调度距离上",
             最终调度距离上8 => "中间变量2"."6梯8层最终调度距离上",
             最终调度距离上9 => "中间变量2"."6梯9层最终调度距离上",
             最终调度距离下2 => "中间变量2"."6梯2层最终调度距离下",
             最终调度距离下3 => "中间变量2"."6梯3层最终调度距离下",
             最终调度距离下4 => "中间变量2"."6梯4层最终调度距离下",
             最终调度距离下5 => "中间变量2"."6梯5层最终调度距离下",
             最终调度距离下6 => "中间变量2"."6梯6层最终调度距离下",
             最终调度距离下7 => "中间变量2"."6梯7层最终调度距离下",
             最终调度距离下8 => "中间变量2"."6梯8层最终调度距离下",
             最终调度距离下9 => "中间变量2"."6梯9层最终调度距离下",
             最终调度距离下10 => "中间变量2"."6梯10层最终调度距离");
END_REGION
END_FUNCTION

FUNCTION "载重量转换" : Void   // FC6, LAD
{ S7_Optimized_Access := 'TRUE' }
VERSION : 0.1
BEGIN

REGION Network 2: 电梯载重量转换
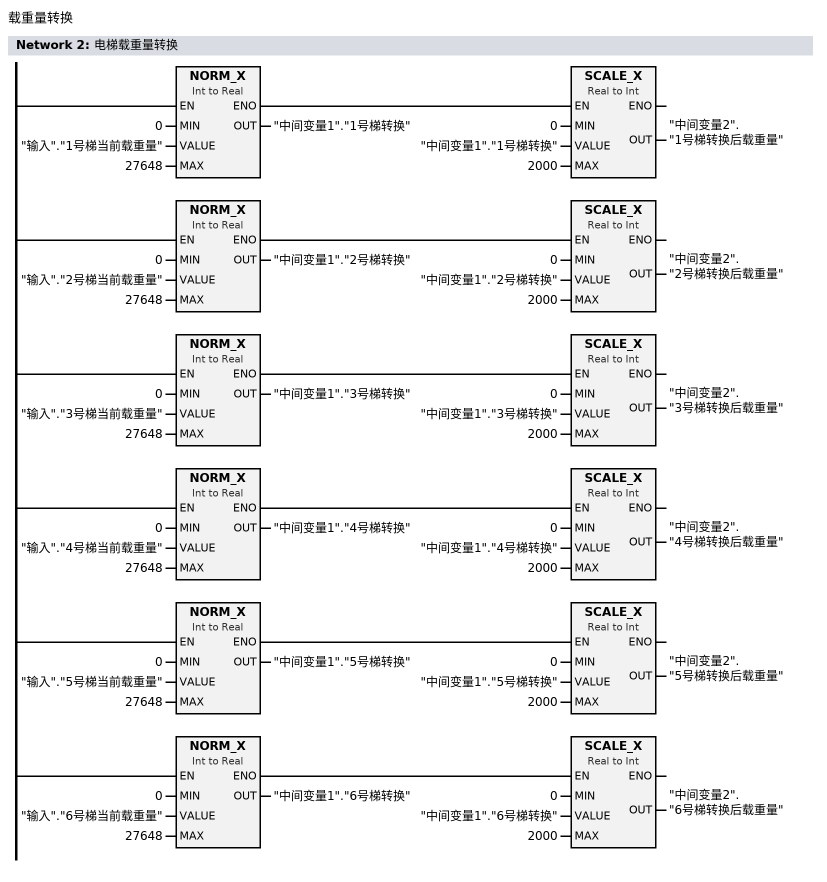
   RUNG wire#powerrail
      { S7_Templates := "[SrcType := Int, DestType := Real]" } Normalize(min := 0, value := "输入"."1号梯当前载重量", max := 27648, out => "中间变量1"."1号梯转换")
      { S7_Templates := "[SrcType := Real, DestType := Int]" } Scale(min := 0, value := "中间变量1"."1号梯转换", max := 2000, out => "中间变量2"."1号梯转换后载重量")
   END_RUNG
   RUNG wire#powerrail
      { S7_Templates := "[SrcType := Int, DestType := Real]" } Normalize(min := 0, value := "输入"."2号梯当前载重量", max := 27648, out => "中间变量1"."2号梯转换")
      { S7_Templates := "[SrcType := Real, DestType := Int]" } Scale(min := 0, value := "中间变量1"."2号梯转换", max := 2000, out => "中间变量2"."2号梯转换后载重量")
   END_RUNG
   RUNG wire#powerrail
      { S7_Templates := "[SrcType := Int, DestType := Real]" } Normalize(min := 0, value := "输入"."3号梯当前载重量", max := 27648, out => "中间变量1"."3号梯转换")
      { S7_Templates := "[SrcType := Real, DestType := Int]" } Scale(min := 0, value := "中间变量1"."3号梯转换", max := 2000, out => "中间变量2"."3号梯转换后载重量")
   END_RUNG
   RUNG wire#powerrail
      { S7_Templates := "[SrcType := Int, DestType := Real]" } Normalize(min := 0, value := "输入"."4号梯当前载重量", max := 27648, out => "中间变量1"."4号梯转换")
      { S7_Templates := "[SrcType := Real, DestType := Int]" } Scale(min := 0, value := "中间变量1"."4号梯转换", max := 2000, out => "中间变量2"."4号梯转换后载重量")
   END_RUNG
   RUNG wire#powerrail
      { S7_Templates := "[SrcType := Int, DestType := Real]" } Normalize(min := 0, value := "输入"."5号梯当前载重量", max := 27648, out => "中间变量1"."5号梯转换")
      { S7_Templates := "[SrcType := Real, DestType := Int]" } Scale(min := 0, value := "中间变量1"."5号梯转换", max := 2000, out => "中间变量2"."5号梯转换后载重量")
   END_RUNG
   RUNG wire#powerrail
      { S7_Templates := "[SrcType := Int, DestType := Real]" } Normalize(min := 0, value := "输入"."6号梯当前载重量", max := 27648, out => "中间变量1"."6号梯转换")
      { S7_Templates := "[SrcType := Real, DestType := Int]" } Scale(min := 0, value := "中间变量1"."6号梯转换", max := 2000, out => "中间变量2"."6号梯转换后载重量")
   END_RUNG
   // the same network as SCL:
   "中间变量1"."1号梯转换" := NORM_X(MIN := 0, VALUE := "输入"."1号梯当前载重量", MAX := 27648);
   "中间变量2"."1号梯转换后载重量" := SCALE_X(MIN := 0, VALUE := "中间变量1"."1号梯转换", MAX := 2000);
   "中间变量1"."2号梯转换" := NORM_X(MIN := 0, VALUE := "输入"."2号梯当前载重量", MAX := 27648);
   "中间变量2"."2号梯转换后载重量" := SCALE_X(MIN := 0, VALUE := "中间变量1"."2号梯转换", MAX := 2000);
   "中间变量1"."3号梯转换" := NORM_X(MIN := 0, VALUE := "输入"."3号梯当前载重量", MAX := 27648);
   "中间变量2"."3号梯转换后载重量" := SCALE_X(MIN := 0, VALUE := "中间变量1"."3号梯转换", MAX := 2000);
   "中间变量1"."4号梯转换" := NORM_X(MIN := 0, VALUE := "输入"."4号梯当前载重量", MAX := 27648);
   "中间变量2"."4号梯转换后载重量" := SCALE_X(MIN := 0, VALUE := "中间变量1"."4号梯转换", MAX := 2000);
   "中间变量1"."5号梯转换" := NORM_X(MIN := 0, VALUE := "输入"."5号梯当前载重量", MAX := 27648);
   "中间变量2"."5号梯转换后载重量" := SCALE_X(MIN := 0, VALUE := "中间变量1"."5号梯转换", MAX := 2000);
   "中间变量1"."6号梯转换" := NORM_X(MIN := 0, VALUE := "输入"."6号梯当前载重量", MAX := 27648);
   "中间变量2"."6号梯转换后载重量" := SCALE_X(MIN := 0, VALUE := "中间变量1"."6号梯转换", MAX := 2000);
END_REGION
END_FUNCTION

FUNCTION "停层次数计算" : Void   // FC7, LAD
{ S7_Optimized_Access := 'TRUE' }
VERSION : 0.1
BEGIN

REGION Network 2: 1号梯
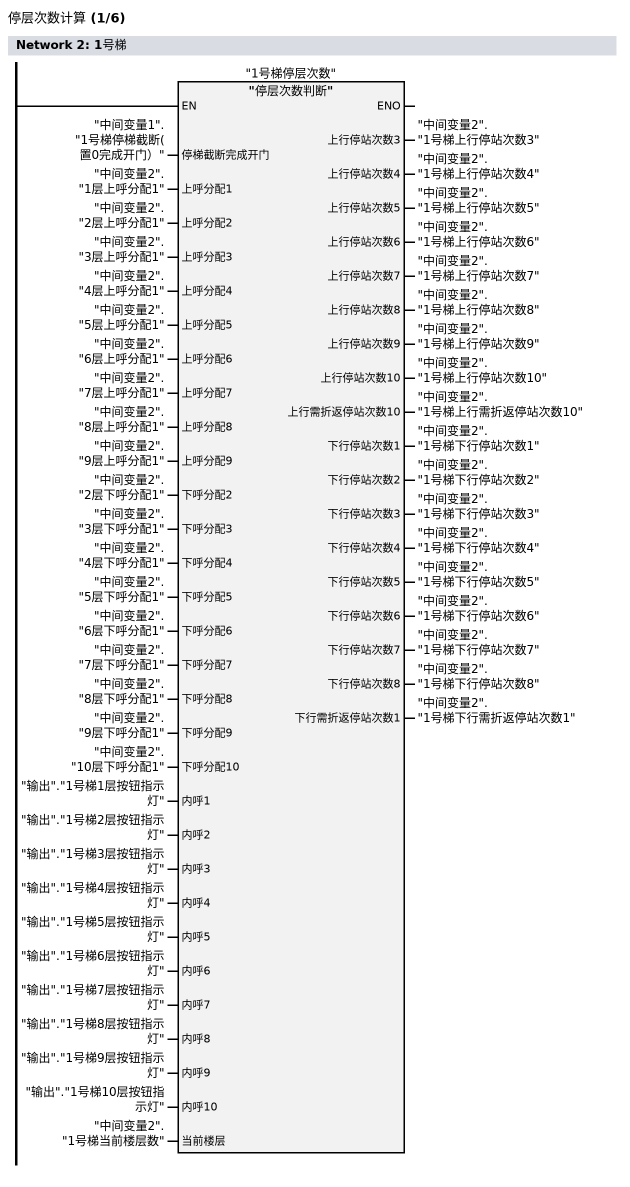
   RUNG wire#powerrail
      "1号梯停层次数"(停梯截断完成开门 := "中间变量1"."1号梯停梯截断(置0完成开门）", 上呼分配1 := "中间变量2"."1层上呼分配1", 上呼分配2 := "中间变量2"."2层上呼分配1", 上呼分配3 := "中间变量2"."3层上呼分配1", 上呼分配4 := "中间变量2"."4层上呼分配1", 上呼分配5 := "中间变量2"."5层上呼分配1", 上呼分配6 := "中间变量2"."6层上呼分配1", 上呼分配7 := "中间变量2"."7层上呼分配1", 上呼分配8 := "中间变量2"."8层上呼分配1", 上呼分配9 := "中间变量2"."9层上呼分配1", 下呼分配2 := "中间变量2"."2层下呼分配1", 下呼分配3 := "中间变量2"."3层下呼分配1", 下呼分配4 := "中间变量2"."4层下呼分配1", 下呼分配5 := "中间变量2"."5层下呼分配1", 下呼分配6 := "中间变量2"."6层下呼分配1", 下呼分配7 := "中间变量2"."7层下呼分配1", 下呼分配8 := "中间变量2"."8层下呼分配1", 下呼分配9 := "中间变量2"."9层下呼分配1", 下呼分配10 := "中间变量2"."10层下呼分配1", 内呼1 := "输出"."1号梯1层按钮指示灯", 内呼2 := "输出"."1号梯2层按钮指示灯", 内呼3 := "输出"."1号梯3层按钮指示灯", 内呼4 := "输出"."1号梯4层按钮指示灯", 内呼5 := "输出"."1号梯5层按钮指示灯", 内呼6 := "输出"."1号梯6层按钮指示灯", 内呼7 := "输出"."1号梯7层按钮指示灯", 内呼8 := "输出"."1号梯8层按钮指示灯", 内呼9 := "输出"."1号梯9层按钮指示灯", 内呼10 := "输出"."1号梯10层按钮指示灯", 当前楼层 := "中间变量2"."1号梯当前楼层数", 上行停站次数3 => "中间变量2"."1号梯上行停站次数3", 上行停站次数4 => "中间变量2"."1号梯上行停站次数4", 上行停站次数5 => "中间变量2"."1号梯上行停站次数5", 上行停站次数6 => "中间变量2"."1号梯上行停站次数6", 上行停站次数7 => "中间变量2"."1号梯上行停站次数7", 上行停站次数8 => "中间变量2"."1号梯上行停站次数8", 上行停站次数9 => "中间变量2"."1号梯上行停站次数9", 上行停站次数10 => "中间变量2"."1号梯上行停站次数10", 上行需折返停站次数10 => "中间变量2"."1号梯上行需折返停站次数10", 下行停站次数1 => "中间变量2"."1号梯下行停站次数1", 下行停站次数2 => "中间变量2"."1号梯下行停站次数2", 下行停站次数3 => "中间变量2"."1号梯下行停站次数3", 下行停站次数4 => "中间变量2"."1号梯下行停站次数4", 下行停站次数5 => "中间变量2"."1号梯下行停站次数5", 下行停站次数6 => "中间变量2"."1号梯下行停站次数6", 下行停站次数7 => "中间变量2"."1号梯下行停站次数7", 下行停站次数8 => "中间变量2"."1号梯下行停站次数8", 下行需折返停站次数1 => "中间变量2"."1号梯下行需折返停站次数1")
   END_RUNG
   // the same network as SCL:
   "1号梯停层次数"(停梯截断完成开门 := "中间变量1"."1号梯停梯截断(置0完成开门）",   // "停层次数判断"
             上呼分配1 := "中间变量2"."1层上呼分配1",
             上呼分配2 := "中间变量2"."2层上呼分配1",
             上呼分配3 := "中间变量2"."3层上呼分配1",
             上呼分配4 := "中间变量2"."4层上呼分配1",
             上呼分配5 := "中间变量2"."5层上呼分配1",
             上呼分配6 := "中间变量2"."6层上呼分配1",
             上呼分配7 := "中间变量2"."7层上呼分配1",
             上呼分配8 := "中间变量2"."8层上呼分配1",
             上呼分配9 := "中间变量2"."9层上呼分配1",
             下呼分配2 := "中间变量2"."2层下呼分配1",
             下呼分配3 := "中间变量2"."3层下呼分配1",
             下呼分配4 := "中间变量2"."4层下呼分配1",
             下呼分配5 := "中间变量2"."5层下呼分配1",
             下呼分配6 := "中间变量2"."6层下呼分配1",
             下呼分配7 := "中间变量2"."7层下呼分配1",
             下呼分配8 := "中间变量2"."8层下呼分配1",
             下呼分配9 := "中间变量2"."9层下呼分配1",
             下呼分配10 := "中间变量2"."10层下呼分配1",
             内呼1 := "输出"."1号梯1层按钮指示灯",
             内呼2 := "输出"."1号梯2层按钮指示灯",
             内呼3 := "输出"."1号梯3层按钮指示灯",
             内呼4 := "输出"."1号梯4层按钮指示灯",
             内呼5 := "输出"."1号梯5层按钮指示灯",
             内呼6 := "输出"."1号梯6层按钮指示灯",
             内呼7 := "输出"."1号梯7层按钮指示灯",
             内呼8 := "输出"."1号梯8层按钮指示灯",
             内呼9 := "输出"."1号梯9层按钮指示灯",
             内呼10 := "输出"."1号梯10层按钮指示灯",
             当前楼层 := "中间变量2"."1号梯当前楼层数",
             上行停站次数3 => "中间变量2"."1号梯上行停站次数3",
             上行停站次数4 => "中间变量2"."1号梯上行停站次数4",
             上行停站次数5 => "中间变量2"."1号梯上行停站次数5",
             上行停站次数6 => "中间变量2"."1号梯上行停站次数6",
             上行停站次数7 => "中间变量2"."1号梯上行停站次数7",
             上行停站次数8 => "中间变量2"."1号梯上行停站次数8",
             上行停站次数9 => "中间变量2"."1号梯上行停站次数9",
             上行停站次数10 => "中间变量2"."1号梯上行停站次数10",
             上行需折返停站次数10 => "中间变量2"."1号梯上行需折返停站次数10",
             下行停站次数1 => "中间变量2"."1号梯下行停站次数1",
             下行停站次数2 => "中间变量2"."1号梯下行停站次数2",
             下行停站次数3 => "中间变量2"."1号梯下行停站次数3",
             下行停站次数4 => "中间变量2"."1号梯下行停站次数4",
             下行停站次数5 => "中间变量2"."1号梯下行停站次数5",
             下行停站次数6 => "中间变量2"."1号梯下行停站次数6",
             下行停站次数7 => "中间变量2"."1号梯下行停站次数7",
             下行停站次数8 => "中间变量2"."1号梯下行停站次数8",
             下行需折返停站次数1 => "中间变量2"."1号梯下行需折返停站次数1");
END_REGION

REGION Network 3: 2号梯
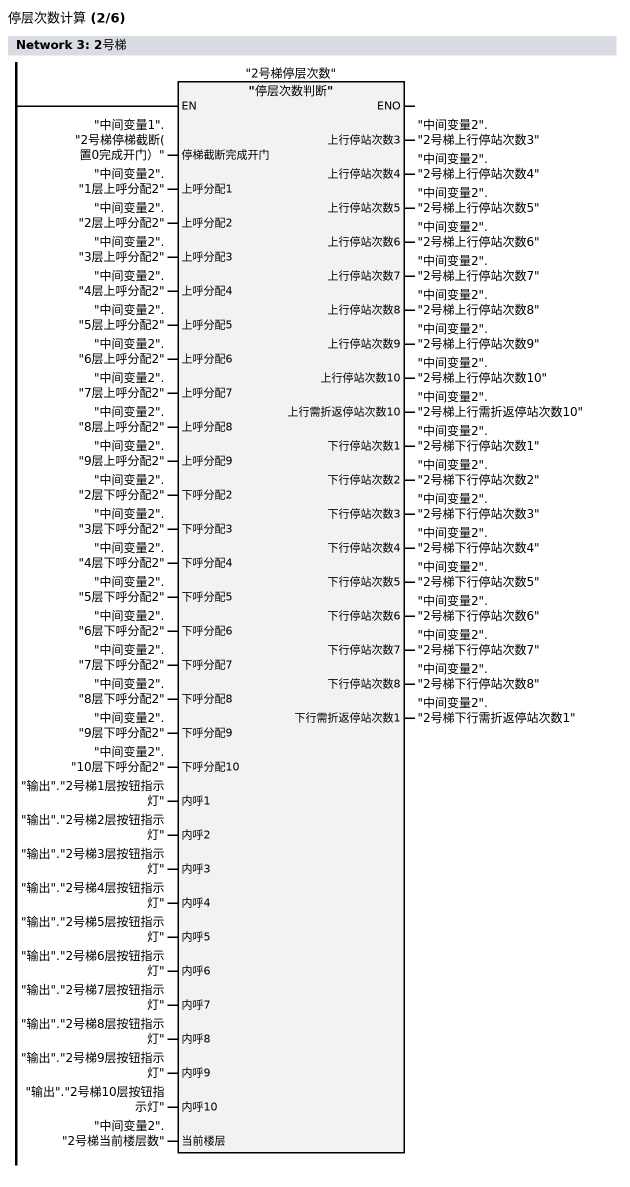
   RUNG wire#powerrail
      "2号梯停层次数"(停梯截断完成开门 := "中间变量1"."2号梯停梯截断(置0完成开门）", 上呼分配1 := "中间变量2"."1层上呼分配2", 上呼分配2 := "中间变量2"."2层上呼分配2", 上呼分配3 := "中间变量2"."3层上呼分配2", 上呼分配4 := "中间变量2"."4层上呼分配2", 上呼分配5 := "中间变量2"."5层上呼分配2", 上呼分配6 := "中间变量2"."6层上呼分配2", 上呼分配7 := "中间变量2"."7层上呼分配2", 上呼分配8 := "中间变量2"."8层上呼分配2", 上呼分配9 := "中间变量2"."9层上呼分配2", 下呼分配2 := "中间变量2"."2层下呼分配2", 下呼分配3 := "中间变量2"."3层下呼分配2", 下呼分配4 := "中间变量2"."4层下呼分配2", 下呼分配5 := "中间变量2"."5层下呼分配2", 下呼分配6 := "中间变量2"."6层下呼分配2", 下呼分配7 := "中间变量2"."7层下呼分配2", 下呼分配8 := "中间变量2"."8层下呼分配2", 下呼分配9 := "中间变量2"."9层下呼分配2", 下呼分配10 := "中间变量2"."10层下呼分配2", 内呼1 := "输出"."2号梯1层按钮指示灯", 内呼2 := "输出"."2号梯2层按钮指示灯", 内呼3 := "输出"."2号梯3层按钮指示灯", 内呼4 := "输出"."2号梯4层按钮指示灯", 内呼5 := "输出"."2号梯5层按钮指示灯", 内呼6 := "输出"."2号梯6层按钮指示灯", 内呼7 := "输出"."2号梯7层按钮指示灯", 内呼8 := "输出"."2号梯8层按钮指示灯", 内呼9 := "输出"."2号梯9层按钮指示灯", 内呼10 := "输出"."2号梯10层按钮指示灯", 当前楼层 := "中间变量2"."2号梯当前楼层数", 上行停站次数3 => "中间变量2"."2号梯上行停站次数3", 上行停站次数4 => "中间变量2"."2号梯上行停站次数4", 上行停站次数5 => "中间变量2"."2号梯上行停站次数5", 上行停站次数6 => "中间变量2"."2号梯上行停站次数6", 上行停站次数7 => "中间变量2"."2号梯上行停站次数7", 上行停站次数8 => "中间变量2"."2号梯上行停站次数8", 上行停站次数9 => "中间变量2"."2号梯上行停站次数9", 上行停站次数10 => "中间变量2"."2号梯上行停站次数10", 上行需折返停站次数10 => "中间变量2"."2号梯上行需折返停站次数10", 下行停站次数1 => "中间变量2"."2号梯下行停站次数1", 下行停站次数2 => "中间变量2"."2号梯下行停站次数2", 下行停站次数3 => "中间变量2"."2号梯下行停站次数3", 下行停站次数4 => "中间变量2"."2号梯下行停站次数4", 下行停站次数5 => "中间变量2"."2号梯下行停站次数5", 下行停站次数6 => "中间变量2"."2号梯下行停站次数6", 下行停站次数7 => "中间变量2"."2号梯下行停站次数7", 下行停站次数8 => "中间变量2"."2号梯下行停站次数8", 下行需折返停站次数1 => "中间变量2"."2号梯下行需折返停站次数1")
   END_RUNG
   // the same network as SCL:
   "2号梯停层次数"(停梯截断完成开门 := "中间变量1"."2号梯停梯截断(置0完成开门）",   // "停层次数判断"
             上呼分配1 := "中间变量2"."1层上呼分配2",
             上呼分配2 := "中间变量2"."2层上呼分配2",
             上呼分配3 := "中间变量2"."3层上呼分配2",
             上呼分配4 := "中间变量2"."4层上呼分配2",
             上呼分配5 := "中间变量2"."5层上呼分配2",
             上呼分配6 := "中间变量2"."6层上呼分配2",
             上呼分配7 := "中间变量2"."7层上呼分配2",
             上呼分配8 := "中间变量2"."8层上呼分配2",
             上呼分配9 := "中间变量2"."9层上呼分配2",
             下呼分配2 := "中间变量2"."2层下呼分配2",
             下呼分配3 := "中间变量2"."3层下呼分配2",
             下呼分配4 := "中间变量2"."4层下呼分配2",
             下呼分配5 := "中间变量2"."5层下呼分配2",
             下呼分配6 := "中间变量2"."6层下呼分配2",
             下呼分配7 := "中间变量2"."7层下呼分配2",
             下呼分配8 := "中间变量2"."8层下呼分配2",
             下呼分配9 := "中间变量2"."9层下呼分配2",
             下呼分配10 := "中间变量2"."10层下呼分配2",
             内呼1 := "输出"."2号梯1层按钮指示灯",
             内呼2 := "输出"."2号梯2层按钮指示灯",
             内呼3 := "输出"."2号梯3层按钮指示灯",
             内呼4 := "输出"."2号梯4层按钮指示灯",
             内呼5 := "输出"."2号梯5层按钮指示灯",
             内呼6 := "输出"."2号梯6层按钮指示灯",
             内呼7 := "输出"."2号梯7层按钮指示灯",
             内呼8 := "输出"."2号梯8层按钮指示灯",
             内呼9 := "输出"."2号梯9层按钮指示灯",
             内呼10 := "输出"."2号梯10层按钮指示灯",
             当前楼层 := "中间变量2"."2号梯当前楼层数",
             上行停站次数3 => "中间变量2"."2号梯上行停站次数3",
             上行停站次数4 => "中间变量2"."2号梯上行停站次数4",
             上行停站次数5 => "中间变量2"."2号梯上行停站次数5",
             上行停站次数6 => "中间变量2"."2号梯上行停站次数6",
             上行停站次数7 => "中间变量2"."2号梯上行停站次数7",
             上行停站次数8 => "中间变量2"."2号梯上行停站次数8",
             上行停站次数9 => "中间变量2"."2号梯上行停站次数9",
             上行停站次数10 => "中间变量2"."2号梯上行停站次数10",
             上行需折返停站次数10 => "中间变量2"."2号梯上行需折返停站次数10",
             下行停站次数1 => "中间变量2"."2号梯下行停站次数1",
             下行停站次数2 => "中间变量2"."2号梯下行停站次数2",
             下行停站次数3 => "中间变量2"."2号梯下行停站次数3",
             下行停站次数4 => "中间变量2"."2号梯下行停站次数4",
             下行停站次数5 => "中间变量2"."2号梯下行停站次数5",
             下行停站次数6 => "中间变量2"."2号梯下行停站次数6",
             下行停站次数7 => "中间变量2"."2号梯下行停站次数7",
             下行停站次数8 => "中间变量2"."2号梯下行停站次数8",
             下行需折返停站次数1 => "中间变量2"."2号梯下行需折返停站次数1");
END_REGION

REGION Network 4: 3号梯
